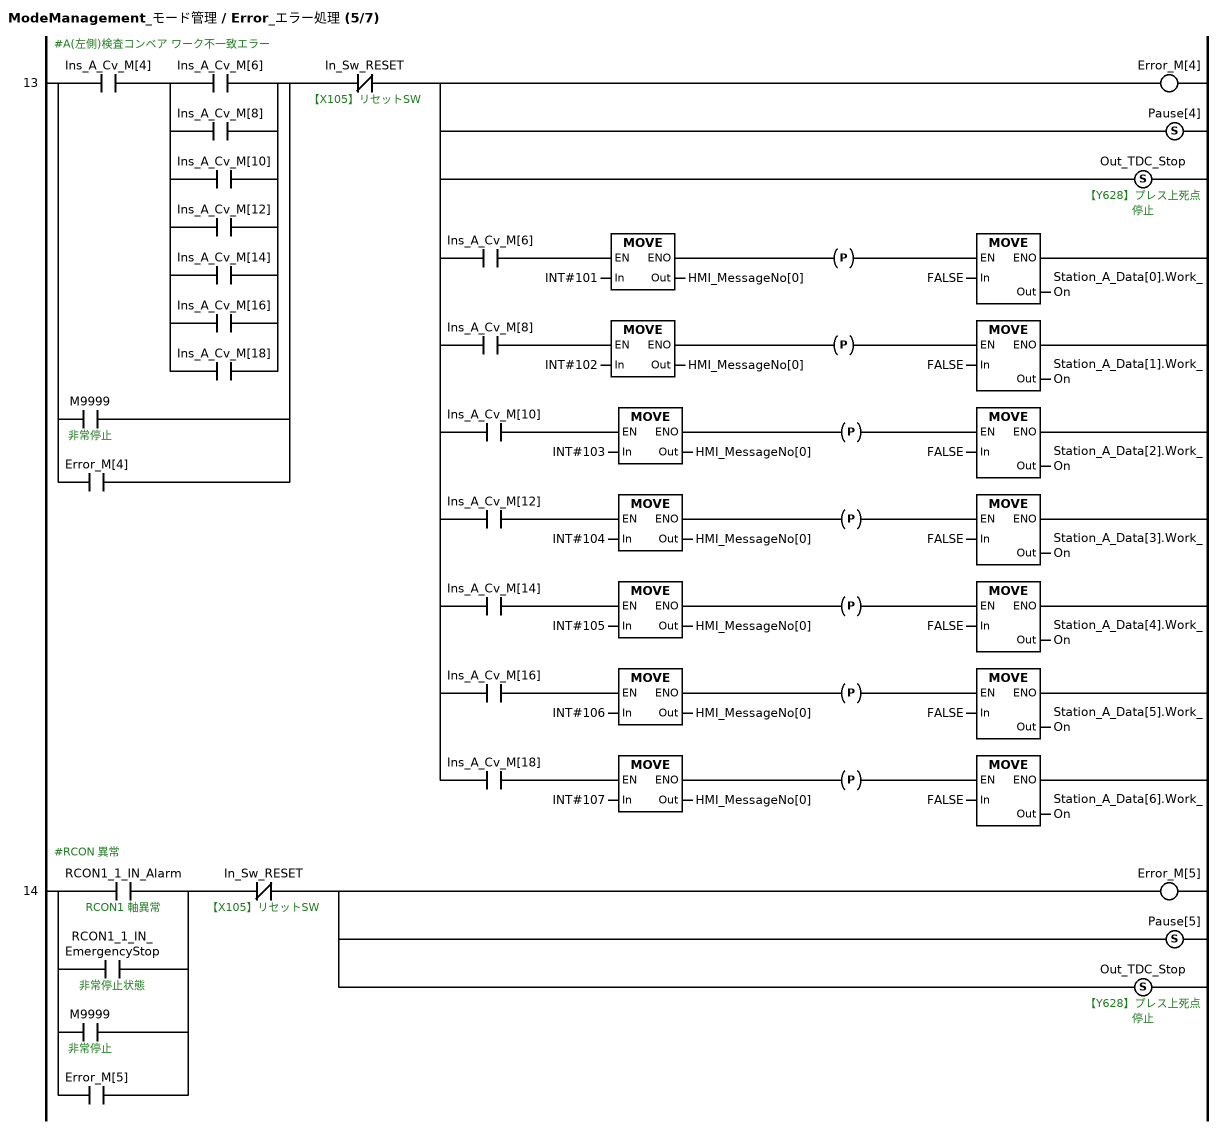
(* [picture p15: ModeManagement_モード管理 / Error_エラー処理, rungs 13-14] *)
(* Rung 13: #A(左側)検査コンベア ワーク不一致エラー *)
_p39 := ((Ins_A_Cv_M[4] AND (Ins_A_Cv_M[6] OR Ins_A_Cv_M[8] OR Ins_A_Cv_M[10] OR Ins_A_Cv_M[12] OR Ins_A_Cv_M[14] OR Ins_A_Cv_M[16] OR Ins_A_Cv_M[18])) OR M9999 OR Error_M[4]) AND NOT In_Sw_RESET;
Error_M[4] := _p39;
IF _p39 THEN
    Pause[4] := TRUE;
    Out_TDC_Stop := TRUE;
END_IF;
IF _p39 AND Ins_A_Cv_M[6] THEN HMI_MessageNo[0] := INT#101; END_IF;
_e40(CLK := _p39 AND Ins_A_Cv_M[6]);
IF _e40.Q THEN Station_A_Data[0].Work_On := FALSE; END_IF;
IF _p39 AND Ins_A_Cv_M[8] THEN HMI_MessageNo[0] := INT#102; END_IF;
_e41(CLK := _p39 AND Ins_A_Cv_M[8]);
IF _e41.Q THEN Station_A_Data[1].Work_On := FALSE; END_IF;
IF _p39 AND Ins_A_Cv_M[10] THEN HMI_MessageNo[0] := INT#103; END_IF;
_e42(CLK := _p39 AND Ins_A_Cv_M[10]);
IF _e42.Q THEN Station_A_Data[2].Work_On := FALSE; END_IF;
IF _p39 AND Ins_A_Cv_M[12] THEN HMI_MessageNo[0] := INT#104; END_IF;
_e43(CLK := _p39 AND Ins_A_Cv_M[12]);
IF _e43.Q THEN Station_A_Data[3].Work_On := FALSE; END_IF;
IF _p39 AND Ins_A_Cv_M[14] THEN HMI_MessageNo[0] := INT#105; END_IF;
_e44(CLK := _p39 AND Ins_A_Cv_M[14]);
IF _e44.Q THEN Station_A_Data[4].Work_On := FALSE; END_IF;
IF _p39 AND Ins_A_Cv_M[16] THEN HMI_MessageNo[0] := INT#106; END_IF;
_e45(CLK := _p39 AND Ins_A_Cv_M[16]);
IF _e45.Q THEN Station_A_Data[5].Work_On := FALSE; END_IF;
IF _p39 AND Ins_A_Cv_M[18] THEN HMI_MessageNo[0] := INT#107; END_IF;
_e46(CLK := _p39 AND Ins_A_Cv_M[18]);
IF _e46.Q THEN Station_A_Data[6].Work_On := FALSE; END_IF;
(* Rung 14: #RCON 異常 *)
_p47 := (RCON1_1_IN_Alarm OR RCON1_1_IN_EmergencyStop OR M9999 OR Error_M[5]) AND NOT In_Sw_RESET;
Error_M[5] := _p47;
IF _p47 THEN
    Pause[5] := TRUE;
    Out_TDC_Stop := TRUE;
END_IF;

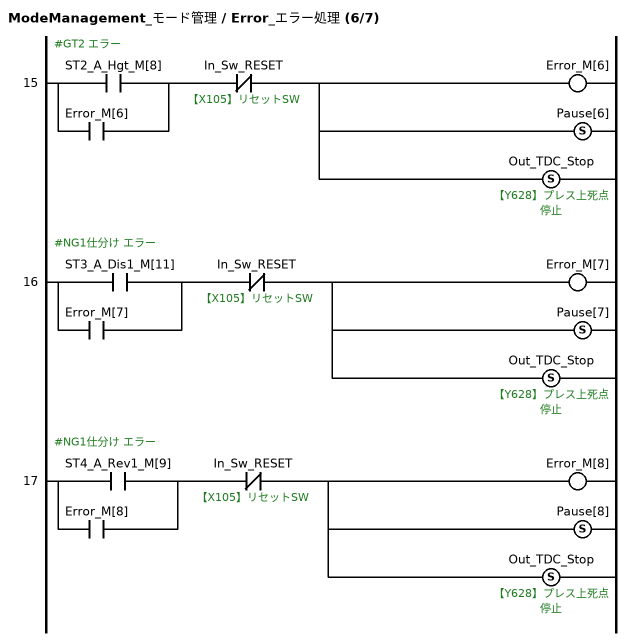
(* Rung 15: #GT2 エラー *)
_p48 := (ST2_A_Hgt_M[8] OR Error_M[6]) AND NOT In_Sw_RESET;
Error_M[6] := _p48;
IF _p48 THEN
    Pause[6] := TRUE;
    Out_TDC_Stop := TRUE;
END_IF;
(* Rung 16: #NG1仕分け エラー *)
_p49 := (ST3_A_Dis1_M[11] OR Error_M[7]) AND NOT In_Sw_RESET;
Error_M[7] := _p49;
IF _p49 THEN
    Pause[7] := TRUE;
    Out_TDC_Stop := TRUE;
END_IF;
(* Rung 17: #NG1仕分け エラー *)
_p50 := (ST4_A_Rev1_M[9] OR Error_M[8]) AND NOT In_Sw_RESET;
Error_M[8] := _p50;
IF _p50 THEN
    Pause[8] := TRUE;
    Out_TDC_Stop := TRUE;
END_IF;

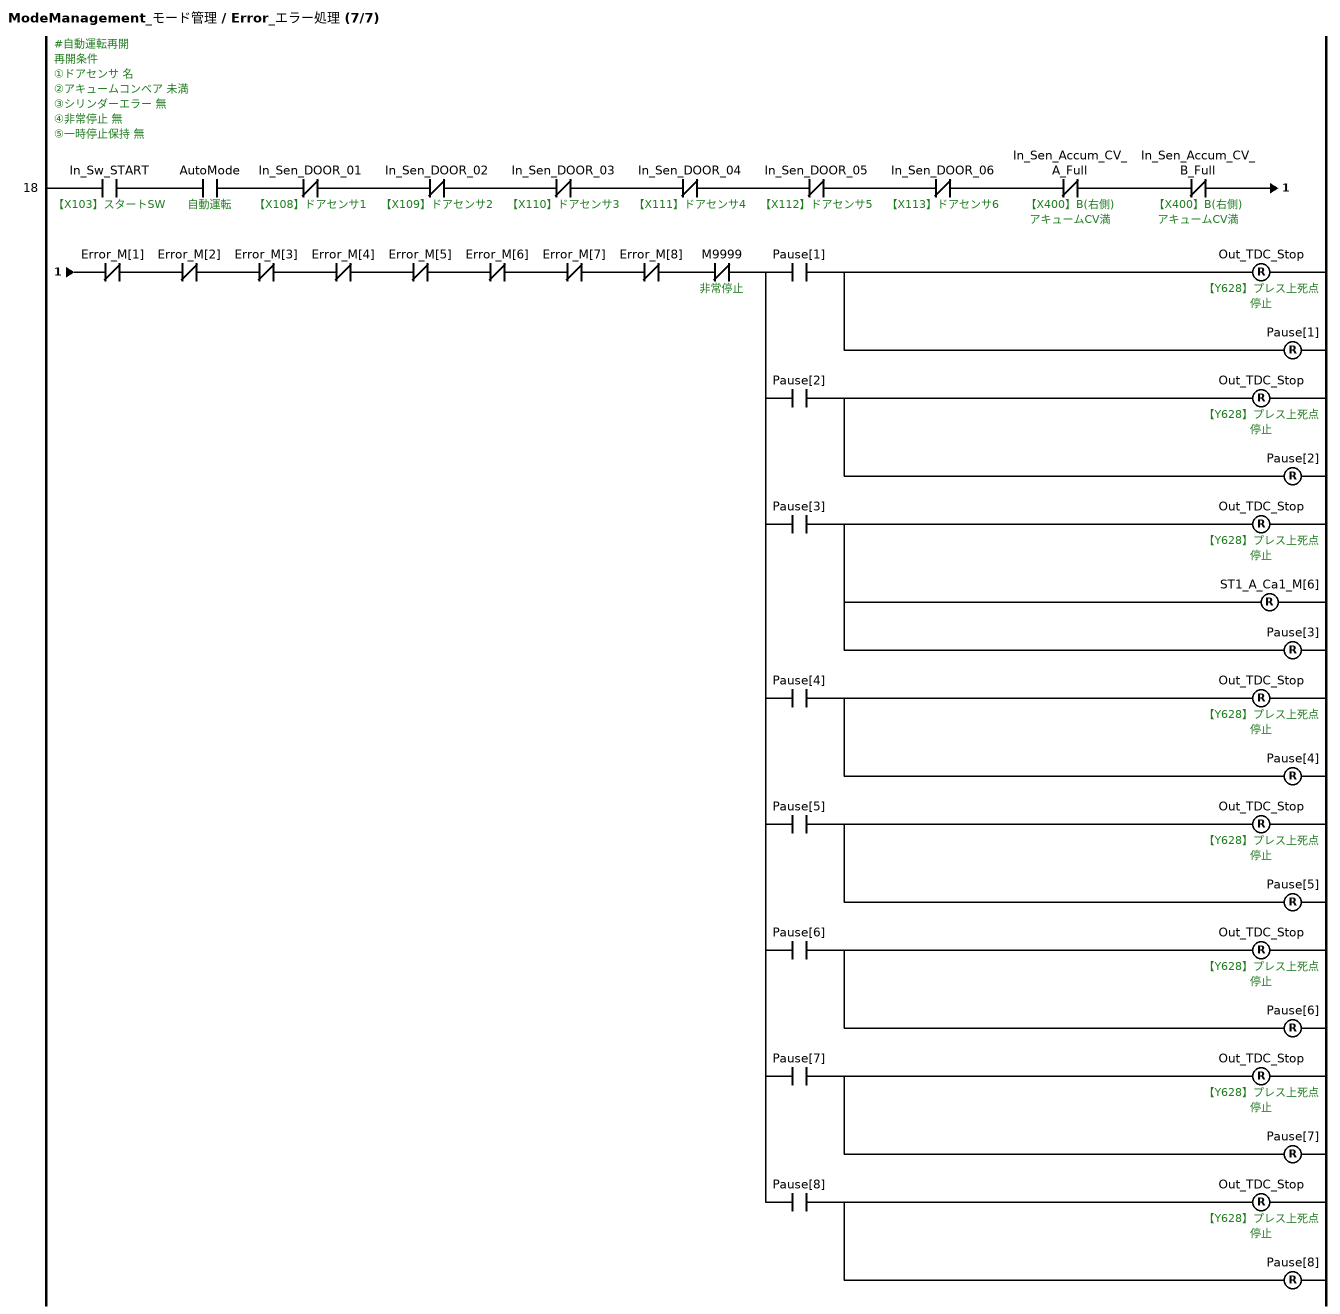
(* Rung 18: #自動運転再開 / 再開条件 / ①ドアセンサ 名 / ②アキュームコンベア 未満 / ③シリンダーエラー 無 / ④非常停止 無 / ⑤一時停止保持 無 *)
_p51 := In_Sw_START AND AutoMode AND NOT In_Sen_DOOR_01 AND NOT In_Sen_DOOR_02 AND NOT In_Sen_DOOR_03 AND NOT In_Sen_DOOR_04 AND NOT In_Sen_DOOR_05 AND NOT In_Sen_DOOR_06 AND NOT In_Sen_Accum_CV_A_Full AND NOT In_Sen_Accum_CV_B_Full AND NOT Error_M[1] AND NOT Error_M[2] AND NOT Error_M[3] AND NOT Error_M[4] AND NOT Error_M[5] AND NOT Error_M[6] AND NOT Error_M[7] AND NOT Error_M[8] AND NOT M9999;
IF _p51 AND Pause[1] THEN
    Out_TDC_Stop := FALSE;
    Pause[1] := FALSE;
END_IF;
IF _p51 AND Pause[2] THEN
    Out_TDC_Stop := FALSE;
    Pause[2] := FALSE;
END_IF;
IF _p51 AND Pause[3] THEN
    Out_TDC_Stop := FALSE;
    ST1_A_Ca1_M[6] := FALSE;
    Pause[3] := FALSE;
END_IF;
IF _p51 AND Pause[4] THEN
    Out_TDC_Stop := FALSE;
    Pause[4] := FALSE;
END_IF;
IF _p51 AND Pause[5] THEN
    Out_TDC_Stop := FALSE;
    Pause[5] := FALSE;
END_IF;
IF _p51 AND Pause[6] THEN
    Out_TDC_Stop := FALSE;
    Pause[6] := FALSE;
END_IF;
IF _p51 AND Pause[7] THEN
    Out_TDC_Stop := FALSE;
    Pause[7] := FALSE;
END_IF;
IF _p51 AND Pause[8] THEN
    Out_TDC_Stop := FALSE;
    Pause[8] := FALSE;
END_IF;
END_PROGRAM

PROGRAM Movements_動作
VAR
    Mo_M : BOOL;
    ST0_A_Sup_M : ARRAY[0..99] OF Bool;  (* [4] 原点位置移動完了 *)
    ST1_Ins_Cv_Rdy : BOOL;
    ST2_Ins_Cv_Rdy : BOOL;
    ST3_Ins_Cv_Rdy : BOOL;
    ST4_Ins_Cv_Rdy : BOOL;
    ST5_Ins_Cv_Rdy : BOOL;
    ST6_Ins_Cv_Rdy : BOOL;
    ST7_Ins_Cv_Rdy : BOOL;
    Ins_A_Cv_T : ARRAY[0..99] OF TON;
    ST1_A_Ca1_Rdy : BOOL;
    GT2_A_Inspection_GetTime : DATE_AND_TIME;
    GT2_A_Inspection_GetTime_ST : STRING[256];
    GT2_A_Inspection_GetTime_ST_Del : STRING[20];
    ST4_A_Rev1_Busy : BOOL;  (* ST4 A 動作中 *)
END_VAR
VAR_EXTERNAL
    ST0_Sup_Start : BOOL;  (* ST0_動作開始 *)
    M9999 : BOOL;
    Out_CYw_Sply_Pick_A_H_Auto : ARRAY[0..10] OF Bool;
    Out_CYw_Sply_Pick_A_H_Done : BOOL;
    Out_CYw_Sply_Slide_A_H_Auto : ARRAY[0..10] OF Bool;
    Out_CYw_Sply_Slide_A_H_Done : BOOL;
    Out_CYw_Sup_Chuck_A_Cl_H_Auto : ARRAY[0..10] OF Bool;
    Out_CYw_Sup_Chuck_A_Cl_H_Done : BOOL;
    In_Sen_Accum_CV_A_Arrival : BOOL;
    In_Sen_Work_A_Pos_00 : BOOL;
    Out_CYw_Sply_Pick_A_F_Auto : ARRAY[0..10] OF Bool;
    Out_CYw_Sply_Pick_A_F_Done : BOOL;
    Out_CYw_Sup_Chuck_A_Cl_F_Auto : ARRAY[0..10] OF Bool;
    Out_CYw_Sup_Chuck_A_Cl_F_Done : BOOL;
    Out_CYw_Sply_Slide_A_F_Auto : ARRAY[0..10] OF Bool;
    Out_CYw_Sply_Slide_A_F_Done : BOOL;
    Station_A_Data : ARRAY[0..8] OF sData;
    Cv_A_Data : ARRAY[0..8] OF sData;
    ST0_A_Sup_End : BOOL;  (* ST0 検査コンベア運転可 *)
    Out_CYS_Pos_01_Stopper_B_H_Auto : ARRAY[0..10] OF Bool;
    Out_CYS_Pos_02_Stopper_B_H_Auto : ARRAY[0..10] OF Bool;
    Out_CYS_Pos_03_Stopper_B_H_Auto : ARRAY[0..10] OF Bool;
    Out_CYS_Pos_04_Stopper_B_H_Auto : ARRAY[0..10] OF Bool;
    Out_CYS_Pos_05_Stopper_B_H_Auto : ARRAY[0..10] OF Bool;
    Out_CYS_Pos_06_Stopper_B_H_Auto : ARRAY[0..10] OF Bool;
    TimerQ_In_SenCY_Pos_01_Stopper_A_H : BOOL;
    TimerQ_In_SenCY_Pos_02_Stopper_A_H : BOOL;
    TimerQ_In_SenCY_Pos_03_Stopper_A_H : BOOL;
    TimerQ_In_SenCY_Pos_04_Stopper_A_H : BOOL;
    TimerQ_In_SenCY_Pos_05_Stopper_A_H : BOOL;
    TimerQ_In_SenCY_Pos_06_Stopper_A_H : BOOL;
    Out_Insp_Cv_A_Run_Auto : ARRAY[0..10] OF Bool;
    TimerQ_In_Sen_Work_A_Pos_01 : BOOL;
    TimerQ_In_Sen_Work_A_Pos_02 : BOOL;
    Pause : ARRAY[0..99] OF Bool;
    TimerQ_In_Sen_Work_A_Pos_03 : BOOL;
    TimerQ_In_Sen_Work_A_Pos_04 : BOOL;
    TimerQ_In_Sen_Work_A_Pos_05 : BOOL;
    TimerQ_In_Sen_Work_A_Pos_06 : BOOL;
    TimerQ_In_Sen_Work_A_Pos_07 : BOOL;
    Out_CYS_Pos_01_Stopper_A_H_Auto : ARRAY[0..10] OF Bool;
    Out_CYS_Pos_02_Stopper_A_H_Auto : ARRAY[0..10] OF Bool;
    Out_CYS_Pos_03_Stopper_A_H_Auto : ARRAY[0..10] OF Bool;
    Out_CYS_Pos_04_Stopper_A_H_Auto : ARRAY[0..10] OF Bool;
    Out_CYS_Pos_05_Stopper_A_H_Auto : ARRAY[0..10] OF Bool;
    Out_CYS_Pos_06_Stopper_A_H_Auto : ARRAY[0..10] OF Bool;
    Ins_A_Cv_M : ARRAY[0..99] OF Bool;
    Ins_A_Cv_Error : BOOL;  (* 検査コンベア ワーク不一致エラー *)
    TimerQ_In_Sen_Work_A_Pos_00 : BOOL;
    Out_CYS_Pos_01_Stopper_A_F_Auto : ARRAY[0..10] OF Bool;
    Out_CYS_Pos_02_Stopper_A_F_Auto : ARRAY[0..10] OF Bool;
    Out_CYS_Pos_03_Stopper_A_F_Auto : ARRAY[0..10] OF Bool;
    Out_CYS_Pos_04_Stopper_A_F_Auto : ARRAY[0..10] OF Bool;
    Out_CYS_Pos_05_Stopper_A_F_Auto : ARRAY[0..10] OF Bool;
    Out_CYS_Pos_06_Stopper_A_F_Auto : ARRAY[0..10] OF Bool;
    Ins_A_Next_Cycle : BOOL;  (* A(左側)検査コンベア 動作完了 *)
    ST0_A_Sup_Busy : BOOL;  (* ST0 稼働中 *)
    Ins_A_End : BOOL;  (* 検査完了 コンベア運転可能 *)
    Auto_A_Start : BOOL;
    Out_CYS_Pos_01_Stopper_A_H_Done : BOOL;
    FH_5552_10_A_Auto : BOOL;
    FH_A_ST1_Done : BOOL;
    ST1_A_Ca1_Busy : BOOL;  (* ST1 A検査中 *)
    ST1_A_Ca1_End : BOOL;  (* ST1 A 動作完了 *)
    ST2_A_Hgt_Busy : BOOL;  (* ST2 A 動作中 *)
    Out_CYw_HgtInsp_Clp_A_H_Auto : ARRAY[0..10] OF Bool;
    Out_CYw_HgtInsp_Clp_A_H_Done : BOOL;
    Out_CYw_HgtInsp_Lf_A_H_Auto : ARRAY[0..10] OF Bool;
    Out_CYw_HgtInsp_Lf_A_H_Done : BOOL;
    Out_CYS_Pos_02_Stopper_A_H_Done : BOOL;
    Out_CYw_HgtInsp_Clp_A_F_Auto : ARRAY[0..10] OF Bool;
    Out_CYw_HgtInsp_Clp_A_F_Done : BOOL;
    Out_CYw_HgtInsp_Lf_A_F_Auto : ARRAY[0..10] OF Bool;
    Out_CYw_HgtInsp_Lf_A_F_Done : BOOL;
    DLEP1_GT2_A_Auto : BOOL;
    Hgt_A_ComputedValueData : LREAL;
    Hight_LowerLimit : LREAL;  (* 高さ検査 下限値 *)
    Hight_UpperLimit : LREAL;  (* 高さ検査 上限値 *)
    ST2_A_Hgt_End : BOOL;  (* 高さ検査完了 *)
    ST3_A_Dis1_Busy : BOOL;  (* ST3 A 動作中 *)
    Out_CYw_NG1_Srt_A_H_Auto : ARRAY[0..10] OF Bool;
    Out_CYw_NG1_Srt_A_H_Done : BOOL;
    Out_CYw_Rev_01_Pick_A_H_Auto : ARRAY[0..10] OF Bool;  (* 自動【Y710】A(左側)ST4 反転1ピックアップ戻： *)
    Out_CYw_Rev_01_Pick_A_H_Done : BOOL;  (* 【Y710】A(左側)ST4 反転1ピックアップ戻 動作完了 *)
    Out_CYw_NG1_Pick_A_H_Auto : ARRAY[0..10] OF Bool;
    Out_CYw_NG1_Pick_A_H_Done : BOOL;
    Out_CYw_NG1_Chk_A_H_Auto : ARRAY[0..10] OF Bool;
    Out_CYw_NG1_Chk_A_H_Done : BOOL;
    RCON1_IAI_Auto : ARRAY[0..99] OF Bool;  (* A(左側) RCON1/Node1/ NG排出： *)
    RCON1_OUT_TargetPos_mm : LREAL;
    HMI_RCON1_OUT_TargetPos : ARRAY[0..99] OF LREAL;  (* HMI RC01 NG仕分け位置： *)
    RCON1_1_M : ARRAY[0..99] OF BOOL;
    Error_M : ARRAY[0..99] OF Bool;
    ST1_A_Ca1_M : ARRAY[0..99] OF Bool;  (* [6] ST2 検査前ワーク不一致エラー; [3] ワーク有無 判定; [1] ST1 A カメラ1 検査開始; [4] ST1 A ワーク有; [5] ST1 A ワーク無; [2] 【Y720】A(左側) 位置1ストッパー 戻; [7] ST1 FH測定開始 *)
    ST2_A_Hgt_M : ARRAY[0..99] OF Bool;  (* [4] 【Y721】A(左側) 位置2ストッパー戻; [6] ST1 A ワーク有; [7] ST1 A ワーク無; [5] ワーク有無 判定; [9] 【Y703】A(左側) 高さ検査持上行; [10] 【Y701】A(左側) 高さ検査押え行; [11] A(左側) 高さ検査OK判定; [12] A(左側) 高さ検査NG判定; [2] 【Y701】A(左側) 高さ検査押え行; [8] ST3 検査前ワーク不一致エラー *)
    Out_CYS_Pos_03_Stopper_A_H_Done : BOOL;
    Out_CYw_NG1_Pick_A_F_Auto : ARRAY[0..10] OF Bool;
    Out_CYw_NG1_Pick_A_F_Done : BOOL;
    Out_CYw_NG1_Chk_A_F_Auto : ARRAY[0..10] OF Bool;
    Out_CYw_NG1_Chk_A_F_Done : BOOL;
    Out_CYw_NG1_Srt_A_F_Auto : ARRAY[0..10] OF Bool;
    Out_CYw_NG1_Srt_A_F_Done : BOOL;
    ST3_A_Dis1_End : BOOL;  (* 左NG1排出 完了 *)
    ST3_A_Dis1_M : ARRAY[0..99] OF Bool;  (* [7] 原点位置 移動開始; [6] 原点位置移動 データ転送; [5] 【Y722】A(左側) 位置3ストッパー戻; [4] 【Y706】A(左側) NG1チャック戻; [8] ワーク有無 / 検査前ワーク不一致 判定; [9] S3 A ワーク有 工程NG; [10] S3 A ワーク無  前工程OK; [14] 【Y704】A(左側) NG1ピックアップ戻 ; [24] 仕分け完了 *)
    ST4_A_Rev1_M : ARRAY[0..99] OF Bool;  (* [2] ワーク有無 / 検査前ワーク不一致 判定; [3] 【Y723】A(左側) 位置4ストッパー戻; [4] ST4 A ワーク有; [5] ST4 A ワーク無 / 前工程NG; [6] ST4 検査前ワーク不一致エラー *)
    Stm_A_Rev_Axis000_MovePos_Degree : LREAL;
    HMI_Stm_A_Rev_Axis000_MovePos_Degree : LREAL;  (* A(左側)ステッピングモータ000 回転角度 *)
    Stm_A_Rev_Axis000_Auto : ARRAY[0..99] OF Bool;  (* [1] 原点位置移動 開始 *)
    Stm_A_Rev_Axis000_MoveAbsoluteDone : BOOL;
END_VAR
VAR
    _e1 : R_TRIG;
    _p2 : BOOL;
    _e3 : R_TRIG;
    _e4 : R_TRIG;
    _p5 : BOOL;
    _e6 : R_TRIG;
    _e7 : R_TRIG;
    _p8 : BOOL;
    _p9 : BOOL;
    _p10 : BOOL;
    _p11 : BOOL;
    _p12 : BOOL;
    _p13 : BOOL;
    _p14 : BOOL;
    _p15 : BOOL;
    _e16 : R_TRIG;
    _p17 : BOOL;
    _p18 : BOOL;
    _p19 : BOOL;
    _p20 : BOOL;
    _p21 : BOOL;
    _p22 : BOOL;
    _p23 : BOOL;
    _p24 : BOOL;
    _p25 : BOOL;
    _p26 : BOOL;
    _p27 : BOOL;
    _p28 : BOOL;
    _e29 : R_TRIG;
    _p30 : BOOL;
    _p31 : BOOL;
    _p32 : BOOL;
    _p33 : BOOL;
    _p34 : BOOL;
    _p35 : BOOL;
    _p36 : BOOL;
    _p37 : BOOL;
    _p38 : BOOL;
    _p39 : BOOL;
    _p40 : BOOL;
    _p41 : BOOL;
    _p42 : BOOL;
    _p43 : BOOL;
    _p44 : BOOL;
    _p45 : BOOL;
    _p46 : BOOL;
    _p47 : BOOL;
    _p48 : BOOL;
    _p49 : BOOL;
    _p50 : BOOL;
    _p51 : BOOL;
    _p52 : BOOL;
    _p53 : BOOL;
    _p54 : BOOL;
    _p55 : BOOL;
    _p56 : BOOL;
    _p57 : BOOL;
    _p58 : BOOL;
    _p59 : BOOL;
    _p60 : BOOL;
    _p61 : BOOL;
END_VAR

(* Section Ins_A_Cv_左検査Cv: ladder, written here as Structured Text *)

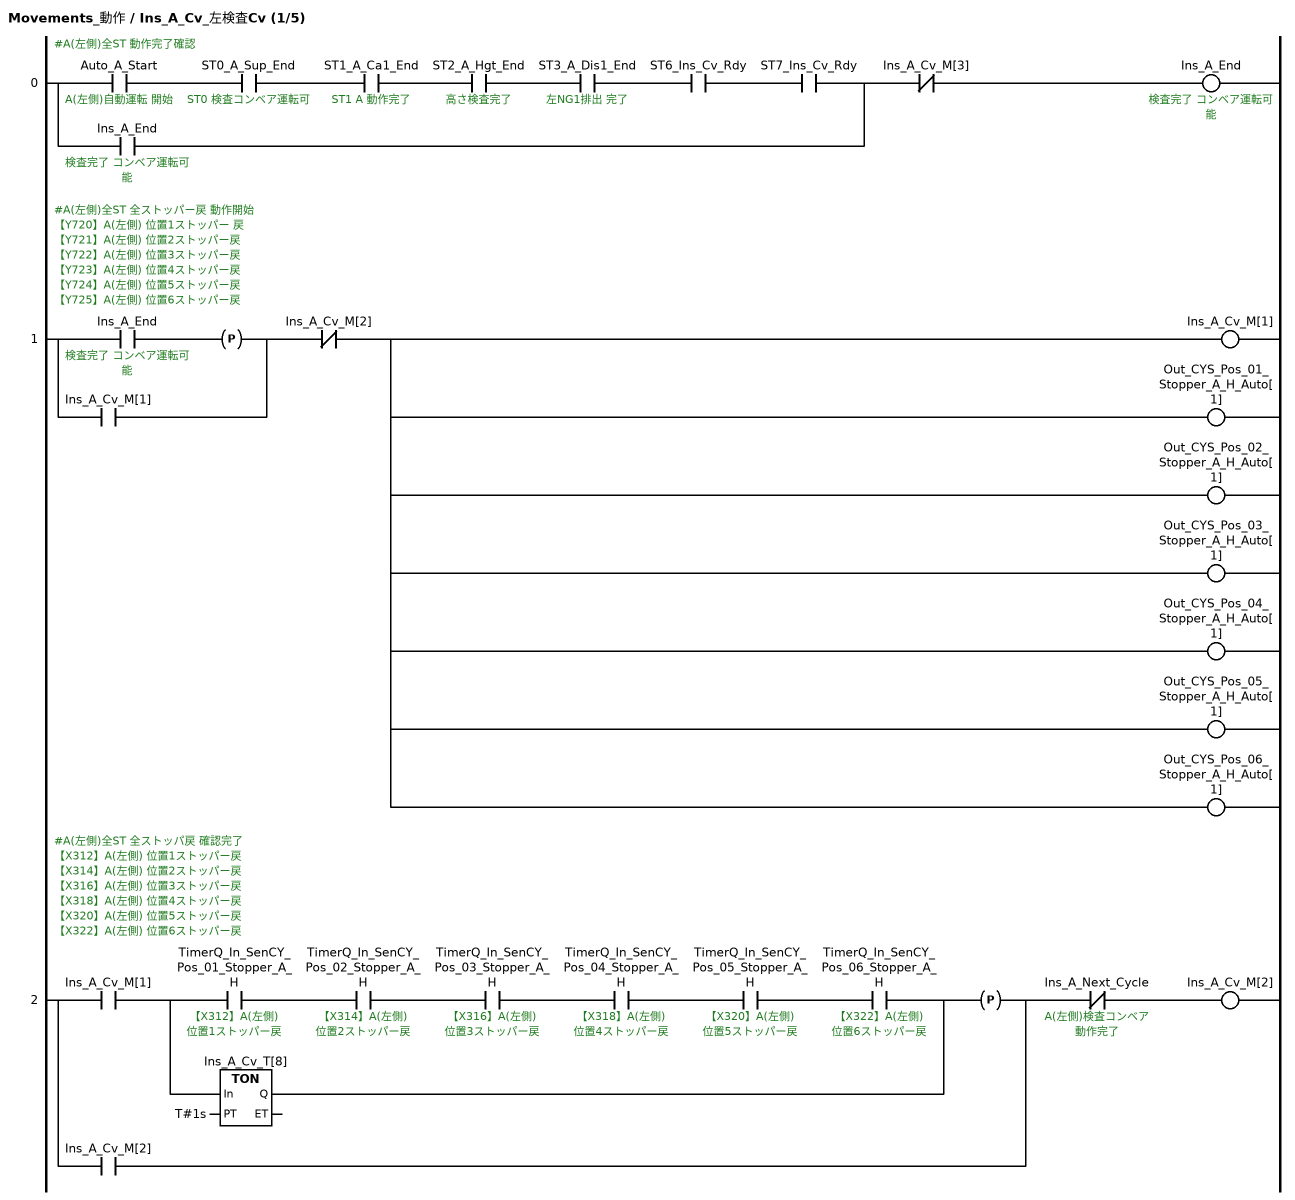
(* Rung 0: #A(左側)全ST 動作完了確認 *)
Ins_A_End := ((Auto_A_Start AND ST0_A_Sup_End AND ST1_A_Ca1_End AND ST2_A_Hgt_End AND ST3_A_Dis1_End AND ST6_Ins_Cv_Rdy AND ST7_Ins_Cv_Rdy) OR Ins_A_End) AND NOT Ins_A_Cv_M[3];
(* Rung 1: #A(左側)全ST 全ストッパー戻 動作開始 / 【Y720】A(左側) 位置1ストッパー 戻 / 【Y721】A(左側) 位置2ストッパー戻 / 【Y722】A(左側) 位置3ストッパー戻 / 【Y723】A(左側) 位置4ストッパー戻 / 【Y724】A(左側) 位置5ストッパー戻 / 【Y725】A(左側) 位置6ストッパー戻 *)
_e1(CLK := Ins_A_End);
_p2 := (_e1.Q OR Ins_A_Cv_M[1]) AND NOT Ins_A_Cv_M[2];
Ins_A_Cv_M[1] := _p2;
Out_CYS_Pos_01_Stopper_A_H_Auto[1] := _p2;
Out_CYS_Pos_02_Stopper_A_H_Auto[1] := _p2;
Out_CYS_Pos_03_Stopper_A_H_Auto[1] := _p2;
Out_CYS_Pos_04_Stopper_A_H_Auto[1] := _p2;
Out_CYS_Pos_05_Stopper_A_H_Auto[1] := _p2;
Out_CYS_Pos_06_Stopper_A_H_Auto[1] := _p2;
(* Rung 2: #A(左側)全ST 全ストッパ戻 確認完了 / 【X312】A(左側) 位置1ストッパー戻 / 【X314】A(左側) 位置2ストッパー戻 / 【X316】A(左側) 位置3ストッパー戻 / 【X318】A(左側) 位置4ストッパー戻 / 【X320】A(左側) 位置5ストッパー戻 / 【X322】A(左側) 位置6ストッパー戻 *)
Ins_A_Cv_T[8](In := Ins_A_Cv_M[1], PT := T#1s);
_e3(CLK := (Ins_A_Cv_M[1] AND TimerQ_In_SenCY_Pos_01_Stopper_A_H AND TimerQ_In_SenCY_Pos_02_Stopper_A_H AND TimerQ_In_SenCY_Pos_03_Stopper_A_H AND TimerQ_In_SenCY_Pos_04_Stopper_A_H AND TimerQ_In_SenCY_Pos_05_Stopper_A_H AND TimerQ_In_SenCY_Pos_06_Stopper_A_H) OR Ins_A_Cv_T[8].Q);
Ins_A_Cv_M[2] := (_e3.Q OR Ins_A_Cv_M[2]) AND NOT Ins_A_Next_Cycle;

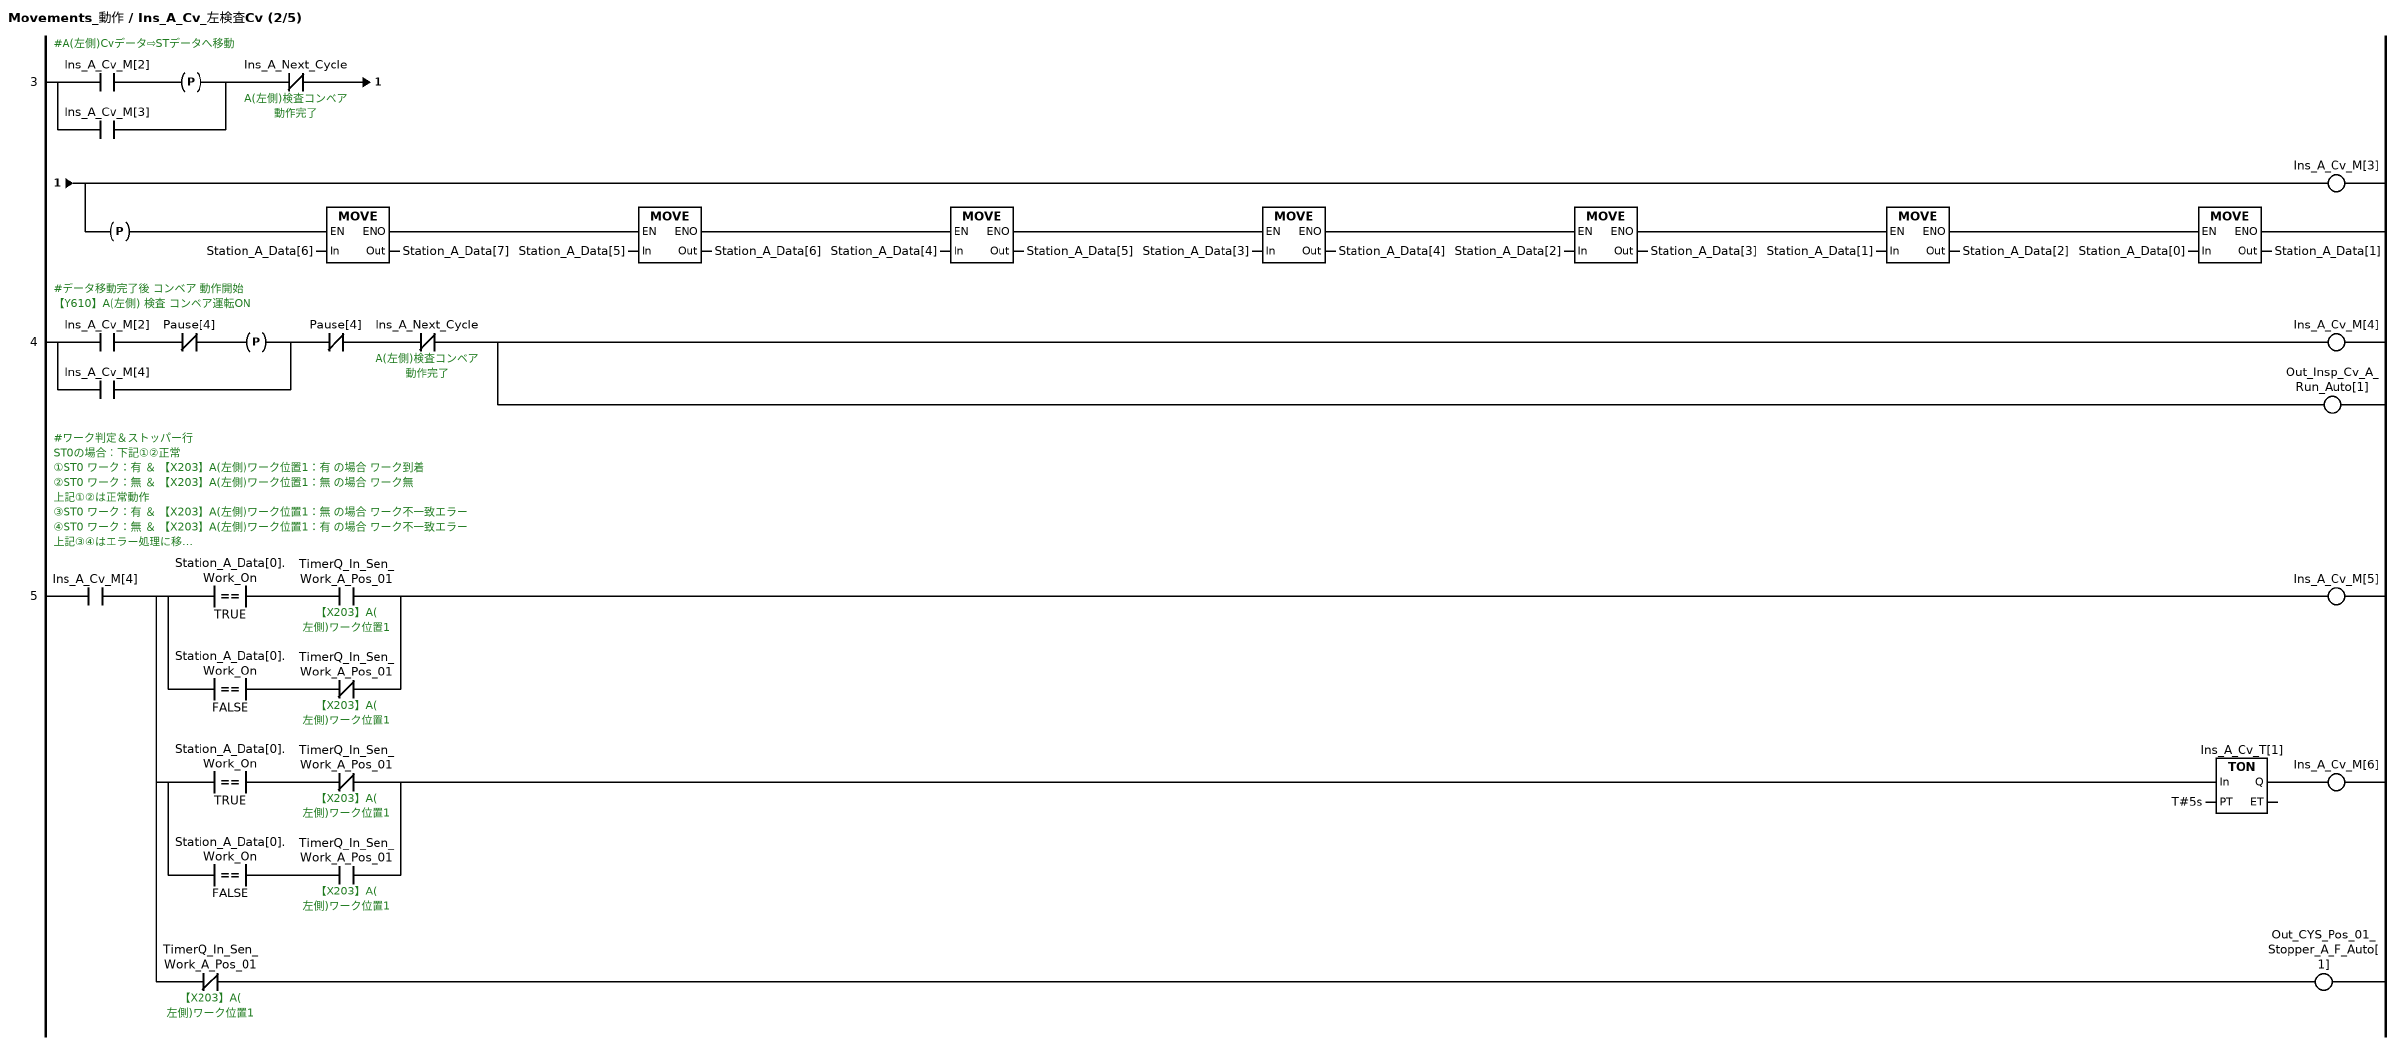
(* Rung 3: #A(左側)Cvデータ⇨STデータへ移動 *)
_e4(CLK := Ins_A_Cv_M[2]);
_p5 := (_e4.Q OR Ins_A_Cv_M[3]) AND NOT Ins_A_Next_Cycle;
Ins_A_Cv_M[3] := _p5;
_e6(CLK := _p5);
IF _e6.Q THEN
    Station_A_Data[7] := Station_A_Data[6];
    Station_A_Data[6] := Station_A_Data[5];
    Station_A_Data[5] := Station_A_Data[4];
    Station_A_Data[4] := Station_A_Data[3];
    Station_A_Data[3] := Station_A_Data[2];
    Station_A_Data[2] := Station_A_Data[1];
    Station_A_Data[1] := Station_A_Data[0];
END_IF;
(* Rung 4: #データ移動完了後 コンベア 動作開始 / 【Y610】A(左側) 検査 コンベア運転ON *)
_e7(CLK := Ins_A_Cv_M[2] AND NOT Pause[4]);
_p8 := (_e7.Q OR Ins_A_Cv_M[4]) AND NOT Pause[4] AND NOT Ins_A_Next_Cycle;
Ins_A_Cv_M[4] := _p8;
Out_Insp_Cv_A_Run_Auto[1] := _p8;
(* Rung 5: #ワーク判定＆ストッパー行 / ST0の場合：下記①②正常 / ①ST0 ワーク：有 ＆ 【X203】A(左側)ワーク位置1：有 の場合 ワーク到着 / ②ST0 ワーク：無 ＆ 【X203】A(左側)ワーク位置1：無 の場合 ワーク無 / 上記①②は正常動作 / ③ST0 ワーク：有 ＆ 【X203】A(左側)ワーク位置1：無 の場合 ワーク不一致エラー / ④ST0 ワーク：無 ＆ 【X203】A(左側)ワーク位置1：有 の場合 ワーク不一致エラー / 上記③④はエラー処理に移動 / ⑤【X203】A(左側)ワーク位置1：無 の場合 / 【Y720】A(左側) 位置1ストッパー 行 *)
_p9 := Ins_A_Cv_M[4];
Ins_A_Cv_M[5] := Ins_A_Cv_M[4] AND (((Station_A_Data[0].Work_On = TRUE) AND TimerQ_In_Sen_Work_A_Pos_01) OR ((Station_A_Data[0].Work_On = FALSE) AND NOT TimerQ_In_Sen_Work_A_Pos_01));
Ins_A_Cv_T[1](In := _p9 AND (((Station_A_Data[0].Work_On = TRUE) AND NOT TimerQ_In_Sen_Work_A_Pos_01) OR ((Station_A_Data[0].Work_On = FALSE) AND TimerQ_In_Sen_Work_A_Pos_01)), PT := T#5s);
Ins_A_Cv_M[6] := Ins_A_Cv_T[1].Q;
Out_CYS_Pos_01_Stopper_A_F_Auto[1] := _p9 AND NOT TimerQ_In_Sen_Work_A_Pos_01;

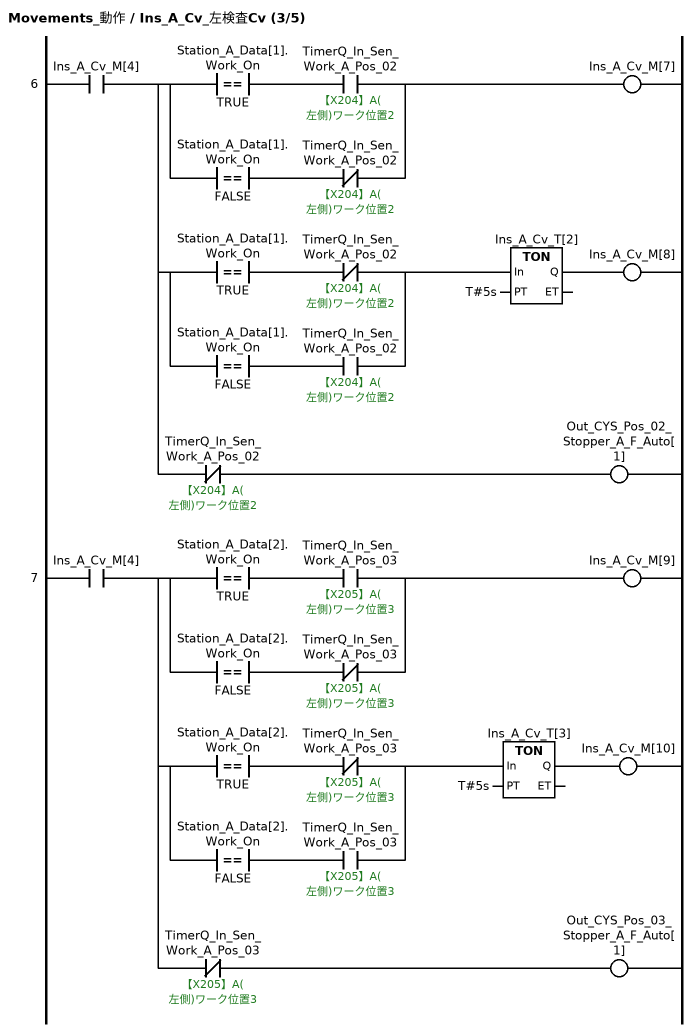
(* Rung 6 *)
_p10 := Ins_A_Cv_M[4];
Ins_A_Cv_M[7] := Ins_A_Cv_M[4] AND (((Station_A_Data[1].Work_On = TRUE) AND TimerQ_In_Sen_Work_A_Pos_02) OR ((Station_A_Data[1].Work_On = FALSE) AND NOT TimerQ_In_Sen_Work_A_Pos_02));
Ins_A_Cv_T[2](In := _p10 AND (((Station_A_Data[1].Work_On = TRUE) AND NOT TimerQ_In_Sen_Work_A_Pos_02) OR ((Station_A_Data[1].Work_On = FALSE) AND TimerQ_In_Sen_Work_A_Pos_02)), PT := T#5s);
Ins_A_Cv_M[8] := Ins_A_Cv_T[2].Q;
Out_CYS_Pos_02_Stopper_A_F_Auto[1] := _p10 AND NOT TimerQ_In_Sen_Work_A_Pos_02;
(* Rung 7 *)
_p11 := Ins_A_Cv_M[4];
Ins_A_Cv_M[9] := Ins_A_Cv_M[4] AND (((Station_A_Data[2].Work_On = TRUE) AND TimerQ_In_Sen_Work_A_Pos_03) OR ((Station_A_Data[2].Work_On = FALSE) AND NOT TimerQ_In_Sen_Work_A_Pos_03));
Ins_A_Cv_T[3](In := _p11 AND (((Station_A_Data[2].Work_On = TRUE) AND NOT TimerQ_In_Sen_Work_A_Pos_03) OR ((Station_A_Data[2].Work_On = FALSE) AND TimerQ_In_Sen_Work_A_Pos_03)), PT := T#5s);
Ins_A_Cv_M[10] := Ins_A_Cv_T[3].Q;
Out_CYS_Pos_03_Stopper_A_F_Auto[1] := _p11 AND NOT TimerQ_In_Sen_Work_A_Pos_03;

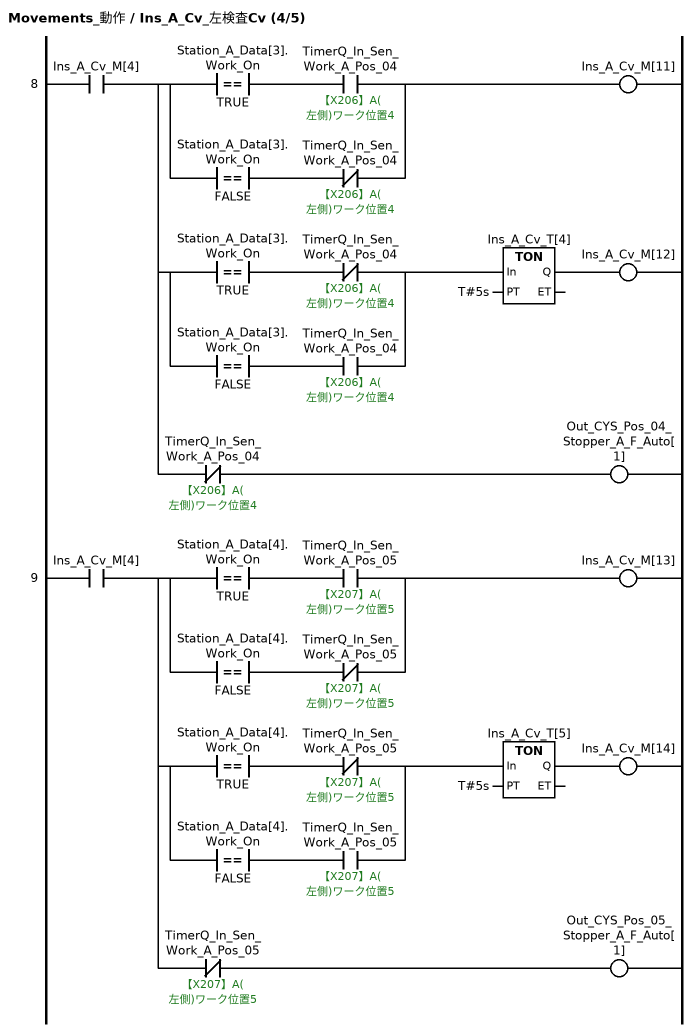
(* Rung 8 *)
_p12 := Ins_A_Cv_M[4];
Ins_A_Cv_M[11] := Ins_A_Cv_M[4] AND (((Station_A_Data[3].Work_On = TRUE) AND TimerQ_In_Sen_Work_A_Pos_04) OR ((Station_A_Data[3].Work_On = FALSE) AND NOT TimerQ_In_Sen_Work_A_Pos_04));
Ins_A_Cv_T[4](In := _p12 AND (((Station_A_Data[3].Work_On = TRUE) AND NOT TimerQ_In_Sen_Work_A_Pos_04) OR ((Station_A_Data[3].Work_On = FALSE) AND TimerQ_In_Sen_Work_A_Pos_04)), PT := T#5s);
Ins_A_Cv_M[12] := Ins_A_Cv_T[4].Q;
Out_CYS_Pos_04_Stopper_A_F_Auto[1] := _p12 AND NOT TimerQ_In_Sen_Work_A_Pos_04;
(* Rung 9 *)
_p13 := Ins_A_Cv_M[4];
Ins_A_Cv_M[13] := Ins_A_Cv_M[4] AND (((Station_A_Data[4].Work_On = TRUE) AND TimerQ_In_Sen_Work_A_Pos_05) OR ((Station_A_Data[4].Work_On = FALSE) AND NOT TimerQ_In_Sen_Work_A_Pos_05));
Ins_A_Cv_T[5](In := _p13 AND (((Station_A_Data[4].Work_On = TRUE) AND NOT TimerQ_In_Sen_Work_A_Pos_05) OR ((Station_A_Data[4].Work_On = FALSE) AND TimerQ_In_Sen_Work_A_Pos_05)), PT := T#5s);
Ins_A_Cv_M[14] := Ins_A_Cv_T[5].Q;
Out_CYS_Pos_05_Stopper_A_F_Auto[1] := _p13 AND NOT TimerQ_In_Sen_Work_A_Pos_05;

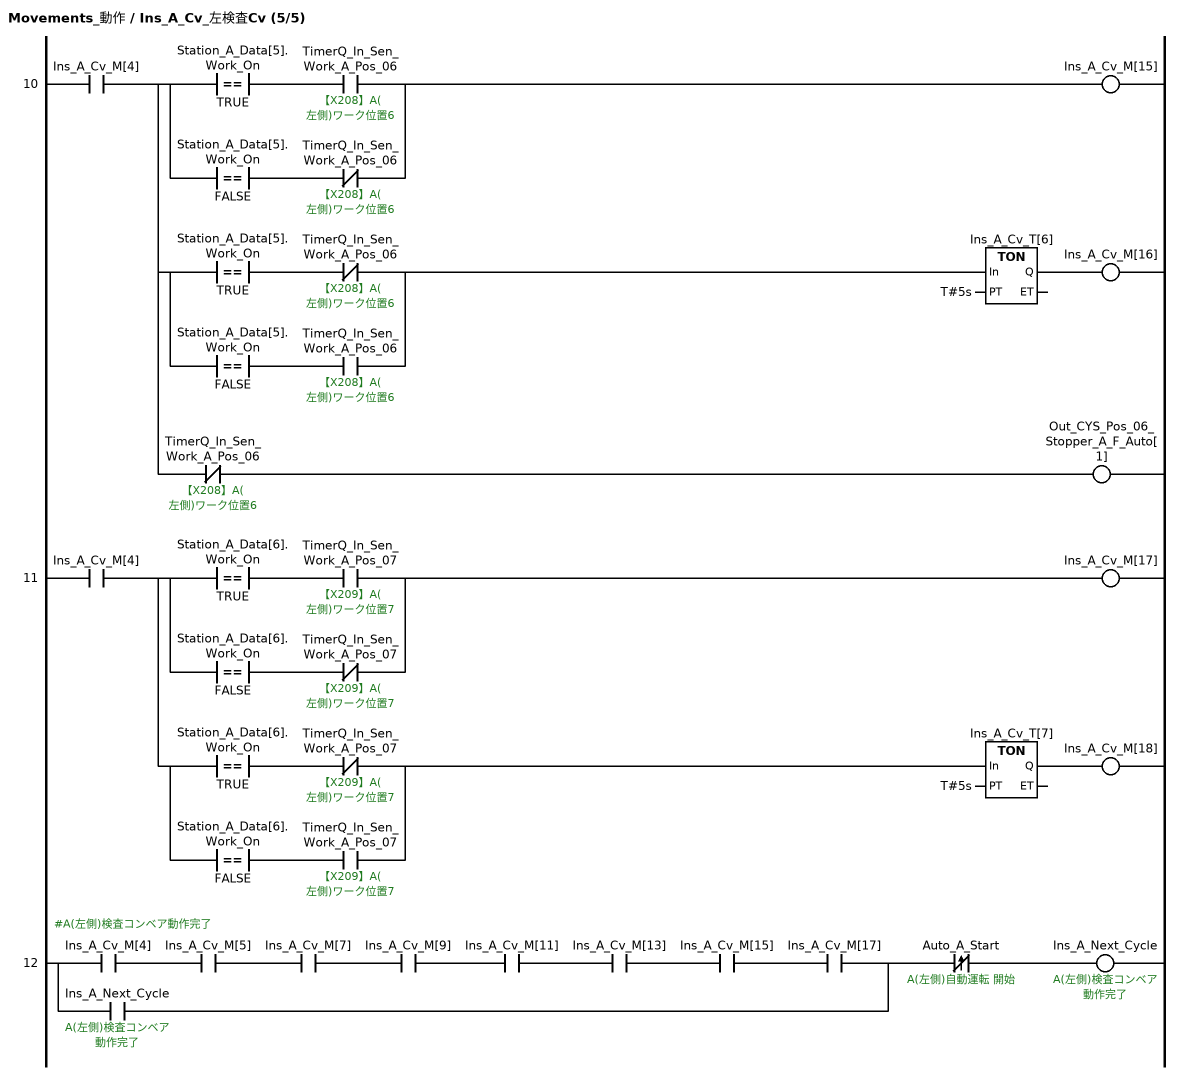
(* Rung 10 *)
_p14 := Ins_A_Cv_M[4];
Ins_A_Cv_M[15] := Ins_A_Cv_M[4] AND (((Station_A_Data[5].Work_On = TRUE) AND TimerQ_In_Sen_Work_A_Pos_06) OR ((Station_A_Data[5].Work_On = FALSE) AND NOT TimerQ_In_Sen_Work_A_Pos_06));
Ins_A_Cv_T[6](In := _p14 AND (((Station_A_Data[5].Work_On = TRUE) AND NOT TimerQ_In_Sen_Work_A_Pos_06) OR ((Station_A_Data[5].Work_On = FALSE) AND TimerQ_In_Sen_Work_A_Pos_06)), PT := T#5s);
Ins_A_Cv_M[16] := Ins_A_Cv_T[6].Q;
Out_CYS_Pos_06_Stopper_A_F_Auto[1] := _p14 AND NOT TimerQ_In_Sen_Work_A_Pos_06;
(* Rung 11 *)
_p15 := Ins_A_Cv_M[4];
Ins_A_Cv_M[17] := Ins_A_Cv_M[4] AND (((Station_A_Data[6].Work_On = TRUE) AND TimerQ_In_Sen_Work_A_Pos_07) OR ((Station_A_Data[6].Work_On = FALSE) AND NOT TimerQ_In_Sen_Work_A_Pos_07));
Ins_A_Cv_T[7](In := _p15 AND (((Station_A_Data[6].Work_On = TRUE) AND NOT TimerQ_In_Sen_Work_A_Pos_07) OR ((Station_A_Data[6].Work_On = FALSE) AND TimerQ_In_Sen_Work_A_Pos_07)), PT := T#5s);
Ins_A_Cv_M[18] := Ins_A_Cv_T[7].Q;
(* Rung 12: #A(左側)検査コンベア動作完了 *)
_e16(CLK := Auto_A_Start);
Ins_A_Next_Cycle := ((Ins_A_Cv_M[4] AND Ins_A_Cv_M[5] AND Ins_A_Cv_M[7] AND Ins_A_Cv_M[9] AND Ins_A_Cv_M[11] AND Ins_A_Cv_M[13] AND Ins_A_Cv_M[15] AND Ins_A_Cv_M[17]) OR Ins_A_Next_Cycle) AND NOT _e16.Q;

(* Section ST0_A_Sup_左供給: ladder, written here as Structured Text *)

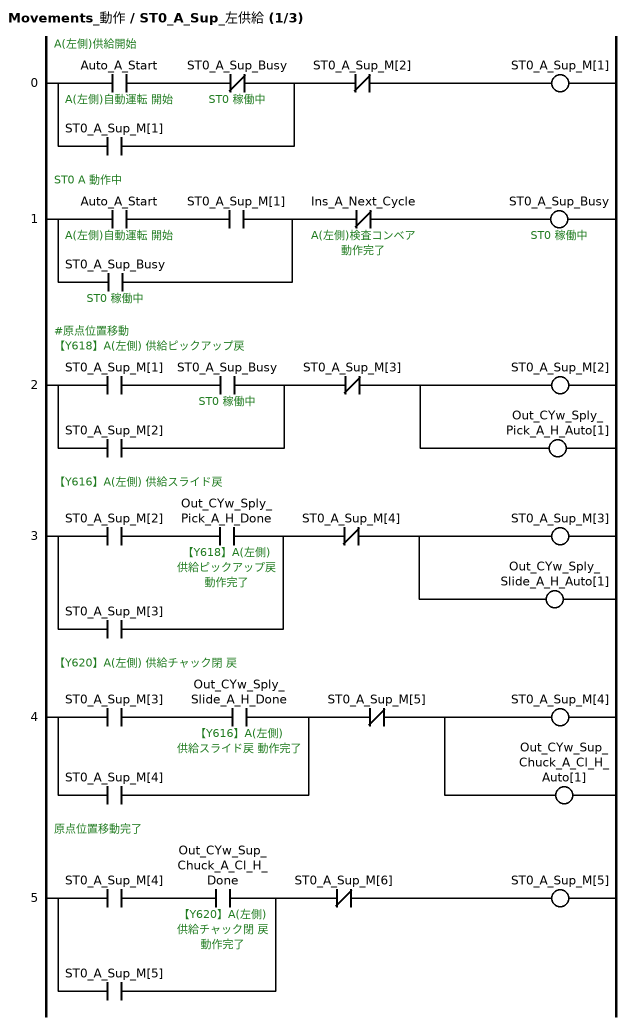
(* Rung 0: A(左側)供給開始 *)
ST0_A_Sup_M[1] := ((Auto_A_Start AND NOT ST0_A_Sup_Busy) OR ST0_A_Sup_M[1]) AND NOT ST0_A_Sup_M[2];
(* Rung 1: ST0 A 動作中 *)
ST0_A_Sup_Busy := ((Auto_A_Start AND ST0_A_Sup_M[1]) OR ST0_A_Sup_Busy) AND NOT Ins_A_Next_Cycle;
(* Rung 2: #原点位置移動 / 【Y618】A(左側) 供給ピックアップ戻 *)
_p17 := ((ST0_A_Sup_M[1] AND ST0_A_Sup_Busy) OR ST0_A_Sup_M[2]) AND NOT ST0_A_Sup_M[3];
ST0_A_Sup_M[2] := _p17;
Out_CYw_Sply_Pick_A_H_Auto[1] := _p17;
(* Rung 3: 【Y616】A(左側) 供給スライド戻 *)
_p18 := ((ST0_A_Sup_M[2] AND Out_CYw_Sply_Pick_A_H_Done) OR ST0_A_Sup_M[3]) AND NOT ST0_A_Sup_M[4];
ST0_A_Sup_M[3] := _p18;
Out_CYw_Sply_Slide_A_H_Auto[1] := _p18;
(* Rung 4: 【Y620】A(左側) 供給チャック閉 戻 *)
_p19 := ((ST0_A_Sup_M[3] AND Out_CYw_Sply_Slide_A_H_Done) OR ST0_A_Sup_M[4]) AND NOT ST0_A_Sup_M[5];
ST0_A_Sup_M[4] := _p19;
Out_CYw_Sup_Chuck_A_Cl_H_Auto[1] := _p19;
(* Rung 5: 原点位置移動完了 *)
ST0_A_Sup_M[5] := ((ST0_A_Sup_M[4] AND Out_CYw_Sup_Chuck_A_Cl_H_Done) OR ST0_A_Sup_M[5]) AND NOT ST0_A_Sup_M[6];

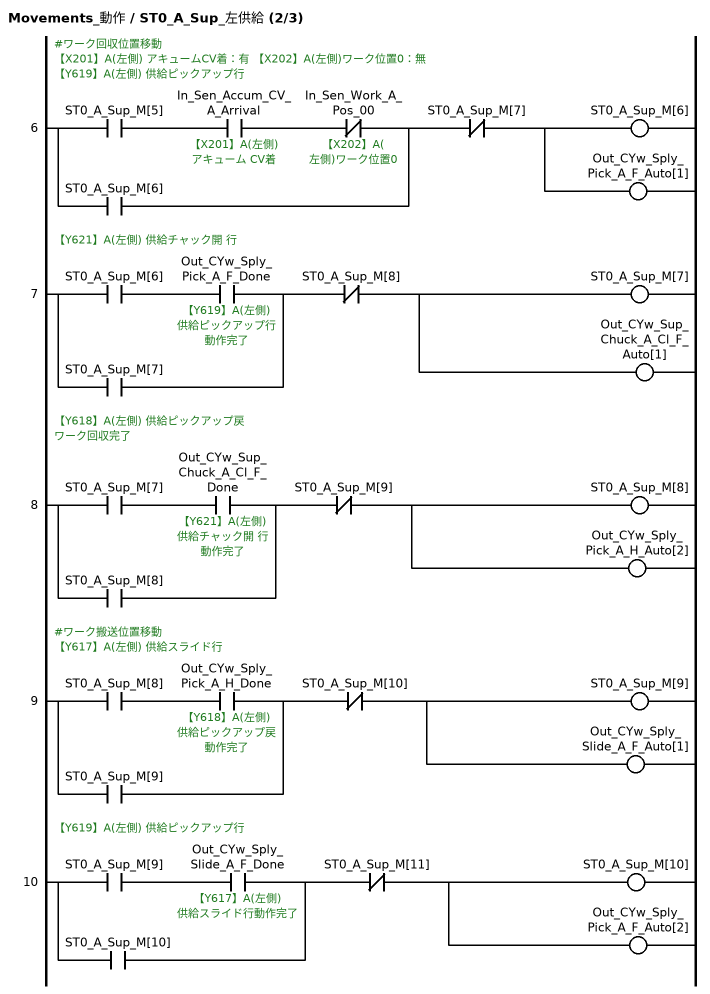
(* Rung 6: #ワーク回収位置移動 / 【X201】A(左側) アキュームCV着：有 【X202】A(左側)ワーク位置0：無 / 【Y619】A(左側) 供給ピックアップ行 *)
_p20 := ((ST0_A_Sup_M[5] AND In_Sen_Accum_CV_A_Arrival AND NOT In_Sen_Work_A_Pos_00) OR ST0_A_Sup_M[6]) AND NOT ST0_A_Sup_M[7];
ST0_A_Sup_M[6] := _p20;
Out_CYw_Sply_Pick_A_F_Auto[1] := _p20;
(* Rung 7: 【Y621】A(左側) 供給チャック開 行 *)
_p21 := ((ST0_A_Sup_M[6] AND Out_CYw_Sply_Pick_A_F_Done) OR ST0_A_Sup_M[7]) AND NOT ST0_A_Sup_M[8];
ST0_A_Sup_M[7] := _p21;
Out_CYw_Sup_Chuck_A_Cl_F_Auto[1] := _p21;
(* Rung 8: 【Y618】A(左側) 供給ピックアップ戻 / ワーク回収完了 *)
_p22 := ((ST0_A_Sup_M[7] AND Out_CYw_Sup_Chuck_A_Cl_F_Done) OR ST0_A_Sup_M[8]) AND NOT ST0_A_Sup_M[9];
ST0_A_Sup_M[8] := _p22;
Out_CYw_Sply_Pick_A_H_Auto[2] := _p22;
(* Rung 9: #ワーク搬送位置移動 / 【Y617】A(左側) 供給スライド行 *)
_p23 := ((ST0_A_Sup_M[8] AND Out_CYw_Sply_Pick_A_H_Done) OR ST0_A_Sup_M[9]) AND NOT ST0_A_Sup_M[10];
ST0_A_Sup_M[9] := _p23;
Out_CYw_Sply_Slide_A_F_Auto[1] := _p23;
(* Rung 10: 【Y619】A(左側) 供給ピックアップ行 *)
_p24 := ((ST0_A_Sup_M[9] AND Out_CYw_Sply_Slide_A_F_Done) OR ST0_A_Sup_M[10]) AND NOT ST0_A_Sup_M[11];
ST0_A_Sup_M[10] := _p24;
Out_CYw_Sply_Pick_A_F_Auto[2] := _p24;

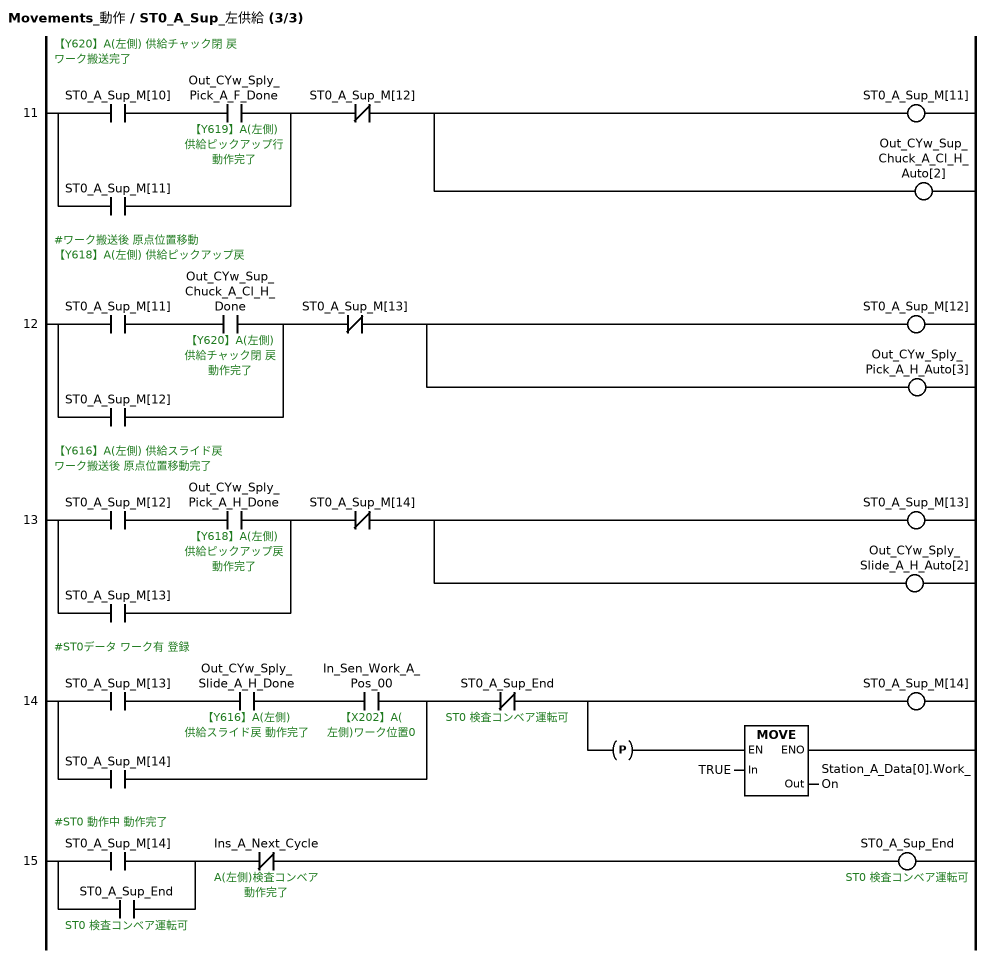
(* Rung 11: 【Y620】A(左側) 供給チャック閉 戻 / ワーク搬送完了 *)
_p25 := ((ST0_A_Sup_M[10] AND Out_CYw_Sply_Pick_A_F_Done) OR ST0_A_Sup_M[11]) AND NOT ST0_A_Sup_M[12];
ST0_A_Sup_M[11] := _p25;
Out_CYw_Sup_Chuck_A_Cl_H_Auto[2] := _p25;
(* Rung 12: #ワーク搬送後 原点位置移動 / 【Y618】A(左側) 供給ピックアップ戻 *)
_p26 := ((ST0_A_Sup_M[11] AND Out_CYw_Sup_Chuck_A_Cl_H_Done) OR ST0_A_Sup_M[12]) AND NOT ST0_A_Sup_M[13];
ST0_A_Sup_M[12] := _p26;
Out_CYw_Sply_Pick_A_H_Auto[3] := _p26;
(* Rung 13: 【Y616】A(左側) 供給スライド戻 / ワーク搬送後 原点位置移動完了 *)
_p27 := ((ST0_A_Sup_M[12] AND Out_CYw_Sply_Pick_A_H_Done) OR ST0_A_Sup_M[13]) AND NOT ST0_A_Sup_M[14];
ST0_A_Sup_M[13] := _p27;
Out_CYw_Sply_Slide_A_H_Auto[2] := _p27;
(* Rung 14: #ST0データ ワーク有 登録 *)
_p28 := ((ST0_A_Sup_M[13] AND Out_CYw_Sply_Slide_A_H_Done AND In_Sen_Work_A_Pos_00) OR ST0_A_Sup_M[14]) AND NOT ST0_A_Sup_End;
ST0_A_Sup_M[14] := _p28;
_e29(CLK := _p28);
IF _e29.Q THEN Station_A_Data[0].Work_On := TRUE; END_IF;
(* Rung 15: #ST0 動作中 動作完了 *)
ST0_A_Sup_End := (ST0_A_Sup_M[14] OR ST0_A_Sup_End) AND NOT Ins_A_Next_Cycle;

(* Section ST1_A_Ca1_左Ca1検査: ladder, written here as Structured Text *)

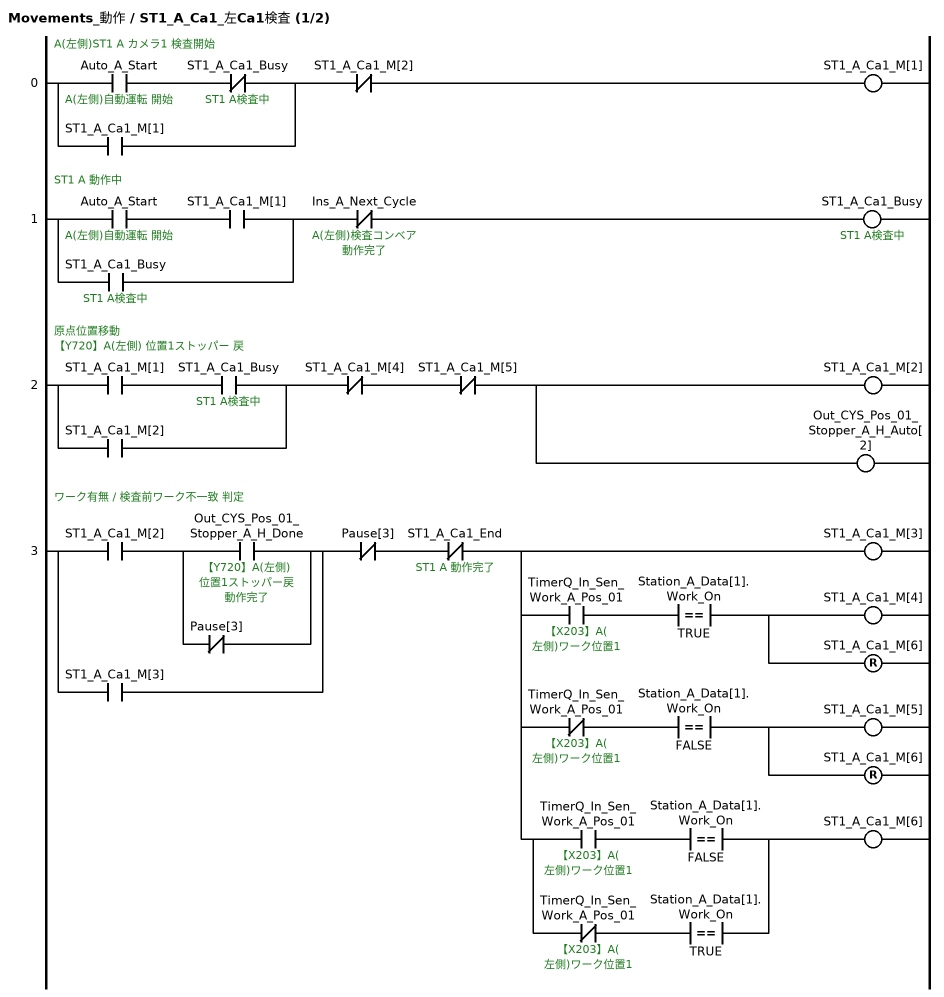
(* Rung 0: A(左側)ST1 A カメラ1 検査開始 *)
ST1_A_Ca1_M[1] := ((Auto_A_Start AND NOT ST1_A_Ca1_Busy) OR ST1_A_Ca1_M[1]) AND NOT ST1_A_Ca1_M[2];
(* Rung 1: ST1 A 動作中 *)
ST1_A_Ca1_Busy := ((Auto_A_Start AND ST1_A_Ca1_M[1]) OR ST1_A_Ca1_Busy) AND NOT Ins_A_Next_Cycle;
(* Rung 2: 原点位置移動 / 【Y720】A(左側) 位置1ストッパー 戻 *)
_p30 := ((ST1_A_Ca1_M[1] AND ST1_A_Ca1_Busy) OR ST1_A_Ca1_M[2]) AND NOT ST1_A_Ca1_M[4] AND NOT ST1_A_Ca1_M[5];
ST1_A_Ca1_M[2] := _p30;
Out_CYS_Pos_01_Stopper_A_H_Auto[2] := _p30;
(* Rung 3: ワーク有無 / 検査前ワーク不一致 判定 *)
_p31 := ((ST1_A_Ca1_M[2] AND (Out_CYS_Pos_01_Stopper_A_H_Done OR NOT Pause[3])) OR ST1_A_Ca1_M[3]) AND NOT Pause[3] AND NOT ST1_A_Ca1_End;
ST1_A_Ca1_M[3] := _p31;
_p32 := _p31 AND TimerQ_In_Sen_Work_A_Pos_01 AND (Station_A_Data[1].Work_On = TRUE);
ST1_A_Ca1_M[4] := _p32;
IF _p32 THEN ST1_A_Ca1_M[6] := FALSE; END_IF;
_p33 := _p31 AND NOT TimerQ_In_Sen_Work_A_Pos_01 AND (Station_A_Data[1].Work_On = FALSE);
ST1_A_Ca1_M[5] := _p33;
IF _p33 THEN ST1_A_Ca1_M[6] := FALSE; END_IF;
ST1_A_Ca1_M[6] := _p31 AND ((TimerQ_In_Sen_Work_A_Pos_01 AND (Station_A_Data[1].Work_On = FALSE)) OR (NOT TimerQ_In_Sen_Work_A_Pos_01 AND (Station_A_Data[1].Work_On = TRUE)));

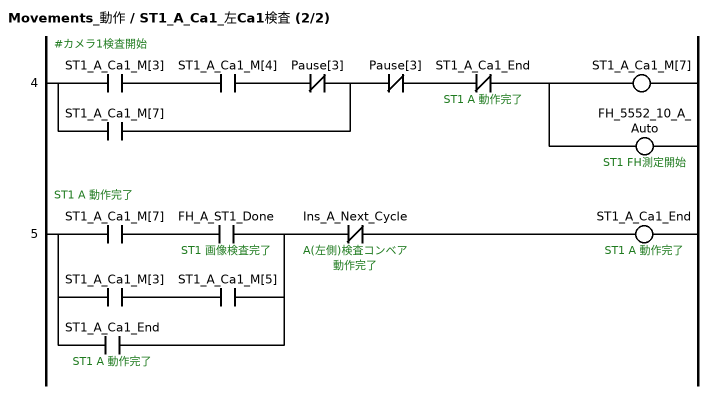
(* Rung 4: #カメラ1検査開始 *)
_p34 := ((ST1_A_Ca1_M[3] AND ST1_A_Ca1_M[4] AND NOT Pause[3]) OR ST1_A_Ca1_M[7]) AND NOT Pause[3] AND NOT ST1_A_Ca1_End;
ST1_A_Ca1_M[7] := _p34;
FH_5552_10_A_Auto := _p34;
(* Rung 5: ST1 A 動作完了 *)
ST1_A_Ca1_End := ((ST1_A_Ca1_M[7] AND FH_A_ST1_Done) OR (ST1_A_Ca1_M[3] AND ST1_A_Ca1_M[5]) OR ST1_A_Ca1_End) AND NOT Ins_A_Next_Cycle;

(* Section ST2_A_Hgt_左高さ検査: ladder, written here as Structured Text *)

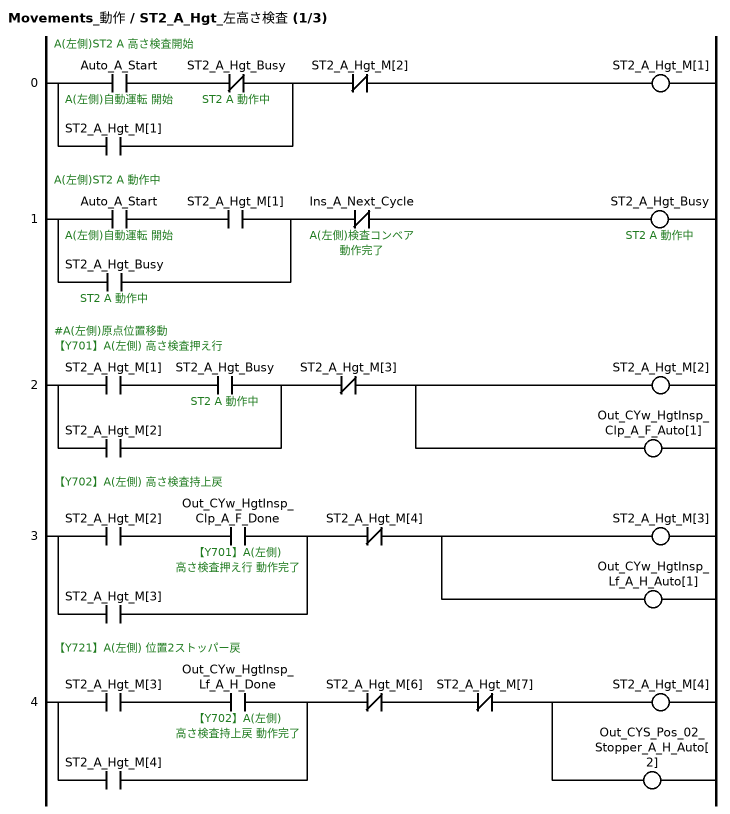
(* Rung 0: A(左側)ST2 A 高さ検査開始 *)
ST2_A_Hgt_M[1] := ((Auto_A_Start AND NOT ST2_A_Hgt_Busy) OR ST2_A_Hgt_M[1]) AND NOT ST2_A_Hgt_M[2];
(* Rung 1: A(左側)ST2 A 動作中 *)
ST2_A_Hgt_Busy := ((Auto_A_Start AND ST2_A_Hgt_M[1]) OR ST2_A_Hgt_Busy) AND NOT Ins_A_Next_Cycle;
(* Rung 2: #A(左側)原点位置移動 / 【Y701】A(左側) 高さ検査押え行 *)
_p35 := ((ST2_A_Hgt_M[1] AND ST2_A_Hgt_Busy) OR ST2_A_Hgt_M[2]) AND NOT ST2_A_Hgt_M[3];
ST2_A_Hgt_M[2] := _p35;
Out_CYw_HgtInsp_Clp_A_F_Auto[1] := _p35;
(* Rung 3: 【Y702】A(左側) 高さ検査持上戻 *)
_p36 := ((ST2_A_Hgt_M[2] AND Out_CYw_HgtInsp_Clp_A_F_Done) OR ST2_A_Hgt_M[3]) AND NOT ST2_A_Hgt_M[4];
ST2_A_Hgt_M[3] := _p36;
Out_CYw_HgtInsp_Lf_A_H_Auto[1] := _p36;
(* Rung 4: 【Y721】A(左側) 位置2ストッパー戻 *)
_p37 := ((ST2_A_Hgt_M[3] AND Out_CYw_HgtInsp_Lf_A_H_Done) OR ST2_A_Hgt_M[4]) AND NOT ST2_A_Hgt_M[6] AND NOT ST2_A_Hgt_M[7];
ST2_A_Hgt_M[4] := _p37;
Out_CYS_Pos_02_Stopper_A_H_Auto[2] := _p37;

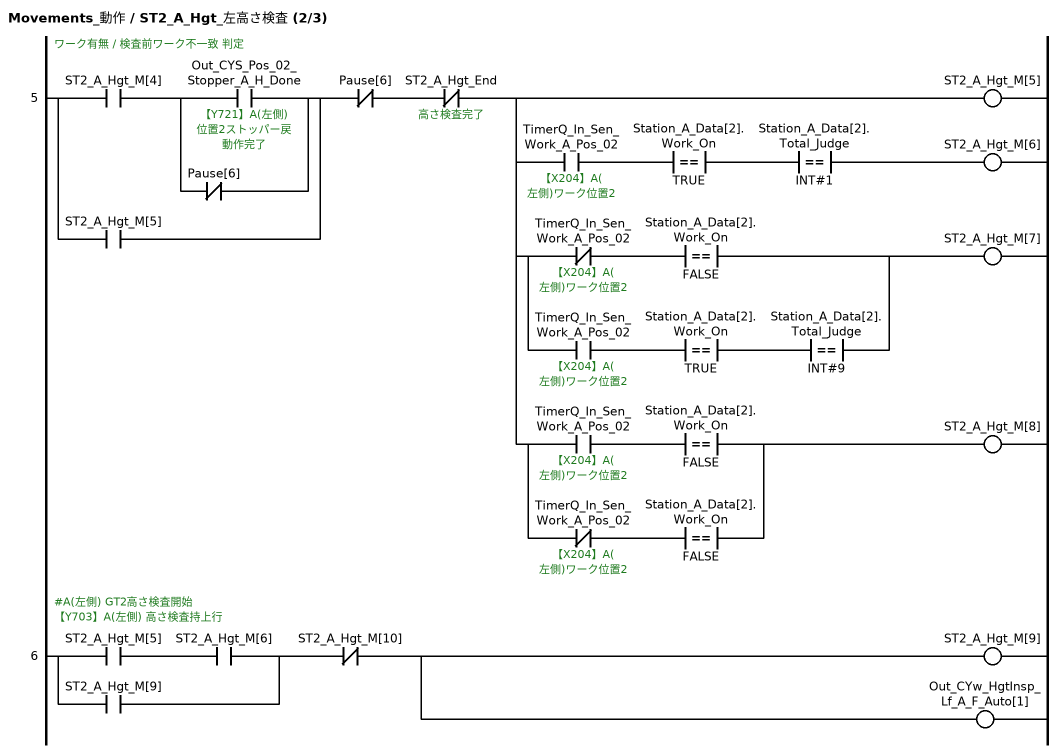
(* Rung 5: ワーク有無 / 検査前ワーク不一致 判定 *)
_p38 := ((ST2_A_Hgt_M[4] AND (Out_CYS_Pos_02_Stopper_A_H_Done OR NOT Pause[6])) OR ST2_A_Hgt_M[5]) AND NOT Pause[6] AND NOT ST2_A_Hgt_End;
ST2_A_Hgt_M[5] := _p38;
ST2_A_Hgt_M[6] := _p38 AND TimerQ_In_Sen_Work_A_Pos_02 AND (Station_A_Data[2].Work_On = TRUE) AND (Station_A_Data[2].Total_Judge = INT#1);
ST2_A_Hgt_M[7] := _p38 AND ((NOT TimerQ_In_Sen_Work_A_Pos_02 AND (Station_A_Data[2].Work_On = FALSE)) OR (TimerQ_In_Sen_Work_A_Pos_02 AND (Station_A_Data[2].Work_On = TRUE) AND (Station_A_Data[2].Total_Judge = INT#9)));
ST2_A_Hgt_M[8] := _p38 AND ((TimerQ_In_Sen_Work_A_Pos_02 AND (Station_A_Data[2].Work_On = FALSE)) OR (NOT TimerQ_In_Sen_Work_A_Pos_02 AND (Station_A_Data[2].Work_On = FALSE)));
(* Rung 6: #A(左側) GT2高さ検査開始 / 【Y703】A(左側) 高さ検査持上行 *)
_p39 := ((ST2_A_Hgt_M[5] AND ST2_A_Hgt_M[6]) OR ST2_A_Hgt_M[9]) AND NOT ST2_A_Hgt_M[10];
ST2_A_Hgt_M[9] := _p39;
Out_CYw_HgtInsp_Lf_A_F_Auto[1] := _p39;

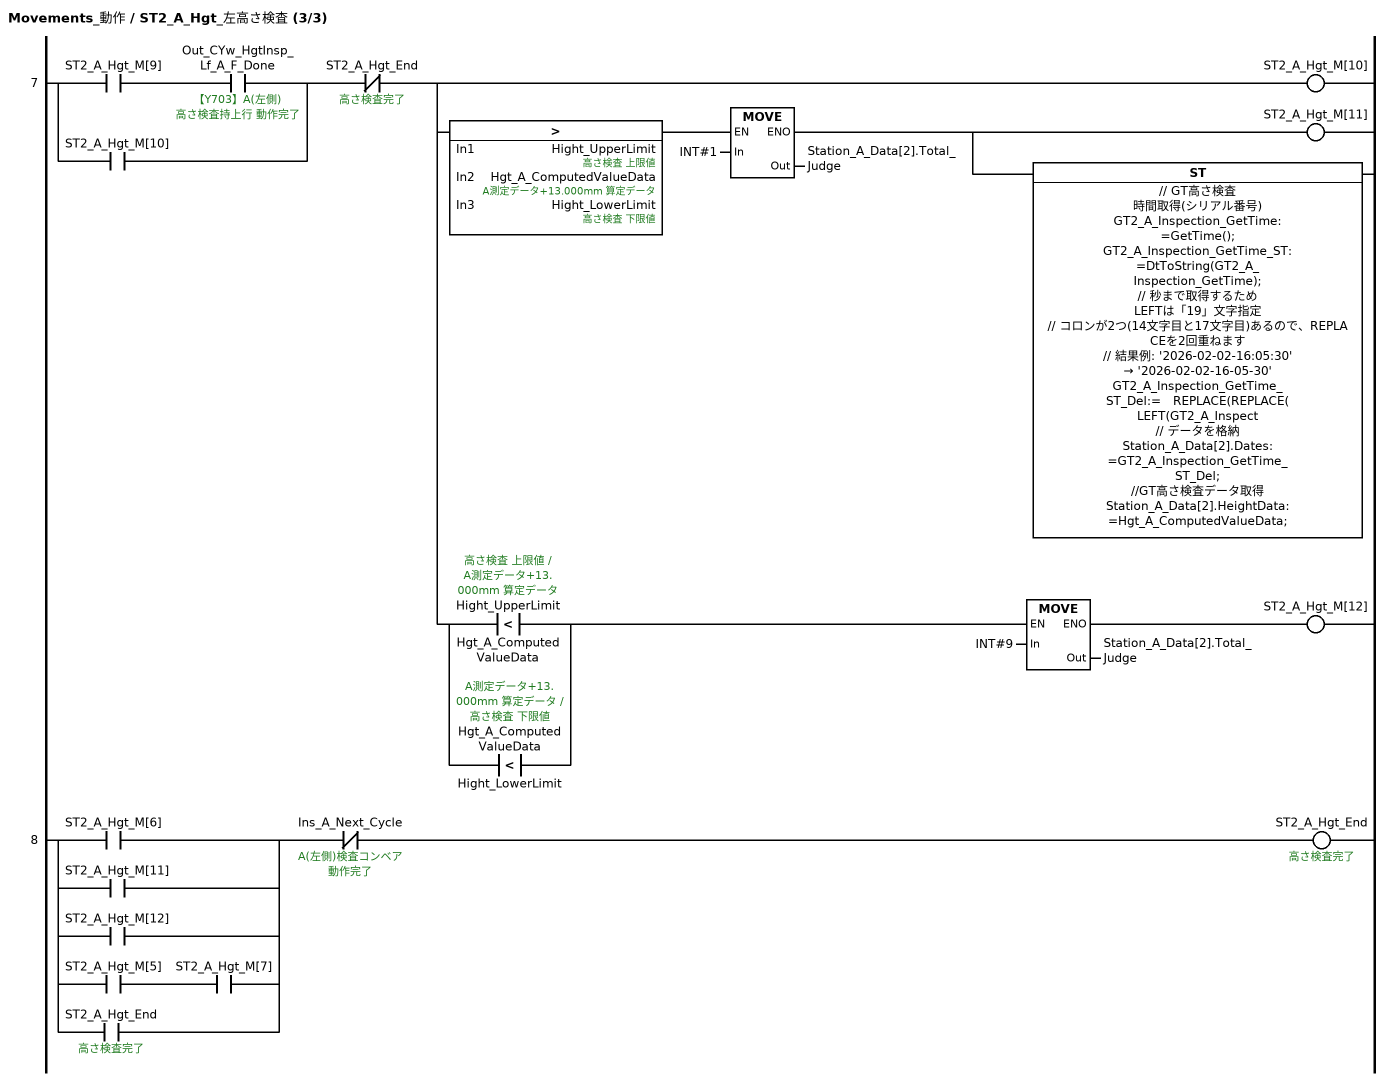
(* Rung 7 *)
_p40 := ((ST2_A_Hgt_M[9] AND Out_CYw_HgtInsp_Lf_A_F_Done) OR ST2_A_Hgt_M[10]) AND NOT ST2_A_Hgt_End;
ST2_A_Hgt_M[10] := _p40;
IF _p40 AND GT(Hight_UpperLimit, Hgt_A_ComputedValueData, Hight_LowerLimit) THEN
    Station_A_Data[2].Total_Judge := INT#1;
END_IF;
_p41 := _p40 AND GT(Hight_UpperLimit, Hgt_A_ComputedValueData, Hight_LowerLimit);
ST2_A_Hgt_M[11] := _p41;
IF _p41 THEN
    // GT高さ検査 時間取得(シリアル番号)
    GT2_A_Inspection_GetTime:=GetTime();
    GT2_A_Inspection_GetTime_ST:=DtToString(GT2_A_Inspection_GetTime);
    // 秒まで取得するため LEFTは「19」文字指定
    // コロンが2つ(14文字目と17文字目)あるので、REPLACEを2回重ねます
    // 結果例: '2026-02-02-16:05:30' → '2026-02-02-16-05-30'
    GT2_A_Inspection_GetTime_ST_Del:=   REPLACE(REPLACE(LEFT(GT2_A_Inspection_GetTime_ST, UINT#19), STRING#'-', UINT#1, UINT#17), STRING#'-', UINT#1, UINT#14);
    // データを格納
    Station_A_Data[2].Dates:=GT2_A_Inspection_GetTime_ST_Del;
    //GT高さ検査データ取得
    Station_A_Data[2].HeightData:=Hgt_A_ComputedValueData;
END_IF;
IF _p40 AND ((Hight_UpperLimit < Hgt_A_ComputedValueData) OR (Hgt_A_ComputedValueData < Hight_LowerLimit)) THEN
    Station_A_Data[2].Total_Judge := INT#9;
END_IF;
ST2_A_Hgt_M[12] := _p40 AND ((Hight_UpperLimit < Hgt_A_ComputedValueData) OR (Hgt_A_ComputedValueData < Hight_LowerLimit));
(* Rung 8 *)
ST2_A_Hgt_End := (ST2_A_Hgt_M[6] OR ST2_A_Hgt_M[11] OR ST2_A_Hgt_M[12] OR (ST2_A_Hgt_M[5] AND ST2_A_Hgt_M[7]) OR ST2_A_Hgt_End) AND NOT Ins_A_Next_Cycle;

(* Section ST3_A_Dis1_左NG1排出: ladder, written here as Structured Text *)

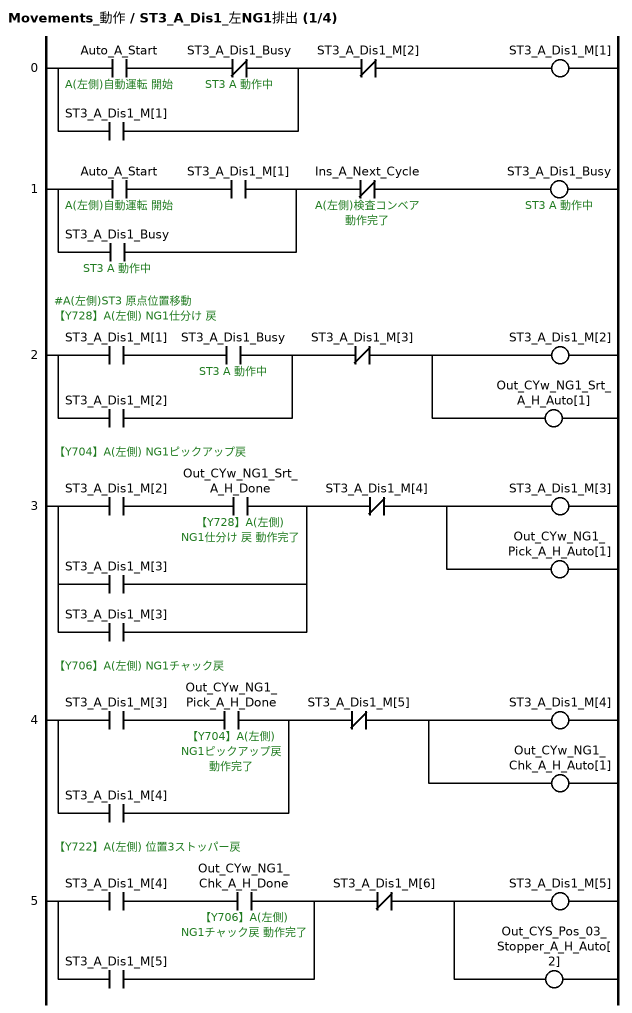
(* Rung 0 *)
ST3_A_Dis1_M[1] := ((Auto_A_Start AND NOT ST3_A_Dis1_Busy) OR ST3_A_Dis1_M[1]) AND NOT ST3_A_Dis1_M[2];
(* Rung 1 *)
ST3_A_Dis1_Busy := ((Auto_A_Start AND ST3_A_Dis1_M[1]) OR ST3_A_Dis1_Busy) AND NOT Ins_A_Next_Cycle;
(* Rung 2: #A(左側)ST3 原点位置移動 / 【Y728】A(左側) NG1仕分け 戻 *)
_p42 := ((ST3_A_Dis1_M[1] AND ST3_A_Dis1_Busy) OR ST3_A_Dis1_M[2]) AND NOT ST3_A_Dis1_M[3];
ST3_A_Dis1_M[2] := _p42;
Out_CYw_NG1_Srt_A_H_Auto[1] := _p42;
(* Rung 3: 【Y704】A(左側) NG1ピックアップ戻 *)
_p43 := ((ST3_A_Dis1_M[2] AND Out_CYw_NG1_Srt_A_H_Done) OR ST3_A_Dis1_M[3] OR ST3_A_Dis1_M[3]) AND NOT ST3_A_Dis1_M[4];
ST3_A_Dis1_M[3] := _p43;
Out_CYw_NG1_Pick_A_H_Auto[1] := _p43;
(* Rung 4: 【Y706】A(左側) NG1チャック戻 *)
_p44 := ((ST3_A_Dis1_M[3] AND Out_CYw_NG1_Pick_A_H_Done) OR ST3_A_Dis1_M[4]) AND NOT ST3_A_Dis1_M[5];
ST3_A_Dis1_M[4] := _p44;
Out_CYw_NG1_Chk_A_H_Auto[1] := _p44;
(* Rung 5: 【Y722】A(左側) 位置3ストッパー戻 *)
_p45 := ((ST3_A_Dis1_M[4] AND Out_CYw_NG1_Chk_A_H_Done) OR ST3_A_Dis1_M[5]) AND NOT ST3_A_Dis1_M[6];
ST3_A_Dis1_M[5] := _p45;
Out_CYS_Pos_03_Stopper_A_H_Auto[2] := _p45;

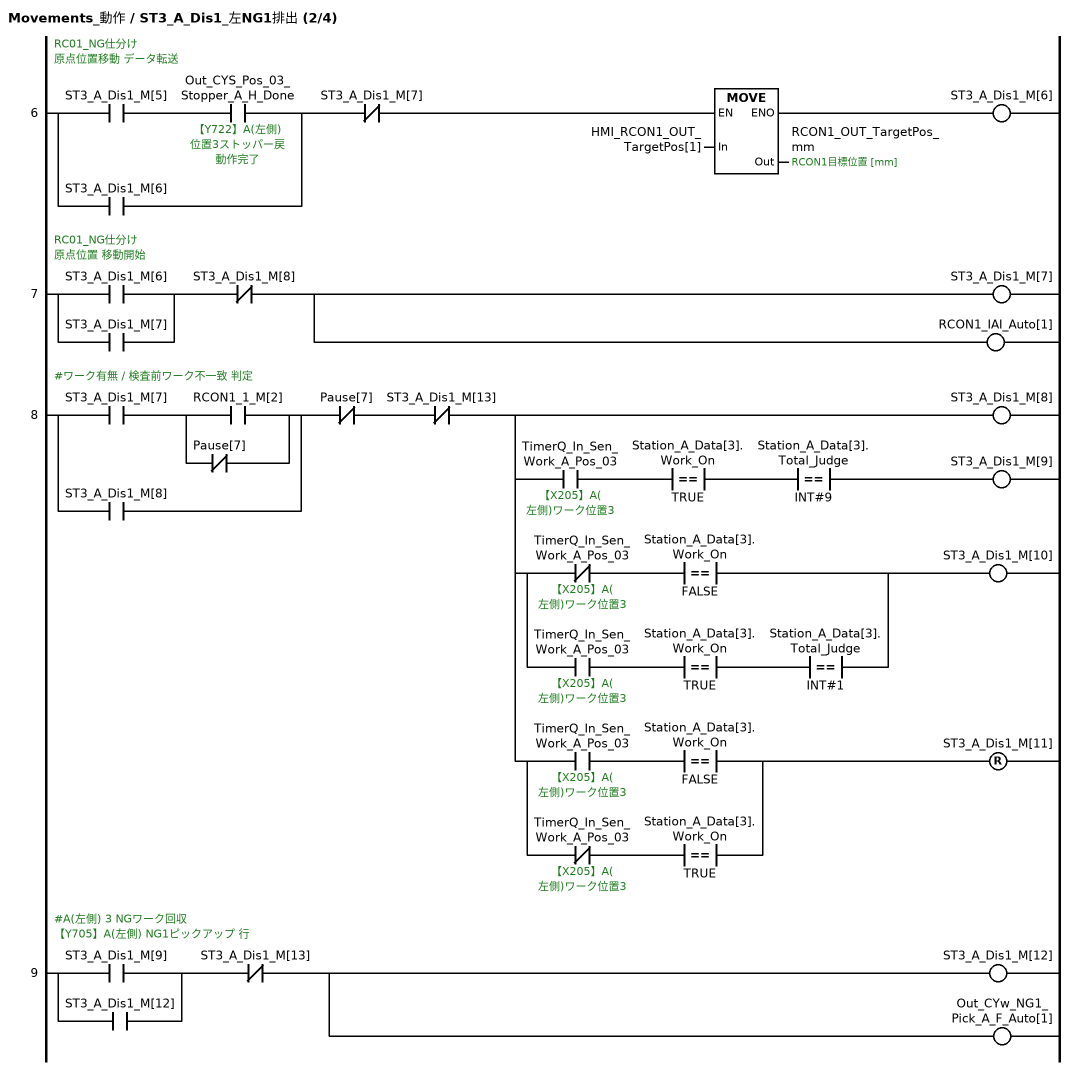
(* Rung 6: RC01_NG仕分け / 原点位置移動 データ転送 *)
IF ((ST3_A_Dis1_M[5] AND Out_CYS_Pos_03_Stopper_A_H_Done) OR ST3_A_Dis1_M[6]) AND NOT ST3_A_Dis1_M[7] THEN
    RCON1_OUT_TargetPos_mm := HMI_RCON1_OUT_TargetPos[1];
END_IF;
ST3_A_Dis1_M[6] := ((ST3_A_Dis1_M[5] AND Out_CYS_Pos_03_Stopper_A_H_Done) OR ST3_A_Dis1_M[6]) AND NOT ST3_A_Dis1_M[7];
(* Rung 7: RC01_NG仕分け / 原点位置 移動開始 *)
_p46 := (ST3_A_Dis1_M[6] OR ST3_A_Dis1_M[7]) AND NOT ST3_A_Dis1_M[8];
ST3_A_Dis1_M[7] := _p46;
RCON1_IAI_Auto[1] := _p46;
(* Rung 8: #ワーク有無 / 検査前ワーク不一致 判定 *)
_p47 := ((ST3_A_Dis1_M[7] AND (RCON1_1_M[2] OR NOT Pause[7])) OR ST3_A_Dis1_M[8]) AND NOT Pause[7] AND NOT ST3_A_Dis1_M[13];
ST3_A_Dis1_M[8] := _p47;
ST3_A_Dis1_M[9] := _p47 AND TimerQ_In_Sen_Work_A_Pos_03 AND (Station_A_Data[3].Work_On = TRUE) AND (Station_A_Data[3].Total_Judge = INT#9);
ST3_A_Dis1_M[10] := _p47 AND ((NOT TimerQ_In_Sen_Work_A_Pos_03 AND (Station_A_Data[3].Work_On = FALSE)) OR (TimerQ_In_Sen_Work_A_Pos_03 AND (Station_A_Data[3].Work_On = TRUE) AND (Station_A_Data[3].Total_Judge = INT#1)));
IF _p47 AND ((TimerQ_In_Sen_Work_A_Pos_03 AND (Station_A_Data[3].Work_On = FALSE)) OR (NOT TimerQ_In_Sen_Work_A_Pos_03 AND (Station_A_Data[3].Work_On = TRUE))) THEN
    ST3_A_Dis1_M[11] := FALSE;
END_IF;
(* Rung 9: #A(左側) 3 NGワーク回収 / 【Y705】A(左側) NG1ピックアップ 行 *)
_p48 := (ST3_A_Dis1_M[9] OR ST3_A_Dis1_M[12]) AND NOT ST3_A_Dis1_M[13];
ST3_A_Dis1_M[12] := _p48;
Out_CYw_NG1_Pick_A_F_Auto[1] := _p48;

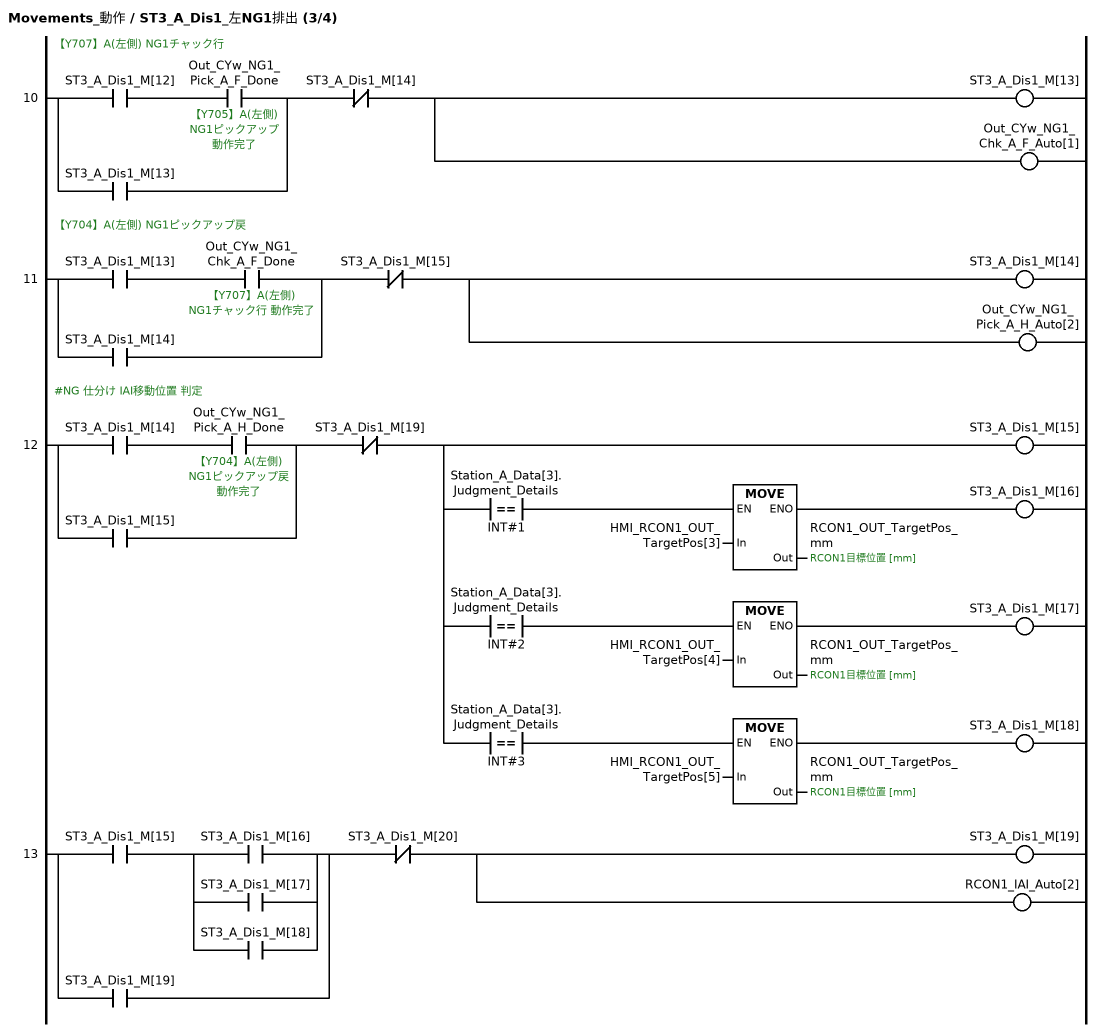
(* Rung 10: 【Y707】A(左側) NG1チャック行 *)
_p49 := ((ST3_A_Dis1_M[12] AND Out_CYw_NG1_Pick_A_F_Done) OR ST3_A_Dis1_M[13]) AND NOT ST3_A_Dis1_M[14];
ST3_A_Dis1_M[13] := _p49;
Out_CYw_NG1_Chk_A_F_Auto[1] := _p49;
(* Rung 11: 【Y704】A(左側) NG1ピックアップ戻 *)
_p50 := ((ST3_A_Dis1_M[13] AND Out_CYw_NG1_Chk_A_F_Done) OR ST3_A_Dis1_M[14]) AND NOT ST3_A_Dis1_M[15];
ST3_A_Dis1_M[14] := _p50;
Out_CYw_NG1_Pick_A_H_Auto[2] := _p50;
(* Rung 12: #NG 仕分け IAI移動位置 判定 *)
_p51 := ((ST3_A_Dis1_M[14] AND Out_CYw_NG1_Pick_A_H_Done) OR ST3_A_Dis1_M[15]) AND NOT ST3_A_Dis1_M[19];
ST3_A_Dis1_M[15] := _p51;
IF _p51 AND (Station_A_Data[3].Judgment_Details = INT#1) THEN
    RCON1_OUT_TargetPos_mm := HMI_RCON1_OUT_TargetPos[3];
END_IF;
ST3_A_Dis1_M[16] := _p51 AND (Station_A_Data[3].Judgment_Details = INT#1);
IF _p51 AND (Station_A_Data[3].Judgment_Details = INT#2) THEN
    RCON1_OUT_TargetPos_mm := HMI_RCON1_OUT_TargetPos[4];
END_IF;
ST3_A_Dis1_M[17] := _p51 AND (Station_A_Data[3].Judgment_Details = INT#2);
IF _p51 AND (Station_A_Data[3].Judgment_Details = INT#3) THEN
    RCON1_OUT_TargetPos_mm := HMI_RCON1_OUT_TargetPos[5];
END_IF;
ST3_A_Dis1_M[18] := _p51 AND (Station_A_Data[3].Judgment_Details = INT#3);
(* Rung 13 *)
_p52 := ((ST3_A_Dis1_M[15] AND (ST3_A_Dis1_M[16] OR ST3_A_Dis1_M[17] OR ST3_A_Dis1_M[18])) OR ST3_A_Dis1_M[19]) AND NOT ST3_A_Dis1_M[20];
ST3_A_Dis1_M[19] := _p52;
RCON1_IAI_Auto[2] := _p52;

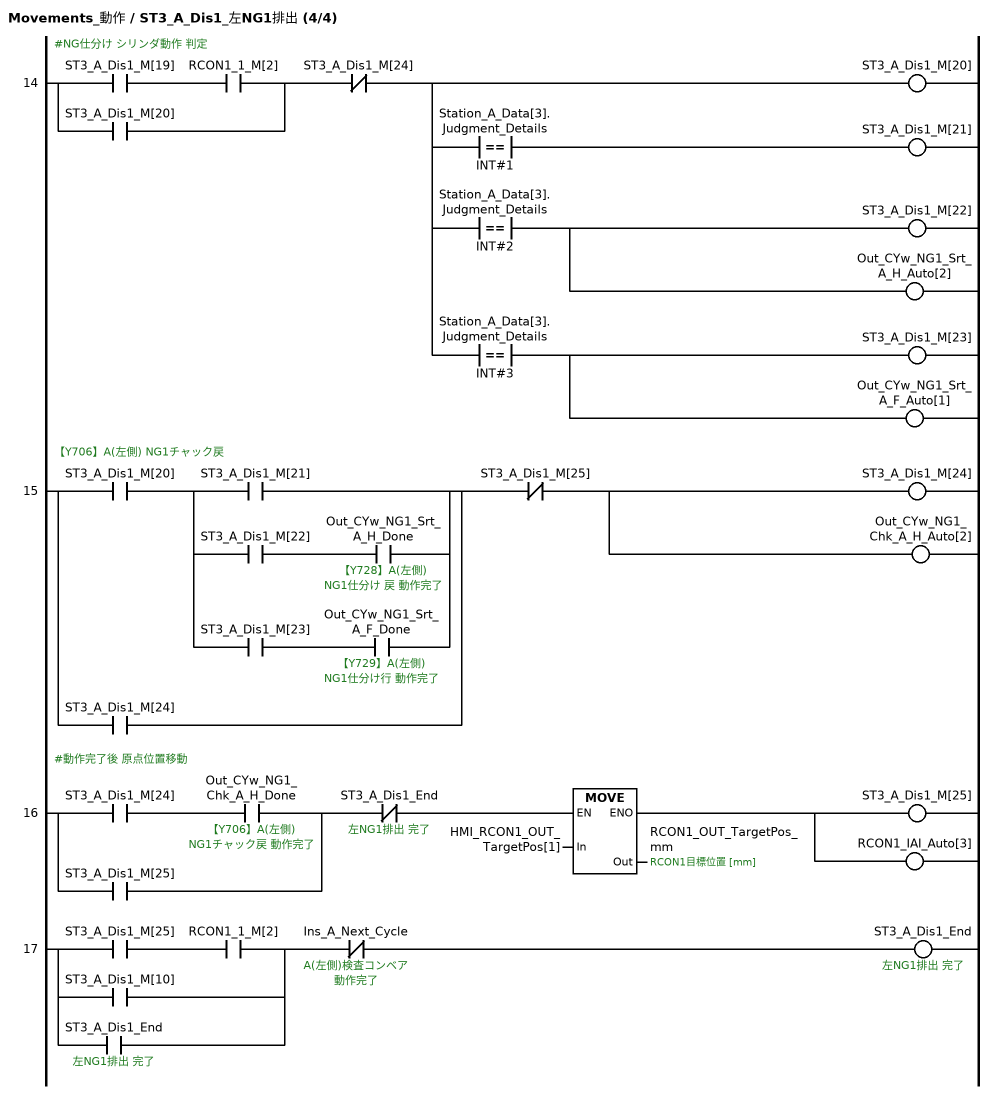
(* Rung 14: #NG仕分け シリンダ動作 判定 *)
_p53 := ((ST3_A_Dis1_M[19] AND RCON1_1_M[2]) OR ST3_A_Dis1_M[20]) AND NOT ST3_A_Dis1_M[24];
ST3_A_Dis1_M[20] := _p53;
ST3_A_Dis1_M[21] := _p53 AND (Station_A_Data[3].Judgment_Details = INT#1);
_p54 := _p53 AND (Station_A_Data[3].Judgment_Details = INT#2);
ST3_A_Dis1_M[22] := _p54;
Out_CYw_NG1_Srt_A_H_Auto[2] := _p54;
_p55 := _p53 AND (Station_A_Data[3].Judgment_Details = INT#3);
ST3_A_Dis1_M[23] := _p55;
Out_CYw_NG1_Srt_A_F_Auto[1] := _p55;
(* Rung 15: 【Y706】A(左側) NG1チャック戻 *)
_p56 := ((ST3_A_Dis1_M[20] AND (ST3_A_Dis1_M[21] OR (ST3_A_Dis1_M[22] AND Out_CYw_NG1_Srt_A_H_Done) OR (ST3_A_Dis1_M[23] AND Out_CYw_NG1_Srt_A_F_Done))) OR ST3_A_Dis1_M[24]) AND NOT ST3_A_Dis1_M[25];
ST3_A_Dis1_M[24] := _p56;
Out_CYw_NG1_Chk_A_H_Auto[2] := _p56;
(* Rung 16: #動作完了後 原点位置移動 *)
IF ((ST3_A_Dis1_M[24] AND Out_CYw_NG1_Chk_A_H_Done) OR ST3_A_Dis1_M[25]) AND NOT ST3_A_Dis1_End THEN
    RCON1_OUT_TargetPos_mm := HMI_RCON1_OUT_TargetPos[1];
END_IF;
_p57 := ((ST3_A_Dis1_M[24] AND Out_CYw_NG1_Chk_A_H_Done) OR ST3_A_Dis1_M[25]) AND NOT ST3_A_Dis1_End;
ST3_A_Dis1_M[25] := _p57;
RCON1_IAI_Auto[3] := _p57;
(* Rung 17 *)
ST3_A_Dis1_End := ((ST3_A_Dis1_M[25] AND RCON1_1_M[2]) OR ST3_A_Dis1_M[10] OR ST3_A_Dis1_End) AND NOT Ins_A_Next_Cycle;

(* Section ST4_A_Rev1_左反転1: ladder, written here as Structured Text *)

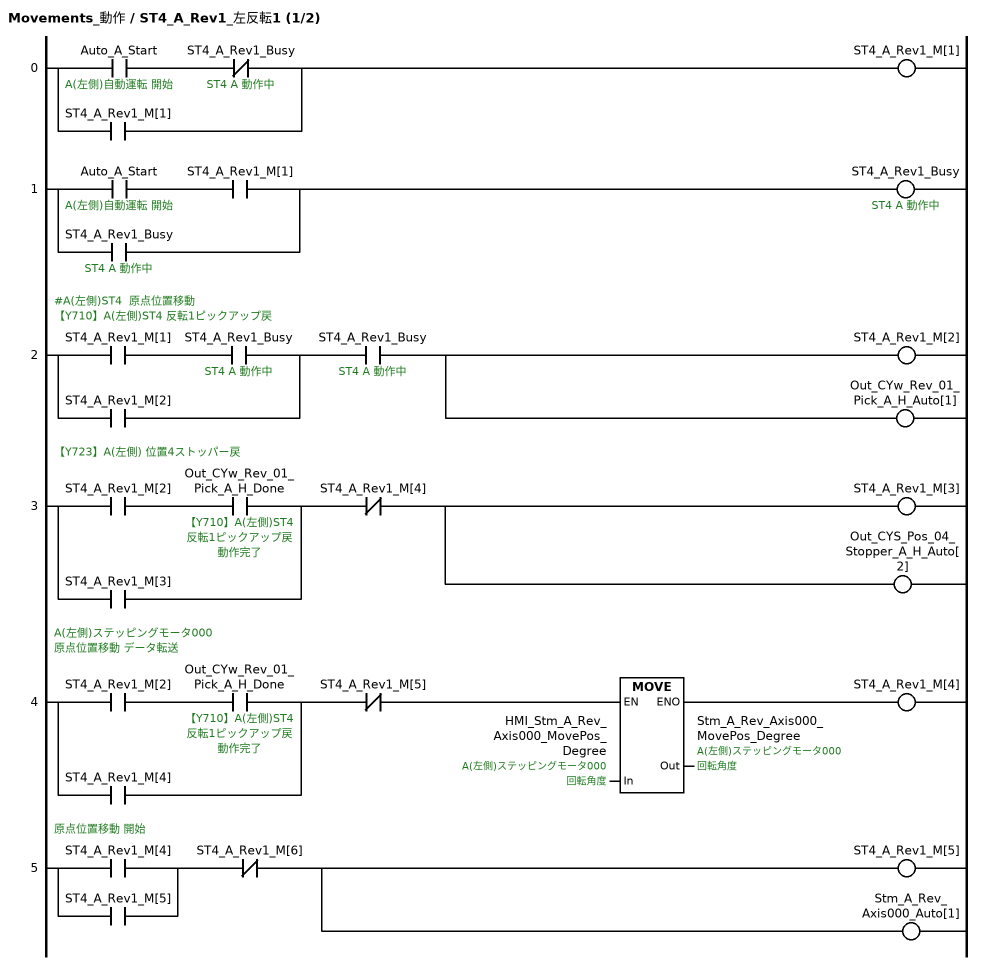
(* Rung 0 *)
ST4_A_Rev1_M[1] := (Auto_A_Start AND NOT ST4_A_Rev1_Busy) OR ST4_A_Rev1_M[1];
(* Rung 1 *)
ST4_A_Rev1_Busy := (Auto_A_Start AND ST4_A_Rev1_M[1]) OR ST4_A_Rev1_Busy;
(* Rung 2: #A(左側)ST4  原点位置移動 / 【Y710】A(左側)ST4 反転1ピックアップ戻 *)
_p58 := ((ST4_A_Rev1_M[1] AND ST4_A_Rev1_Busy) OR ST4_A_Rev1_M[2]) AND ST4_A_Rev1_Busy;
ST4_A_Rev1_M[2] := _p58;
Out_CYw_Rev_01_Pick_A_H_Auto[1] := _p58;
(* Rung 3: 【Y723】A(左側) 位置4ストッパー戻 *)
_p59 := ((ST4_A_Rev1_M[2] AND Out_CYw_Rev_01_Pick_A_H_Done) OR ST4_A_Rev1_M[3]) AND NOT ST4_A_Rev1_M[4];
ST4_A_Rev1_M[3] := _p59;
Out_CYS_Pos_04_Stopper_A_H_Auto[2] := _p59;
(* Rung 4: A(左側)ステッピングモータ000 / 原点位置移動 データ転送 *)
IF ((ST4_A_Rev1_M[2] AND Out_CYw_Rev_01_Pick_A_H_Done) OR ST4_A_Rev1_M[4]) AND NOT ST4_A_Rev1_M[5] THEN
    Stm_A_Rev_Axis000_MovePos_Degree := HMI_Stm_A_Rev_Axis000_MovePos_Degree;
END_IF;
ST4_A_Rev1_M[4] := ((ST4_A_Rev1_M[2] AND Out_CYw_Rev_01_Pick_A_H_Done) OR ST4_A_Rev1_M[4]) AND NOT ST4_A_Rev1_M[5];
(* Rung 5: 原点位置移動 開始 *)
_p60 := (ST4_A_Rev1_M[4] OR ST4_A_Rev1_M[5]) AND NOT ST4_A_Rev1_M[6];
ST4_A_Rev1_M[5] := _p60;
Stm_A_Rev_Axis000_Auto[1] := _p60;

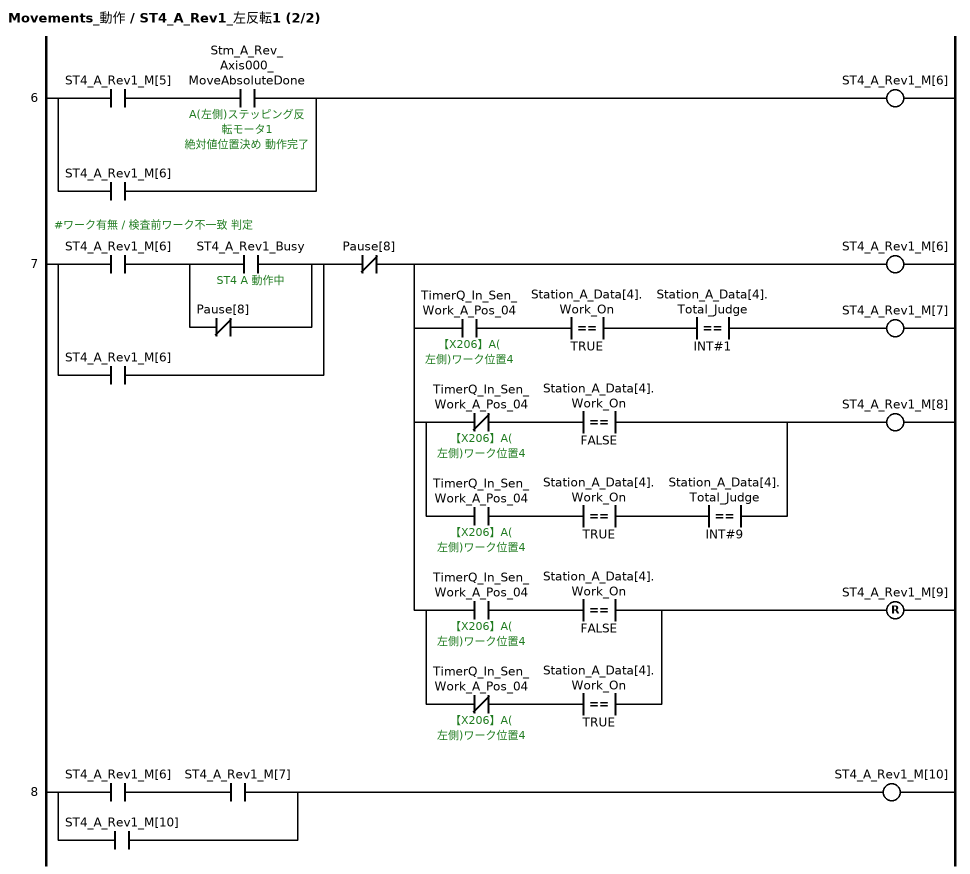
(* Rung 6 *)
ST4_A_Rev1_M[6] := (ST4_A_Rev1_M[5] AND Stm_A_Rev_Axis000_MoveAbsoluteDone) OR ST4_A_Rev1_M[6];
(* Rung 7: #ワーク有無 / 検査前ワーク不一致 判定 *)
_p61 := ((ST4_A_Rev1_M[6] AND (ST4_A_Rev1_Busy OR NOT Pause[8])) OR ST4_A_Rev1_M[6]) AND NOT Pause[8];
ST4_A_Rev1_M[6] := _p61;
ST4_A_Rev1_M[7] := _p61 AND TimerQ_In_Sen_Work_A_Pos_04 AND (Station_A_Data[4].Work_On = TRUE) AND (Station_A_Data[4].Total_Judge = INT#1);
ST4_A_Rev1_M[8] := _p61 AND ((NOT TimerQ_In_Sen_Work_A_Pos_04 AND (Station_A_Data[4].Work_On = FALSE)) OR (TimerQ_In_Sen_Work_A_Pos_04 AND (Station_A_Data[4].Work_On = TRUE) AND (Station_A_Data[4].Total_Judge = INT#9)));
IF _p61 AND ((TimerQ_In_Sen_Work_A_Pos_04 AND (Station_A_Data[4].Work_On = FALSE)) OR (NOT TimerQ_In_Sen_Work_A_Pos_04 AND (Station_A_Data[4].Work_On = TRUE))) THEN
    ST4_A_Rev1_M[9] := FALSE;
END_IF;
(* Rung 8 *)
ST4_A_Rev1_M[10] := (ST4_A_Rev1_M[6] AND ST4_A_Rev1_M[7]) OR ST4_A_Rev1_M[10];
END_PROGRAM

PROGRAM OtherDevice_外部機器
VAR
    FH_M : BOOL;
    GT2_M : BOOL;
    IAI_M : BOOL;  (* 旧ダミーマーカー（ST許可ではない） *)
    HMI_M : BOOL;
    FH_A_ST1_M : ARRAY[0..99] OF Bool;  (* [1] ST1 FH測定中; [5] ST1 測定完了 *)
    FH_A_ST1_OK : BOOL;  (* ST1 OK判定 *)
    FH_A_ST1_NG : BOOL;  (* ST1 NG 判定 *)
    FH_A_ST1_TON : ARRAY[0..99] OF TON;
    FH_A_ST1_TOF : ARRAY[0..99] OF TOF;
    ４ : UINT;
    ConvWordIndex : INT;  (* 作業用 ワード番号 *)
    ConvAxisIndex : INT;  (* 作業用 軸番号（RCON1:1～6／RCON2:1～5） *)
    ConvBase : INT;  (* 作業用 軸先頭ワード番号 *)
    ConvDWord : DWORD;  (* 作業用 32bit分割・結合 *)
    ConvPos : DINT;  (* 作業用 目標位置 [0.01mm・符号付き] *)
    ConvBand : UDINT;  (* 作業用 位置決め幅 [0.01mm] *)
    ConvSpeed : UINT;  (* 作業用 速度送信値 *)
    ConvAccDec : UINT;  (* 作業用 共通加減速 [0.01G] *)
    ConvPush : UINT;  (* 作業用 押付け制限 [255=100%] *)
    ConvScaled : LREAL;  (* 作業用 換算後の小数値 *)
    ConvWord : WORD;  (* 作業用 16bitワード *)
    ConvUnitOK : BOOL;  (* 作業用 速度単位正常 *)
    RCON1_1_TOF : ARRAY[0..99] OF TOF;
    RCON1_1_TON : ARRAY[0..99] OF TON;
    Stm_A_Rev_Axis000_ZeroSet : MC_SetPosition;
    Stm_A_Rev_Axis000_HomeWithParameter : MC_HomeWithParameter;
    Stm_A_Rev_Axis000_Power : MC_Power;  (* A(左側)ステッピングモータ000 電源ON状態 *)
    Stm_A_Rev_Axis000_MoveAbsolute : MC_MoveAbsolute;
    Stm_A_Rev_Axis000_MoveVel : LREAL;  (* 動作速度 *)
    Stm_A_Rev_Axis000_MoveAcc : LREAL;  (* 動作加速度 *)
    Stm_A_Rev_Axis000_MoveDec : LREAL;  (* 動作減速度 *)
    Stm_A_Rev_Axis000_MoveBusy : BOOL;  (* 動作中 *)
    Stm_A_Rev_Axis000_MoveError : BOOL;  (* 動作エラー *)
    Stm_A_Rev_Axis000_TON : ARRAY[0..99] OF TON;
END_VAR
VAR_EXTERNAL
    HMI_MessageNo : ARRAY[0..9] OF UINT;
    HMI_Message : ARRAY[0..9] OF String[256];
    HMI_Language : BOOL;
    FH_Line0_Trigger_Ready_1 : BOOL;
    FH_Line0_Trigger_1 : BOOL;
    M9999 : BOOL;
    FH_Line0_Busy_1 : BOOL;
    FH_Line0_Result_Notification_1 : BOOL;
    FH_Line0_DINT_Result_Data_0_1 : DINT;
    FH_Line0_DINT_Result_Data_1_1 : DINT;
    FH_Line0_DINT_Result_Data_2_1 : DINT;
    FH_Line0_Command_Code_1 : DWORD;
    FH_Line0_Command_Request_1 : BOOL;
    FH_Line0_Command_Completion_1 : BOOL;
    MdlChg : BOOL;  (* 機種切替：ON【GA120】 OFF【GA90】 *)
    FH_Line0_Error_Status_1 : BOOL;
    FH_5552_10_A_Auto : BOOL;  (* ST1 FH測定開始 *)
    FH_A_ST1_Manual : BOOL;  (* ST1 *)
    Pause : ARRAY[0..99] OF Bool;
    FH_A_ST1_Done : BOOL;  (* ST1 画像検査完了 *)
    Station_A_Data : ARRAY[0..8] OF sData;
    DLEP1_OUT : ARRAY[0..79] OF BOOL;
    DLEP2_OUT : ARRAY[0..79] OF BOOL;
    DLEP1_IN : ARRAY[0..167] OF byte;
    DLEP2_IN : ARRAY[0..167] OF byte;
    DLEP2_IN_Error : BOOL;  (* B(右側)センサエラー *)
    DLEP1_IN_Error : BOOL;  (* A(右側)センサエラー *)
    GT2_A_CurrentVal : INT;  (* A(左側) 測定値 *)
    GT2_B_CurrentVal : INT;  (* B(右側) 測定値 *)
    Hgt_A_Ins_Data : LREAL;  (* A測定データに変換 *)
    Hgt_B_Ins_Data : LREAL;
    Hgt_A_ComputedValueData : LREAL;  (* A測定データ+13.000mm 算定データ *)
    Hgt_B_ComputedValueData : LREAL;  (* B測定データ+13.000mm 算定データ *)
    E001_In_IN00_2004_01 : UINT;  (* RCON1 IN00 GW状態 *)
    E001_In_IN01_2004_02 : UINT;  (* RCON1 IN01 軸リンク状態 *)
    E001_In_IN02_2004_03 : UINT;  (* RCON1 IN02 電源状態0 *)
    E001_In_IN03_2004_04 : UINT;  (* RCON1 IN03 電源状態1 *)
    E001_In_IN04_2004_05 : UINT;  (* RCON1 IN04 電源状態2 *)
    E001_In_IN05_2004_06 : UINT;  (* RCON1 IN05 電源状態3 *)
    E001_In_IN06_2004_07 : UINT;  (* RCON1 IN06 電源状態4（構成依存） *)
    E001_In_IN07_2004_08 : UINT;  (* RCON1 IN07 予約（使用禁止） *)
    E001_In_IN08_2004_09 : UINT;  (* RCON1 IN08 1軸目 現在位置 下位 [0.01mm] *)
    E001_In_IN09_2004_0A : UINT;  (* RCON1 IN09 1軸目 現在位置 上位 [0.01mm] *)
    E001_In_IN10_2004_0B : UINT;  (* RCON1 IN10 1軸目 指令電流 下位 [mA] *)
    E001_In_IN11_2004_0C : UINT;  (* RCON1 IN11 1軸目 指令電流 上位 [mA] *)
    E001_In_IN12_2004_0D : UINT;  (* RCON1 IN12 1軸目 現在速度 [実機単位・符号付き] *)
    E001_In_IN13_2004_0E : UINT;  (* RCON1 IN13 1軸目 予約（使用禁止） *)
    E001_In_IN14_2004_0F : UINT;  (* RCON1 IN14 1軸目 軸異常コード *)
    E001_In_IN15_2004_10 : UINT;  (* RCON1 IN15 1軸目 状態信号（PEND/SV等） *)
    E001_In_IN16_2004_11 : UINT;  (* RCON1 IN16 2軸目 現在位置 下位 [0.01mm] *)
    E001_In_IN17_2004_12 : UINT;  (* RCON1 IN17 2軸目 現在位置 上位 [0.01mm] *)
    E001_In_IN18_2004_13 : UINT;  (* RCON1 IN18 2軸目 指令電流 下位 [mA] *)
    E001_In_IN19_2004_14 : UINT;  (* RCON1 IN19 2軸目 指令電流 上位 [mA] *)
    E001_In_IN20_2004_15 : UINT;  (* RCON1 IN20 2軸目 現在速度 [実機単位・符号付き] *)
    E001_In_IN21_2004_16 : UINT;  (* RCON1 IN21 2軸目 予約（使用禁止） *)
    E001_In_IN22_2004_17 : UINT;  (* RCON1 IN22 2軸目 軸異常コード *)
    E001_In_IN23_2004_18 : UINT;  (* RCON1 IN23 2軸目 状態信号（PEND/SV等） *)
    E001_In_IN24_2004_19 : UINT;  (* RCON1 IN24 3軸目 現在位置 下位 [0.01mm] *)
    E001_In_IN25_2004_1A : UINT;  (* RCON1 IN25 3軸目 現在位置 上位 [0.01mm] *)
    E001_In_IN26_2004_1B : UINT;  (* RCON1 IN26 3軸目 指令電流 下位 [mA] *)
    E001_In_IN27_2004_1C : UINT;  (* RCON1 IN27 3軸目 指令電流 上位 [mA] *)
    E001_In_IN28_2004_1D : UINT;  (* RCON1 IN28 3軸目 現在速度 [実機単位・符号付き] *)
    E001_In_IN29_2004_1E : UINT;  (* RCON1 IN29 3軸目 予約（使用禁止） *)
    E001_In_IN30_2004_1F : UINT;  (* RCON1 IN30 3軸目 軸異常コード *)
    E001_In_IN31_2004_20 : UINT;  (* RCON1 IN31 3軸目 状態信号（PEND/SV等） *)
    E001_In_IN32_2004_21 : UINT;  (* RCON1 IN32 4軸目 現在位置 下位 [0.01mm] *)
    E001_In_IN33_2004_22 : UINT;  (* RCON1 IN33 4軸目 現在位置 上位 [0.01mm] *)
    E001_In_IN34_2004_23 : UINT;  (* RCON1 IN34 4軸目 指令電流 下位 [mA] *)
    E001_In_IN35_2004_24 : UINT;  (* RCON1 IN35 4軸目 指令電流 上位 [mA] *)
    E001_In_IN36_2004_25 : UINT;  (* RCON1 IN36 4軸目 現在速度 [実機単位・符号付き] *)
    E001_In_IN37_2004_26 : UINT;  (* RCON1 IN37 4軸目 予約（使用禁止） *)
    E001_In_IN38_2004_27 : UINT;  (* RCON1 IN38 4軸目 軸異常コード *)
    E001_In_IN39_2004_28 : UINT;  (* RCON1 IN39 4軸目 状態信号（PEND/SV等） *)
    E001_In_IN40_2004_29 : UINT;  (* RCON1 IN40 5軸目 現在位置 下位 [0.01mm] *)
    E001_In_IN41_2004_2A : UINT;  (* RCON1 IN41 5軸目 現在位置 上位 [0.01mm] *)
    E001_In_IN42_2004_2B : UINT;  (* RCON1 IN42 5軸目 指令電流 下位 [mA] *)
    E001_In_IN43_2004_2C : UINT;  (* RCON1 IN43 5軸目 指令電流 上位 [mA] *)
    E001_In_IN44_2004_2D : UINT;  (* RCON1 IN44 5軸目 現在速度 [実機単位・符号付き] *)
    E001_In_IN45_2004_2E : UINT;  (* RCON1 IN45 5軸目 予約（使用禁止） *)
    E001_In_IN46_2004_2F : UINT;  (* RCON1 IN46 5軸目 軸異常コード *)
    E001_In_IN47_2004_30 : UINT;  (* RCON1 IN47 5軸目 状態信号（PEND/SV等） *)
    E001_In_IN48_2004_31 : UINT;  (* RCON1 IN48 6軸目 現在位置 下位 [0.01mm] *)
    E001_In_IN49_2004_32 : UINT;  (* RCON1 IN49 6軸目 現在位置 上位 [0.01mm] *)
    E001_In_IN50_2004_33 : UINT;  (* RCON1 IN50 6軸目 指令電流 下位 [mA] *)
    E001_In_IN51_2004_34 : UINT;  (* RCON1 IN51 6軸目 指令電流 上位 [mA] *)
    E001_In_IN52_2004_35 : UINT;  (* RCON1 IN52 6軸目 現在速度 [実機単位・符号付き] *)
    E001_In_IN53_2004_36 : UINT;  (* RCON1 IN53 6軸目 予約（使用禁止） *)
    E001_In_IN54_2004_37 : UINT;  (* RCON1 IN54 6軸目 軸異常コード *)
    E001_In_IN55_2004_38 : UINT;  (* RCON1 IN55 6軸目 状態信号（PEND/SV等） *)
    E001_In_IN56_2004_39 : UINT;  (* RCON1 IN56 112Byte範囲外（未割付・不使用） *)
    E001_In_IN57_2004_3A : UINT;  (* RCON1 IN57 112Byte範囲外（未割付・不使用） *)
    E001_In_IN58_2004_3B : UINT;  (* RCON1 IN58 112Byte範囲外（未割付・不使用） *)
    E001_In_IN59_2004_3C : UINT;  (* RCON1 IN59 112Byte範囲外（未割付・不使用） *)
    E001_In_IN60_2004_3D : UINT;  (* RCON1 IN60 112Byte範囲外（未割付・不使用） *)
    E001_In_IN61_2004_3E : UINT;  (* RCON1 IN61 112Byte範囲外（未割付・不使用） *)
    E001_In_IN62_2004_3F : UINT;  (* RCON1 IN62 112Byte範囲外（未割付・不使用） *)
    E001_In_IN63_2004_40 : UINT;  (* RCON1 IN63 112Byte範囲外（未割付・不使用） *)
    E001_In_IN64_2004_41 : UINT;  (* RCON1 IN64 112Byte範囲外（未割付・不使用） *)
    E001_In_IN65_2004_42 : UINT;  (* RCON1 IN65 112Byte範囲外（未割付・不使用） *)
    E001_In_IN66_2004_43 : UINT;  (* RCON1 IN66 112Byte範囲外（未割付・不使用） *)
    E001_In_IN67_2004_44 : UINT;  (* RCON1 IN67 112Byte範囲外（未割付・不使用） *)
    E001_In_IN68_2004_45 : UINT;  (* RCON1 IN68 112Byte範囲外（未割付・不使用） *)
    E001_In_IN69_2004_46 : UINT;  (* RCON1 IN69 112Byte範囲外（未割付・不使用） *)
    E001_In_IN70_2004_47 : UINT;  (* RCON1 IN70 112Byte範囲外（未割付・不使用） *)
    E001_In_IN71_2004_48 : UINT;  (* RCON1 IN71 112Byte範囲外（未割付・不使用） *)
    E001_Out_OUT00_2003_01 : UINT;  (* RCON1 OUT00 共通制御（MON/RTE） *)
    E001_Out_OUT08_2003_09 : UINT;  (* RCON1 OUT08 1軸目 目標位置 下位 [0.01mm] *)
    E001_Out_OUT09_2003_0A : UINT;  (* RCON1 OUT09 1軸目 目標位置 上位 [0.01mm] *)
    E001_Out_OUT10_2003_0B : UINT;  (* RCON1 OUT10 1軸目 位置決め幅 下位 [0.01mm] *)
    E001_Out_OUT11_2003_0C : UINT;  (* RCON1 OUT11 1軸目 位置決め幅 上位 [0.01mm] *)
    E001_Out_OUT12_2003_0D : UINT;  (* RCON1 OUT12 1軸目 速度指令 [実機単位] *)
    E001_Out_OUT13_2003_0E : UINT;  (* RCON1 OUT13 1軸目 共通加減速 [0.01G] *)
    E001_Out_OUT14_2003_0F : UINT;  (* RCON1 OUT14 1軸目 押付け制限 [255=100%] *)
    E001_Out_OUT15_2003_10 : UINT;  (* RCON1 OUT15 1軸目 制御信号（DSTR/SON等） *)
    E001_Out_OUT16_2003_11 : UINT;  (* RCON1 OUT16 2軸目 目標位置 下位 [0.01mm] *)
    E001_Out_OUT17_2003_12 : UINT;  (* RCON1 OUT17 2軸目 目標位置 上位 [0.01mm] *)
    E001_Out_OUT18_2003_13 : UINT;  (* RCON1 OUT18 2軸目 位置決め幅 下位 [0.01mm] *)
    E001_Out_OUT19_2003_14 : UINT;  (* RCON1 OUT19 2軸目 位置決め幅 上位 [0.01mm] *)
    E001_Out_OUT20_2003_15 : UINT;  (* RCON1 OUT20 2軸目 速度指令 [実機単位] *)
    E001_Out_OUT21_2003_16 : UINT;  (* RCON1 OUT21 2軸目 共通加減速 [0.01G] *)
    E001_Out_OUT22_2003_17 : UINT;  (* RCON1 OUT22 2軸目 押付け制限 [255=100%] *)
    E001_Out_OUT23_2003_18 : UINT;  (* RCON1 OUT23 2軸目 制御信号（DSTR/SON等） *)
    E001_Out_OUT24_2003_19 : UINT;  (* RCON1 OUT24 3軸目 目標位置 下位 [0.01mm] *)
    E001_Out_OUT25_2003_1A : UINT;  (* RCON1 OUT25 3軸目 目標位置 上位 [0.01mm] *)
    E001_Out_OUT26_2003_1B : UINT;  (* RCON1 OUT26 3軸目 位置決め幅 下位 [0.01mm] *)
    E001_Out_OUT27_2003_1C : UINT;  (* RCON1 OUT27 3軸目 位置決め幅 上位 [0.01mm] *)
    E001_Out_OUT28_2003_1D : UINT;  (* RCON1 OUT28 3軸目 速度指令 [実機単位] *)
    E001_Out_OUT29_2003_1E : UINT;  (* RCON1 OUT29 3軸目 共通加減速 [0.01G] *)
    E001_Out_OUT30_2003_1F : UINT;  (* RCON1 OUT30 3軸目 押付け制限 [255=100%] *)
    E001_Out_OUT31_2003_20 : UINT;  (* RCON1 OUT31 3軸目 制御信号（DSTR/SON等） *)
    E001_Out_OUT32_2003_21 : UINT;  (* RCON1 OUT32 4軸目 目標位置 下位 [0.01mm] *)
    E001_Out_OUT33_2003_22 : UINT;  (* RCON1 OUT33 4軸目 目標位置 上位 [0.01mm] *)
    E001_Out_OUT34_2003_23 : UINT;  (* RCON1 OUT34 4軸目 位置決め幅 下位 [0.01mm] *)
    E001_Out_OUT35_2003_24 : UINT;  (* RCON1 OUT35 4軸目 位置決め幅 上位 [0.01mm] *)
    E001_Out_OUT36_2003_25 : UINT;  (* RCON1 OUT36 4軸目 速度指令 [実機単位] *)
    E001_Out_OUT37_2003_26 : UINT;  (* RCON1 OUT37 4軸目 共通加減速 [0.01G] *)
    E001_Out_OUT38_2003_27 : UINT;  (* RCON1 OUT38 4軸目 押付け制限 [255=100%] *)
    E001_Out_OUT39_2003_28 : UINT;  (* RCON1 OUT39 4軸目 制御信号（DSTR/SON等） *)
    E001_Out_OUT40_2003_29 : UINT;  (* RCON1 OUT40 5軸目 目標位置 下位 [0.01mm] *)
    E001_Out_OUT41_2003_2A : UINT;  (* RCON1 OUT41 5軸目 目標位置 上位 [0.01mm] *)
    E001_Out_OUT42_2003_2B : UINT;  (* RCON1 OUT42 5軸目 位置決め幅 下位 [0.01mm] *)
    E001_Out_OUT43_2003_2C : UINT;  (* RCON1 OUT43 5軸目 位置決め幅 上位 [0.01mm] *)
    E001_Out_OUT44_2003_2D : UINT;  (* RCON1 OUT44 5軸目 速度指令 [実機単位] *)
    E001_Out_OUT45_2003_2E : UINT;  (* RCON1 OUT45 5軸目 共通加減速 [0.01G] *)
    E001_Out_OUT46_2003_2F : UINT;  (* RCON1 OUT46 5軸目 押付け制限 [255=100%] *)
    E001_Out_OUT47_2003_30 : UINT;  (* RCON1 OUT47 5軸目 制御信号（DSTR/SON等） *)
    E001_Out_OUT48_2003_31 : UINT;  (* RCON1 OUT48 6軸目 目標位置 下位 [0.01mm] *)
    E001_Out_OUT49_2003_32 : UINT;  (* RCON1 OUT49 6軸目 目標位置 上位 [0.01mm] *)
    E001_Out_OUT50_2003_33 : UINT;  (* RCON1 OUT50 6軸目 位置決め幅 下位 [0.01mm] *)
    E001_Out_OUT51_2003_34 : UINT;  (* RCON1 OUT51 6軸目 位置決め幅 上位 [0.01mm] *)
    E001_Out_OUT52_2003_35 : UINT;  (* RCON1 OUT52 6軸目 速度指令 [実機単位] *)
    E001_Out_OUT53_2003_36 : UINT;  (* RCON1 OUT53 6軸目 共通加減速 [0.01G] *)
    E001_Out_OUT54_2003_37 : UINT;  (* RCON1 OUT54 6軸目 押付け制限 [255=100%] *)
    E001_Out_OUT55_2003_38 : UINT;  (* RCON1 OUT55 6軸目 制御信号（DSTR/SON等） *)
    E005_In_IN00_2004_01_1 : UINT;  (* RCON2 IN00 GW状態 *)
    E005_In_IN01_2004_02_1 : UINT;  (* RCON2 IN01 軸リンク状態 *)
    E005_In_IN02_2004_03_1 : UINT;  (* RCON2 IN02 電源状態0 *)
    E005_In_IN03_2004_04_1 : UINT;  (* RCON2 IN03 電源状態1 *)
    E005_In_IN04_2004_05_1 : UINT;  (* RCON2 IN04 電源状態2 *)
    E005_In_IN05_2004_06_1 : UINT;  (* RCON2 IN05 電源状態3 *)
    E005_In_IN06_2004_07_1 : UINT;  (* RCON2 IN06 電源状態4（構成依存） *)
    E005_In_IN07_2004_08_1 : UINT;  (* RCON2 IN07 予約（使用禁止） *)
    E005_In_IN08_2004_09_1 : UINT;  (* RCON2 IN08 1軸目 現在位置 下位 [0.01mm] *)
    E005_In_IN09_2004_0A_1 : UINT;  (* RCON2 IN09 1軸目 現在位置 上位 [0.01mm] *)
    E005_In_IN10_2004_0B_1 : UINT;  (* RCON2 IN10 1軸目 指令電流 下位 [mA] *)
    E005_In_IN11_2004_0C_1 : UINT;  (* RCON2 IN11 1軸目 指令電流 上位 [mA] *)
    E005_In_IN12_2004_0D_1 : UINT;  (* RCON2 IN12 1軸目 現在速度 [実機単位・符号付き] *)
    E005_In_IN13_2004_0E_1 : UINT;  (* RCON2 IN13 1軸目 予約（使用禁止） *)
    E005_In_IN14_2004_0F_1 : UINT;  (* RCON2 IN14 1軸目 軸異常コード *)
    E005_In_IN15_2004_10_1 : UINT;  (* RCON2 IN15 1軸目 状態信号（PEND/SV等） *)
    E005_In_IN16_2004_11_1 : UINT;  (* RCON2 IN16 2軸目 現在位置 下位 [0.01mm] *)
    E005_In_IN17_2004_12_1 : UINT;  (* RCON2 IN17 2軸目 現在位置 上位 [0.01mm] *)
    E005_In_IN18_2004_13_1 : UINT;  (* RCON2 IN18 2軸目 指令電流 下位 [mA] *)
    E005_In_IN19_2004_14_1 : UINT;  (* RCON2 IN19 2軸目 指令電流 上位 [mA] *)
    E005_In_IN20_2004_15_1 : UINT;  (* RCON2 IN20 2軸目 現在速度 [実機単位・符号付き] *)
    E005_In_IN21_2004_16_1 : UINT;  (* RCON2 IN21 2軸目 予約（使用禁止） *)
    E005_In_IN22_2004_17_1 : UINT;  (* RCON2 IN22 2軸目 軸異常コード *)
    E005_In_IN23_2004_18_1 : UINT;  (* RCON2 IN23 2軸目 状態信号（PEND/SV等） *)
    E005_In_IN24_2004_19_1 : UINT;  (* RCON2 IN24 3軸目 現在位置 下位 [0.01mm] *)
    E005_In_IN25_2004_1A_1 : UINT;  (* RCON2 IN25 3軸目 現在位置 上位 [0.01mm] *)
    E005_In_IN26_2004_1B_1 : UINT;  (* RCON2 IN26 3軸目 指令電流 下位 [mA] *)
    E005_In_IN27_2004_1C_1 : UINT;  (* RCON2 IN27 3軸目 指令電流 上位 [mA] *)
    E005_In_IN28_2004_1D_1 : UINT;  (* RCON2 IN28 3軸目 現在速度 [実機単位・符号付き] *)
    E005_In_IN29_2004_1E_1 : UINT;  (* RCON2 IN29 3軸目 予約（使用禁止） *)
    E005_In_IN30_2004_1F_1 : UINT;  (* RCON2 IN30 3軸目 軸異常コード *)
    E005_In_IN31_2004_20_1 : UINT;  (* RCON2 IN31 3軸目 状態信号（PEND/SV等） *)
    E005_In_IN32_2004_21_1 : UINT;  (* RCON2 IN32 4軸目 現在位置 下位 [0.01mm] *)
    E005_In_IN33_2004_22_1 : UINT;  (* RCON2 IN33 4軸目 現在位置 上位 [0.01mm] *)
    E005_In_IN34_2004_23_1 : UINT;  (* RCON2 IN34 4軸目 指令電流 下位 [mA] *)
    E005_In_IN35_2004_24_1 : UINT;  (* RCON2 IN35 4軸目 指令電流 上位 [mA] *)
    E005_In_IN36_2004_25_1 : UINT;  (* RCON2 IN36 4軸目 現在速度 [実機単位・符号付き] *)
    E005_In_IN37_2004_26_1 : UINT;  (* RCON2 IN37 4軸目 予約（使用禁止） *)
    E005_In_IN38_2004_27_1 : UINT;  (* RCON2 IN38 4軸目 軸異常コード *)
    E005_In_IN39_2004_28_1 : UINT;  (* RCON2 IN39 4軸目 状態信号（PEND/SV等） *)
    E005_In_IN40_2004_29_1 : UINT;  (* RCON2 IN40 5軸目 現在位置 下位 [0.01mm] *)
    E005_In_IN41_2004_2A_1 : UINT;  (* RCON2 IN41 5軸目 現在位置 上位 [0.01mm] *)
    E005_In_IN42_2004_2B_1 : UINT;  (* RCON2 IN42 5軸目 指令電流 下位 [mA] *)
    E005_In_IN43_2004_2C_1 : UINT;  (* RCON2 IN43 5軸目 指令電流 上位 [mA] *)
    E005_In_IN44_2004_2D_1 : UINT;  (* RCON2 IN44 5軸目 現在速度 [実機単位・符号付き] *)
    E005_In_IN45_2004_2E_1 : UINT;  (* RCON2 IN45 5軸目 予約（使用禁止） *)
    E005_In_IN46_2004_2F_1 : UINT;  (* RCON2 IN46 5軸目 軸異常コード *)
    E005_In_IN47_2004_30_1 : UINT;  (* RCON2 IN47 5軸目 状態信号（PEND/SV等） *)
    E005_In_IN48_2004_31_1 : UINT;  (* RCON2 IN48 用途未確認（今回未使用） *)
    E005_In_IN49_2004_32_1 : UINT;  (* RCON2 IN49 用途未確認（今回未使用） *)
    E005_In_IN50_2004_33_1 : UINT;  (* RCON2 IN50 用途未確認（今回未使用） *)
    E005_In_IN51_2004_34_1 : UINT;  (* RCON2 IN51 用途未確認（今回未使用） *)
    E005_In_IN52_2004_35_1 : UINT;  (* RCON2 IN52 用途未確認（今回未使用） *)
    E005_In_IN53_2004_36_1 : UINT;  (* RCON2 IN53 用途未確認（今回未使用） *)
    E005_In_IN54_2004_37_1 : UINT;  (* RCON2 IN54 用途未確認（今回未使用） *)
    E005_In_IN55_2004_38_1 : UINT;  (* RCON2 IN55 用途未確認（今回未使用） *)
    E005_Out_OUT00_2003_01_1 : UINT;  (* RCON2 OUT00 共通制御（MON/RTE） *)
    E005_Out_OUT08_2003_09_1 : UINT;  (* RCON2 OUT08 1軸目 目標位置 下位 [0.01mm] *)
    E005_Out_OUT09_2003_0A_1 : UINT;  (* RCON2 OUT09 1軸目 目標位置 上位 [0.01mm] *)
    E005_Out_OUT10_2003_0B_1 : UINT;  (* RCON2 OUT10 1軸目 位置決め幅 下位 [0.01mm] *)
    E005_Out_OUT11_2003_0C_1 : UINT;  (* RCON2 OUT11 1軸目 位置決め幅 上位 [0.01mm] *)
    E005_Out_OUT12_2003_0D_1 : UINT;  (* RCON2 OUT12 1軸目 速度指令 [実機単位] *)
    E005_Out_OUT13_2003_0E_1 : UINT;  (* RCON2 OUT13 1軸目 共通加減速 [0.01G] *)
    E005_Out_OUT14_2003_0F_1 : UINT;  (* RCON2 OUT14 1軸目 押付け制限 [255=100%] *)
    E005_Out_OUT15_2003_10_1 : UINT;  (* RCON2 OUT15 1軸目 制御信号（DSTR/SON等） *)
    E005_Out_OUT16_2003_11_1 : UINT;  (* RCON2 OUT16 2軸目 目標位置 下位 [0.01mm] *)
    E005_Out_OUT17_2003_12_1 : UINT;  (* RCON2 OUT17 2軸目 目標位置 上位 [0.01mm] *)
    E005_Out_OUT18_2003_13_1 : UINT;  (* RCON2 OUT18 2軸目 位置決め幅 下位 [0.01mm] *)
    E005_Out_OUT19_2003_14_1 : UINT;  (* RCON2 OUT19 2軸目 位置決め幅 上位 [0.01mm] *)
    E005_Out_OUT20_2003_15_1 : UINT;  (* RCON2 OUT20 2軸目 速度指令 [実機単位] *)
    E005_Out_OUT21_2003_16_1 : UINT;  (* RCON2 OUT21 2軸目 共通加減速 [0.01G] *)
    E005_Out_OUT22_2003_17_1 : UINT;  (* RCON2 OUT22 2軸目 押付け制限 [255=100%] *)
    E005_Out_OUT23_2003_18_1 : UINT;  (* RCON2 OUT23 2軸目 制御信号（DSTR/SON等） *)
    E005_Out_OUT24_2003_19_1 : UINT;  (* RCON2 OUT24 3軸目 目標位置 下位 [0.01mm] *)
    E005_Out_OUT25_2003_1A_1 : UINT;  (* RCON2 OUT25 3軸目 目標位置 上位 [0.01mm] *)
    E005_Out_OUT26_2003_1B_1 : UINT;  (* RCON2 OUT26 3軸目 位置決め幅 下位 [0.01mm] *)
    E005_Out_OUT27_2003_1C_1 : UINT;  (* RCON2 OUT27 3軸目 位置決め幅 上位 [0.01mm] *)
    E005_Out_OUT28_2003_1D_1 : UINT;  (* RCON2 OUT28 3軸目 速度指令 [実機単位] *)
    E005_Out_OUT29_2003_1E_1 : UINT;  (* RCON2 OUT29 3軸目 共通加減速 [0.01G] *)
    E005_Out_OUT30_2003_1F_1 : UINT;  (* RCON2 OUT30 3軸目 押付け制限 [255=100%] *)
    E005_Out_OUT31_2003_20_1 : UINT;  (* RCON2 OUT31 3軸目 制御信号（DSTR/SON等） *)
    E005_Out_OUT32_2003_21_1 : UINT;  (* RCON2 OUT32 4軸目 目標位置 下位 [0.01mm] *)
    E005_Out_OUT33_2003_22_1 : UINT;  (* RCON2 OUT33 4軸目 目標位置 上位 [0.01mm] *)
    E005_Out_OUT34_2003_23_1 : UINT;  (* RCON2 OUT34 4軸目 位置決め幅 下位 [0.01mm] *)
    E005_Out_OUT35_2003_24_1 : UINT;  (* RCON2 OUT35 4軸目 位置決め幅 上位 [0.01mm] *)
    E005_Out_OUT36_2003_25_1 : UINT;  (* RCON2 OUT36 4軸目 速度指令 [実機単位] *)
    E005_Out_OUT37_2003_26_1 : UINT;  (* RCON2 OUT37 4軸目 共通加減速 [0.01G] *)
    E005_Out_OUT38_2003_27_1 : UINT;  (* RCON2 OUT38 4軸目 押付け制限 [255=100%] *)
    E005_Out_OUT39_2003_28_1 : UINT;  (* RCON2 OUT39 4軸目 制御信号（DSTR/SON等） *)
    E005_Out_OUT40_2003_29_1 : UINT;  (* RCON2 OUT40 5軸目 目標位置 下位 [0.01mm] *)
    E005_Out_OUT41_2003_2A_1 : UINT;  (* RCON2 OUT41 5軸目 目標位置 上位 [0.01mm] *)
    E005_Out_OUT42_2003_2B_1 : UINT;  (* RCON2 OUT42 5軸目 位置決め幅 下位 [0.01mm] *)
    E005_Out_OUT43_2003_2C_1 : UINT;  (* RCON2 OUT43 5軸目 位置決め幅 上位 [0.01mm] *)
    E005_Out_OUT44_2003_2D_1 : UINT;  (* RCON2 OUT44 5軸目 速度指令 [実機単位] *)
    E005_Out_OUT45_2003_2E_1 : UINT;  (* RCON2 OUT45 5軸目 共通加減速 [0.01G] *)
    E005_Out_OUT46_2003_2F_1 : UINT;  (* RCON2 OUT46 5軸目 押付け制限 [255=100%] *)
    E005_Out_OUT47_2003_30_1 : UINT;  (* RCON2 OUT47 5軸目 制御信号（DSTR/SON等） *)
    RCON1_AxisApply : ARRAY[1..6] OF BOOL;  (* RCON1 軸別出力更新許可（OFF=前値保持）; [1] 1軸目（No.0）出力更新許可（OFF=前値保持）; [2] 2軸目（No.1）出力更新許可（OFF=前値保持）; [3] 3軸目（No.2）出力更新許可（OFF=前値保持）; [4] 4軸目（No.3）出力更新許可（OFF=前値保持）; [5] 5軸目（No.4）出力更新許可（OFF=前値保持）; [6] 6軸目（No.5）出力更新許可（OFF=前値保持） *)
    RCON1_AxisLinked : ARRAY[1..6] OF BOOL;  (* RCON1 軸別リンク状態; [1] 1軸目（No.0）リンク状態; [2] 2軸目（No.1）リンク状態; [3] 3軸目（No.2）リンク状態; [4] 4軸目（No.3）リンク状態; [5] 5軸目（No.4）リンク状態; [6] 6軸目（No.5）リンク状態 *)
    RCON1_AxisWritten : ARRAY[1..6] OF BOOL;  (* RCON1 軸別出力代入済み（RCON受付とは別）; [1] 1軸目（No.0）出力代入済み（RCON受付とは別）; [2] 2軸目（No.1）出力代入済み（RCON受付とは別）; [3] 3軸目（No.2）出力代入済み（RCON受付とは別）; [4] 4軸目（No.3）出力代入済み（RCON受付とは別）; [5] 5軸目（No.4）出力代入済み（RCON受付とは別）; [6] 6軸目（No.5）出力代入済み（RCON受付とは別） *)
    RCON1_ByteOrderConfirmed : BOOL;  (* RCON1 ワード・バイト順確認済み（初期OFF） *)
    RCON1_CommOK : BOOL;  (* RCON1 通信正常（外部判定・固定ON不可） *)
    RCON1_EncodeError : ARRAY[1..6] OF UINT;  (* RCON1 軸別変換エラー番号（0=正常）; [1] 1軸目（No.0）変換エラー番号; [2] 2軸目（No.1）変換エラー番号; [3] 3軸目（No.2）変換エラー番号; [4] 4軸目（No.3）変換エラー番号; [5] 5軸目（No.4）変換エラー番号; [6] 6軸目（No.5）変換エラー番号 *)
    RCON1_EncodeOK : ARRAY[1..6] OF BOOL;  (* RCON1 軸別変換正常（運転許可とは別）; [1] 1軸目（No.0）変換正常; [2] 2軸目（No.1）変換正常; [3] 3軸目（No.2）変換正常; [4] 4軸目（No.3）変換正常; [5] 5軸目（No.4）変換正常; [6] 6軸目（No.5）変換正常 *)
    RCON1_GwAlarmCode : UINT;  (* RCON1 GW異常コード（ALMC/b0～7） *)
    RCON1_GwApply : BOOL;  (* RCON1 共通出力更新許可（OFF=前値保持） *)
    RCON1_GwAxisCommError : BOOL;  (* RCON1 GW－軸 通信異常（ERRT/b13） *)
    RCON1_GwControllerCommLatch : BOOL;  (* RCON1 GW通信異常保持（LERC/b14） *)
    RCON1_GwHeavyAlarm : BOOL;  (* RCON1 GW重故障（ALMH/b11） *)
    RCON1_GwLightAlarm : BOOL;  (* RCON1 GW軽故障（ALML/b10） *)
    RCON1_GwMON_Request : BOOL;  (* RCON1 MON要求（b15） *)
    RCON1_GwManual : BOOL;  (* RCON1 手動モード（MOD/b12） *)
    RCON1_GwRTE_Request : BOOL;  (* RCON1 通信異常ラッチ解除要求（b13） *)
    RCON1_GwRun : BOOL;  (* RCON1 GW動作中（RUN/b15） *)
    RCON1_GwSystemStop : BOOL;  (* RCON1 システム停止状態（SEMG/b8・監視用） *)
    RCON1_GwWritten : BOOL;  (* RCON1 共通出力代入済み（RCON受付とは別） *)
    RCON1_IN : ARRAY[1..6] OF ST_RCON_Direct_IN_Axis;  (* RCON1 入力情報（RCON→PLC）; [1] 1軸目（No.0）入力情報; [2] 2軸目（No.1）入力情報; [3] 3軸目（No.2）入力情報; [4] 4軸目（No.3）入力情報; [5] 5軸目（No.4）入力情報; [6] 6軸目（No.5）入力情報 *)
    RCON1_LayoutConfirmed : BOOL;  (* RCON1 I/O配置確認済み（初期OFF） *)
    RCON1_MotionPermit : ARRAY[1..6] OF BOOL;  (* RCON1 軸別運転許可（外部判定・初期OFF）; [1] 1軸目（No.0）運転許可（外部判定）; [2] 2軸目（No.1）運転許可（外部判定）; [3] 3軸目（No.2）運転許可（外部判定）; [4] 4軸目（No.3）運転許可（外部判定）; [5] 5軸目（No.4）運転許可（外部判定）; [6] 6軸目（No.5）運転許可（外部判定） *)
    RCON1_OUT : ARRAY[1..6] OF ST_RCON_Direct_OUT_Axis;  (* RCON1 出力指令（PLC→RCON）; [1] 1軸目（No.0）出力指令; [2] 2軸目（No.1）出力指令; [3] 3軸目（No.2）出力指令; [4] 4軸目（No.3）出力指令; [5] 5軸目（No.4）出力指令; [6] 6軸目（No.5）出力指令 *)
    RCON1_PowerStateRaw : ARRAY[0..4] OF WORD;  (* RCON1 電源状態ワード（詳細未確認）; [0] IN02 電源状態0（詳細未確認）; [1] IN03 電源状態1（詳細未確認）; [2] IN04 電源状態2（詳細未確認）; [3] IN05 電源状態3（詳細未確認）; [4] IN06 電源状態4（詳細未確認） *)
    RCON1_RxRaw : ARRAY[0..55] OF UINT;  (* RCON1 受信値（バイト交換前）; [0] IN00 GW状態; [1] IN01 軸リンク状態; [2] IN02 電源状態0; [3] IN03 電源状態1; [4] IN04 電源状態2; [5] IN05 電源状態3; [6] IN06 電源状態4（構成依存）; [7] IN07 予約（使用禁止）; [8] IN08 1軸目 現在位置 下位 [0.01mm]; [9] IN09 1軸目 現在位置 上位 [0.01mm]; [10] IN10 1軸目 指令電流 下位 [mA]; [11] IN11 1軸目 指令電流 上位 [mA]; [12] IN12 1軸目 現在速度 [実機単位・符号付き]; [13] IN13 1軸目 予約（使用禁止）; [14] IN14 1軸目 軸異常コード; [15] IN15 1軸目 状態信号（PEND/SV等）; [16] IN16 2軸目 現在位置 下位 [0.01mm]; [17] IN17 2軸目 現在位置 上位 [0.01mm]; [18] IN18 2軸目 指令電流 下位 [mA]; [19] IN19 2軸目 指令電流 上位 [mA]; [20] IN20 2軸目 現在速度 [実機単位・符号付き]; [21] IN21 2軸目 予約（使用禁止）; [22] IN22 2軸目 軸異常コード; [23] IN23 2軸目 状態信号（PEND/SV等）; [24] IN24 3軸目 現在位置 下位 [0.01mm]; [25] IN25 3軸目 現在位置 上位 [0.01mm]; [26] IN26 3軸目 指令電流 下位 [mA]; [27] IN27 3軸目 指令電流 上位 [mA]; [28] IN28 3軸目 現在速度 [実機単位・符号付き]; [29] IN29 3軸目 予約（使用禁止）; [30] IN30 3軸目 軸異常コード; [31] IN31 3軸目 状態信号（PEND/SV等）; [32] IN32 4軸目 現在位置 下位 [0.01mm]; [33] IN33 4軸目 現在位置 上位 [0.01mm]; [34] IN34 4軸目 指令電流 下位 [mA]; [35] IN35 4軸目 指令電流 上位 [mA]; [36] IN36 4軸目 現在速度 [実機単位・符号付き]; [37] IN37 4軸目 予約（使用禁止）; [38] IN38 4軸目 軸異常コード; [39] IN39 4軸目 状態信号（PEND/SV等）; [40] IN40 5軸目 現在位置 下位 [0.01mm]; [41] IN41 5軸目 現在位置 上位 [0.01mm]; [42] IN42 5軸目 指令電流 下位 [mA]; [43] IN43 5軸目 指令電流 上位 [mA]; [44] IN44 5軸目 現在速度 [実機単位・符号付き]; [45] IN45 5軸目 予約（使用禁止）; [46] IN46 5軸目 軸異常コード; [47] IN47 5軸目 状態信号（PEND/SV等）; [48] IN48 6軸目 現在位置 下位 [0.01mm]; [49] IN49 6軸目 現在位置 上位 [0.01mm]; [50] IN50 6軸目 指令電流 下位 [mA]; [51] IN51 6軸目 指令電流 上位 [mA]; [52] IN52 6軸目 現在速度 [実機単位・符号付き]; [53] IN53 6軸目 予約（使用禁止）; [54] IN54 6軸目 軸異常コード; [55] IN55 6軸目 状態信号（PEND/SV等） *)
    RCON1_RxWord : ARRAY[0..55] OF WORD;  (* RCON1 受信ワード（正規化後）; [0] IN00 GW状態; [1] IN01 軸リンク状態; [2] IN02 電源状態0; [3] IN03 電源状態1; [4] IN04 電源状態2; [5] IN05 電源状態3; [6] IN06 電源状態4（構成依存）; [7] IN07 予約（使用禁止）; [8] IN08 1軸目 現在位置 下位 [0.01mm]; [9] IN09 1軸目 現在位置 上位 [0.01mm]; [10] IN10 1軸目 指令電流 下位 [mA]; [11] IN11 1軸目 指令電流 上位 [mA]; [12] IN12 1軸目 現在速度 [実機単位・符号付き]; [13] IN13 1軸目 予約（使用禁止）; [14] IN14 1軸目 軸異常コード; [15] IN15 1軸目 状態信号（PEND/SV等）; [16] IN16 2軸目 現在位置 下位 [0.01mm]; [17] IN17 2軸目 現在位置 上位 [0.01mm]; [18] IN18 2軸目 指令電流 下位 [mA]; [19] IN19 2軸目 指令電流 上位 [mA]; [20] IN20 2軸目 現在速度 [実機単位・符号付き]; [21] IN21 2軸目 予約（使用禁止）; [22] IN22 2軸目 軸異常コード; [23] IN23 2軸目 状態信号（PEND/SV等）; [24] IN24 3軸目 現在位置 下位 [0.01mm]; [25] IN25 3軸目 現在位置 上位 [0.01mm]; [26] IN26 3軸目 指令電流 下位 [mA]; [27] IN27 3軸目 指令電流 上位 [mA]; [28] IN28 3軸目 現在速度 [実機単位・符号付き]; [29] IN29 3軸目 予約（使用禁止）; [30] IN30 3軸目 軸異常コード; [31] IN31 3軸目 状態信号（PEND/SV等）; [32] IN32 4軸目 現在位置 下位 [0.01mm]; [33] IN33 4軸目 現在位置 上位 [0.01mm]; [34] IN34 4軸目 指令電流 下位 [mA]; [35] IN35 4軸目 指令電流 上位 [mA]; [36] IN36 4軸目 現在速度 [実機単位・符号付き]; [37] IN37 4軸目 予約（使用禁止）; [38] IN38 4軸目 軸異常コード; [39] IN39 4軸目 状態信号（PEND/SV等）; [40] IN40 5軸目 現在位置 下位 [0.01mm]; [41] IN41 5軸目 現在位置 上位 [0.01mm]; [42] IN42 5軸目 指令電流 下位 [mA]; [43] IN43 5軸目 指令電流 上位 [mA]; [44] IN44 5軸目 現在速度 [実機単位・符号付き]; [45] IN45 5軸目 予約（使用禁止）; [46] IN46 5軸目 軸異常コード; [47] IN47 5軸目 状態信号（PEND/SV等）; [48] IN48 6軸目 現在位置 下位 [0.01mm]; [49] IN49 6軸目 現在位置 上位 [0.01mm]; [50] IN50 6軸目 指令電流 下位 [mA]; [51] IN51 6軸目 指令電流 上位 [mA]; [52] IN52 6軸目 現在速度 [実機単位・符号付き]; [53] IN53 6軸目 予約（使用禁止）; [54] IN54 6軸目 軸異常コード; [55] IN55 6軸目 状態信号（PEND/SV等） *)
    RCON1_SpeedUnit_mm_s : LREAL;  (* RCON1 速度単位 [mm/s/カウント]（1.0/0.1） *)
    RCON1_SwapBytes : BOOL;  (* RCON1 上下バイト交換設定（ON=交換） *)
    RCON1_TxUInt : ARRAY[0..55] OF UINT;  (* RCON1 送信UINT候補（実I/Oではない）; [0] OUT00 共通制御（MON/RTE）; [1] OUT01 予約（書込禁止）; [2] OUT02 予約（書込禁止）; [3] OUT03 予約（書込禁止）; [4] OUT04 予約（書込禁止）; [5] OUT05 予約（書込禁止）; [6] OUT06 予約（書込禁止）; [7] OUT07 予約（書込禁止）; [8] OUT08 1軸目 目標位置 下位 [0.01mm]; [9] OUT09 1軸目 目標位置 上位 [0.01mm]; [10] OUT10 1軸目 位置決め幅 下位 [0.01mm]; [11] OUT11 1軸目 位置決め幅 上位 [0.01mm]; [12] OUT12 1軸目 速度指令 [実機単位]; [13] OUT13 1軸目 共通加減速 [0.01G]; [14] OUT14 1軸目 押付け制限 [255=100%]; [15] OUT15 1軸目 制御信号（DSTR/SON等）; [16] OUT16 2軸目 目標位置 下位 [0.01mm]; [17] OUT17 2軸目 目標位置 上位 [0.01mm]; [18] OUT18 2軸目 位置決め幅 下位 [0.01mm]; [19] OUT19 2軸目 位置決め幅 上位 [0.01mm]; [20] OUT20 2軸目 速度指令 [実機単位]; [21] OUT21 2軸目 共通加減速 [0.01G]; [22] OUT22 2軸目 押付け制限 [255=100%]; [23] OUT23 2軸目 制御信号（DSTR/SON等）; [24] OUT24 3軸目 目標位置 下位 [0.01mm]; [25] OUT25 3軸目 目標位置 上位 [0.01mm]; [26] OUT26 3軸目 位置決め幅 下位 [0.01mm]; [27] OUT27 3軸目 位置決め幅 上位 [0.01mm]; [28] OUT28 3軸目 速度指令 [実機単位]; [29] OUT29 3軸目 共通加減速 [0.01G]; [30] OUT30 3軸目 押付け制限 [255=100%]; [31] OUT31 3軸目 制御信号（DSTR/SON等）; [32] OUT32 4軸目 目標位置 下位 [0.01mm]; [33] OUT33 4軸目 目標位置 上位 [0.01mm]; [34] OUT34 4軸目 位置決め幅 下位 [0.01mm]; [35] OUT35 4軸目 位置決め幅 上位 [0.01mm]; [36] OUT36 4軸目 速度指令 [実機単位]; [37] OUT37 4軸目 共通加減速 [0.01G]; [38] OUT38 4軸目 押付け制限 [255=100%]; [39] OUT39 4軸目 制御信号（DSTR/SON等）; [40] OUT40 5軸目 目標位置 下位 [0.01mm]; [41] OUT41 5軸目 目標位置 上位 [0.01mm]; [42] OUT42 5軸目 位置決め幅 下位 [0.01mm]; [43] OUT43 5軸目 位置決め幅 上位 [0.01mm]; [44] OUT44 5軸目 速度指令 [実機単位]; [45] OUT45 5軸目 共通加減速 [0.01G]; [46] OUT46 5軸目 押付け制限 [255=100%]; [47] OUT47 5軸目 制御信号（DSTR/SON等）; [48] OUT48 6軸目 目標位置 下位 [0.01mm]; [49] OUT49 6軸目 目標位置 上位 [0.01mm]; [50] OUT50 6軸目 位置決め幅 下位 [0.01mm]; [51] OUT51 6軸目 位置決め幅 上位 [0.01mm]; [52] OUT52 6軸目 速度指令 [実機単位]; [53] OUT53 6軸目 共通加減速 [0.01G]; [54] OUT54 6軸目 押付け制限 [255=100%]; [55] OUT55 6軸目 制御信号（DSTR/SON等） *)
    RCON1_TxWord : ARRAY[0..55] OF WORD;  (* RCON1 送信ワード候補; [0] OUT00 共通制御（MON/RTE）; [1] OUT01 予約（書込禁止）; [2] OUT02 予約（書込禁止）; [3] OUT03 予約（書込禁止）; [4] OUT04 予約（書込禁止）; [5] OUT05 予約（書込禁止）; [6] OUT06 予約（書込禁止）; [7] OUT07 予約（書込禁止）; [8] OUT08 1軸目 目標位置 下位 [0.01mm]; [9] OUT09 1軸目 目標位置 上位 [0.01mm]; [10] OUT10 1軸目 位置決め幅 下位 [0.01mm]; [11] OUT11 1軸目 位置決め幅 上位 [0.01mm]; [12] OUT12 1軸目 速度指令 [実機単位]; [13] OUT13 1軸目 共通加減速 [0.01G]; [14] OUT14 1軸目 押付け制限 [255=100%]; [15] OUT15 1軸目 制御信号（DSTR/SON等）; [16] OUT16 2軸目 目標位置 下位 [0.01mm]; [17] OUT17 2軸目 目標位置 上位 [0.01mm]; [18] OUT18 2軸目 位置決め幅 下位 [0.01mm]; [19] OUT19 2軸目 位置決め幅 上位 [0.01mm]; [20] OUT20 2軸目 速度指令 [実機単位]; [21] OUT21 2軸目 共通加減速 [0.01G]; [22] OUT22 2軸目 押付け制限 [255=100%]; [23] OUT23 2軸目 制御信号（DSTR/SON等）; [24] OUT24 3軸目 目標位置 下位 [0.01mm]; [25] OUT25 3軸目 目標位置 上位 [0.01mm]; [26] OUT26 3軸目 位置決め幅 下位 [0.01mm]; [27] OUT27 3軸目 位置決め幅 上位 [0.01mm]; [28] OUT28 3軸目 速度指令 [実機単位]; [29] OUT29 3軸目 共通加減速 [0.01G]; [30] OUT30 3軸目 押付け制限 [255=100%]; [31] OUT31 3軸目 制御信号（DSTR/SON等）; [32] OUT32 4軸目 目標位置 下位 [0.01mm]; [33] OUT33 4軸目 目標位置 上位 [0.01mm]; [34] OUT34 4軸目 位置決め幅 下位 [0.01mm]; [35] OUT35 4軸目 位置決め幅 上位 [0.01mm]; [36] OUT36 4軸目 速度指令 [実機単位]; [37] OUT37 4軸目 共通加減速 [0.01G]; [38] OUT38 4軸目 押付け制限 [255=100%]; [39] OUT39 4軸目 制御信号（DSTR/SON等）; [40] OUT40 5軸目 目標位置 下位 [0.01mm]; [41] OUT41 5軸目 目標位置 上位 [0.01mm]; [42] OUT42 5軸目 位置決め幅 下位 [0.01mm]; [43] OUT43 5軸目 位置決め幅 上位 [0.01mm]; [44] OUT44 5軸目 速度指令 [実機単位]; [45] OUT45 5軸目 共通加減速 [0.01G]; [46] OUT46 5軸目 押付け制限 [255=100%]; [47] OUT47 5軸目 制御信号（DSTR/SON等）; [48] OUT48 6軸目 目標位置 下位 [0.01mm]; [49] OUT49 6軸目 目標位置 上位 [0.01mm]; [50] OUT50 6軸目 位置決め幅 下位 [0.01mm]; [51] OUT51 6軸目 位置決め幅 上位 [0.01mm]; [52] OUT52 6軸目 速度指令 [実機単位]; [53] OUT53 6軸目 共通加減速 [0.01G]; [54] OUT54 6軸目 押付け制限 [255=100%]; [55] OUT55 6軸目 制御信号（DSTR/SON等） *)
    RCON1_WriteEnable : BOOL;  (* RCON1 実出力書込み許可（OFF=前値保持・停止不可） *)
    RCON2_AxisApply : ARRAY[1..5] OF BOOL;  (* RCON2 軸別出力更新許可（OFF=前値保持）; [1] 1軸目（No.0）出力更新許可（OFF=前値保持）; [2] 2軸目（No.1）出力更新許可（OFF=前値保持）; [3] 3軸目（No.2）出力更新許可（OFF=前値保持）; [4] 4軸目（No.3）出力更新許可（OFF=前値保持）; [5] 5軸目（No.4）出力更新許可（OFF=前値保持） *)
    RCON2_AxisLinked : ARRAY[1..5] OF BOOL;  (* RCON2 軸別リンク状態; [1] 1軸目（No.0）リンク状態; [2] 2軸目（No.1）リンク状態; [3] 3軸目（No.2）リンク状態; [4] 4軸目（No.3）リンク状態; [5] 5軸目（No.4）リンク状態 *)
    RCON2_AxisWritten : ARRAY[1..5] OF BOOL;  (* RCON2 軸別出力代入済み（RCON受付とは別）; [1] 1軸目（No.0）出力代入済み（RCON受付とは別）; [2] 2軸目（No.1）出力代入済み（RCON受付とは別）; [3] 3軸目（No.2）出力代入済み（RCON受付とは別）; [4] 4軸目（No.3）出力代入済み（RCON受付とは別）; [5] 5軸目（No.4）出力代入済み（RCON受付とは別） *)
    RCON2_ByteOrderConfirmed : BOOL;  (* RCON2 ワード・バイト順確認済み（初期OFF） *)
    RCON2_CommOK : BOOL;  (* RCON2 通信正常（外部判定・固定ON不可） *)
    RCON2_EncodeError : ARRAY[1..5] OF UINT;  (* RCON2 軸別変換エラー番号（0=正常）; [1] 1軸目（No.0）変換エラー番号; [2] 2軸目（No.1）変換エラー番号; [3] 3軸目（No.2）変換エラー番号; [4] 4軸目（No.3）変換エラー番号; [5] 5軸目（No.4）変換エラー番号 *)
    RCON2_EncodeOK : ARRAY[1..5] OF BOOL;  (* RCON2 軸別変換正常（運転許可とは別）; [1] 1軸目（No.0）変換正常; [2] 2軸目（No.1）変換正常; [3] 3軸目（No.2）変換正常; [4] 4軸目（No.3）変換正常; [5] 5軸目（No.4）変換正常 *)
    RCON2_GwAlarmCode : UINT;  (* RCON2 GW異常コード（ALMC/b0～7） *)
    RCON2_GwApply : BOOL;  (* RCON2 共通出力更新許可（OFF=前値保持） *)
    RCON2_GwAxisCommError : BOOL;  (* RCON2 GW－軸 通信異常（ERRT/b13） *)
    RCON2_GwControllerCommLatch : BOOL;  (* RCON2 GW通信異常保持（LERC/b14） *)
    RCON2_GwHeavyAlarm : BOOL;  (* RCON2 GW重故障（ALMH/b11） *)
    RCON2_GwLightAlarm : BOOL;  (* RCON2 GW軽故障（ALML/b10） *)
    RCON2_GwMON_Request : BOOL;  (* RCON2 MON要求（b15） *)
    RCON2_GwManual : BOOL;  (* RCON2 手動モード（MOD/b12） *)
    RCON2_GwRTE_Request : BOOL;  (* RCON2 通信異常ラッチ解除要求（b13） *)
    RCON2_GwRun : BOOL;  (* RCON2 GW動作中（RUN/b15） *)
    RCON2_GwSystemStop : BOOL;  (* RCON2 システム停止状態（SEMG/b8・監視用） *)
    RCON2_GwWritten : BOOL;  (* RCON2 共通出力代入済み（RCON受付とは別） *)
    RCON2_IN : ARRAY[1..5] OF ST_RCON_Direct_IN_Axis;  (* RCON2 入力情報（RCON→PLC）; [1] 1軸目（No.0）入力情報; [2] 2軸目（No.1）入力情報; [3] 3軸目（No.2）入力情報; [4] 4軸目（No.3）入力情報; [5] 5軸目（No.4）入力情報 *)
    RCON2_LayoutConfirmed : BOOL;  (* RCON2 I/O配置確認済み（初期OFF） *)
    RCON2_MotionPermit : ARRAY[1..5] OF BOOL;  (* RCON2 軸別運転許可（外部判定・初期OFF）; [1] 1軸目（No.0）運転許可（外部判定）; [2] 2軸目（No.1）運転許可（外部判定）; [3] 3軸目（No.2）運転許可（外部判定）; [4] 4軸目（No.3）運転許可（外部判定）; [5] 5軸目（No.4）運転許可（外部判定） *)
    RCON2_OUT : ARRAY[1..5] OF ST_RCON_Direct_OUT_Axis;  (* RCON2 出力指令（PLC→RCON）; [1] 1軸目（No.0）出力指令; [2] 2軸目（No.1）出力指令; [3] 3軸目（No.2）出力指令; [4] 4軸目（No.3）出力指令; [5] 5軸目（No.4）出力指令 *)
    RCON2_PowerStateRaw : ARRAY[0..4] OF WORD;  (* RCON2 電源状態ワード（詳細未確認）; [0] IN02 電源状態0（詳細未確認）; [1] IN03 電源状態1（詳細未確認）; [2] IN04 電源状態2（詳細未確認）; [3] IN05 電源状態3（詳細未確認）; [4] IN06 電源状態4（詳細未確認） *)
    RCON2_RxRaw : ARRAY[0..55] OF UINT;  (* RCON2 受信値（バイト交換前）; [0] IN00 GW状態; [1] IN01 軸リンク状態; [2] IN02 電源状態0; [3] IN03 電源状態1; [4] IN04 電源状態2; [5] IN05 電源状態3; [6] IN06 電源状態4（構成依存）; [7] IN07 予約（使用禁止）; [8] IN08 1軸目 現在位置 下位 [0.01mm]; [9] IN09 1軸目 現在位置 上位 [0.01mm]; [10] IN10 1軸目 指令電流 下位 [mA]; [11] IN11 1軸目 指令電流 上位 [mA]; [12] IN12 1軸目 現在速度 [実機単位・符号付き]; [13] IN13 1軸目 予約（使用禁止）; [14] IN14 1軸目 軸異常コード; [15] IN15 1軸目 状態信号（PEND/SV等）; [16] IN16 2軸目 現在位置 下位 [0.01mm]; [17] IN17 2軸目 現在位置 上位 [0.01mm]; [18] IN18 2軸目 指令電流 下位 [mA]; [19] IN19 2軸目 指令電流 上位 [mA]; [20] IN20 2軸目 現在速度 [実機単位・符号付き]; [21] IN21 2軸目 予約（使用禁止）; [22] IN22 2軸目 軸異常コード; [23] IN23 2軸目 状態信号（PEND/SV等）; [24] IN24 3軸目 現在位置 下位 [0.01mm]; [25] IN25 3軸目 現在位置 上位 [0.01mm]; [26] IN26 3軸目 指令電流 下位 [mA]; [27] IN27 3軸目 指令電流 上位 [mA]; [28] IN28 3軸目 現在速度 [実機単位・符号付き]; [29] IN29 3軸目 予約（使用禁止）; [30] IN30 3軸目 軸異常コード; [31] IN31 3軸目 状態信号（PEND/SV等）; [32] IN32 4軸目 現在位置 下位 [0.01mm]; [33] IN33 4軸目 現在位置 上位 [0.01mm]; [34] IN34 4軸目 指令電流 下位 [mA]; [35] IN35 4軸目 指令電流 上位 [mA]; [36] IN36 4軸目 現在速度 [実機単位・符号付き]; [37] IN37 4軸目 予約（使用禁止）; [38] IN38 4軸目 軸異常コード; [39] IN39 4軸目 状態信号（PEND/SV等）; [40] IN40 5軸目 現在位置 下位 [0.01mm]; [41] IN41 5軸目 現在位置 上位 [0.01mm]; [42] IN42 5軸目 指令電流 下位 [mA]; [43] IN43 5軸目 指令電流 上位 [mA]; [44] IN44 5軸目 現在速度 [実機単位・符号付き]; [45] IN45 5軸目 予約（使用禁止）; [46] IN46 5軸目 軸異常コード; [47] IN47 5軸目 状態信号（PEND/SV等）; [48] IN48 用途未確認（今回未使用）; [49] IN49 用途未確認（今回未使用）; [50] IN50 用途未確認（今回未使用）; [51] IN51 用途未確認（今回未使用）; [52] IN52 用途未確認（今回未使用）; [53] IN53 用途未確認（今回未使用）; [54] IN54 用途未確認（今回未使用）; [55] IN55 用途未確認（今回未使用） *)
    RCON2_RxWord : ARRAY[0..55] OF WORD;  (* RCON2 受信ワード（正規化後）; [0] IN00 GW状態; [1] IN01 軸リンク状態; [2] IN02 電源状態0; [3] IN03 電源状態1; [4] IN04 電源状態2; [5] IN05 電源状態3; [6] IN06 電源状態4（構成依存）; [7] IN07 予約（使用禁止）; [8] IN08 1軸目 現在位置 下位 [0.01mm]; [9] IN09 1軸目 現在位置 上位 [0.01mm]; [10] IN10 1軸目 指令電流 下位 [mA]; [11] IN11 1軸目 指令電流 上位 [mA]; [12] IN12 1軸目 現在速度 [実機単位・符号付き]; [13] IN13 1軸目 予約（使用禁止）; [14] IN14 1軸目 軸異常コード; [15] IN15 1軸目 状態信号（PEND/SV等）; [16] IN16 2軸目 現在位置 下位 [0.01mm]; [17] IN17 2軸目 現在位置 上位 [0.01mm]; [18] IN18 2軸目 指令電流 下位 [mA]; [19] IN19 2軸目 指令電流 上位 [mA]; [20] IN20 2軸目 現在速度 [実機単位・符号付き]; [21] IN21 2軸目 予約（使用禁止）; [22] IN22 2軸目 軸異常コード; [23] IN23 2軸目 状態信号（PEND/SV等）; [24] IN24 3軸目 現在位置 下位 [0.01mm]; [25] IN25 3軸目 現在位置 上位 [0.01mm]; [26] IN26 3軸目 指令電流 下位 [mA]; [27] IN27 3軸目 指令電流 上位 [mA]; [28] IN28 3軸目 現在速度 [実機単位・符号付き]; [29] IN29 3軸目 予約（使用禁止）; [30] IN30 3軸目 軸異常コード; [31] IN31 3軸目 状態信号（PEND/SV等）; [32] IN32 4軸目 現在位置 下位 [0.01mm]; [33] IN33 4軸目 現在位置 上位 [0.01mm]; [34] IN34 4軸目 指令電流 下位 [mA]; [35] IN35 4軸目 指令電流 上位 [mA]; [36] IN36 4軸目 現在速度 [実機単位・符号付き]; [37] IN37 4軸目 予約（使用禁止）; [38] IN38 4軸目 軸異常コード; [39] IN39 4軸目 状態信号（PEND/SV等）; [40] IN40 5軸目 現在位置 下位 [0.01mm]; [41] IN41 5軸目 現在位置 上位 [0.01mm]; [42] IN42 5軸目 指令電流 下位 [mA]; [43] IN43 5軸目 指令電流 上位 [mA]; [44] IN44 5軸目 現在速度 [実機単位・符号付き]; [45] IN45 5軸目 予約（使用禁止）; [46] IN46 5軸目 軸異常コード; [47] IN47 5軸目 状態信号（PEND/SV等）; [48] IN48 用途未確認（今回未使用）; [49] IN49 用途未確認（今回未使用）; [50] IN50 用途未確認（今回未使用）; [51] IN51 用途未確認（今回未使用）; [52] IN52 用途未確認（今回未使用）; [53] IN53 用途未確認（今回未使用）; [54] IN54 用途未確認（今回未使用）; [55] IN55 用途未確認（今回未使用） *)
    RCON2_SpeedUnit_mm_s : LREAL;  (* RCON2 速度単位 [mm/s/カウント]（1.0/0.1） *)
    RCON2_SwapBytes : BOOL;  (* RCON2 上下バイト交換設定（ON=交換） *)
    RCON2_TxUInt : ARRAY[0..47] OF UINT;  (* RCON2 送信UINT候補（実I/Oではない）; [0] OUT00 共通制御（MON/RTE）; [1] OUT01 予約（書込禁止）; [2] OUT02 予約（書込禁止）; [3] OUT03 予約（書込禁止）; [4] OUT04 予約（書込禁止）; [5] OUT05 予約（書込禁止）; [6] OUT06 予約（書込禁止）; [7] OUT07 予約（書込禁止）; [8] OUT08 1軸目 目標位置 下位 [0.01mm]; [9] OUT09 1軸目 目標位置 上位 [0.01mm]; [10] OUT10 1軸目 位置決め幅 下位 [0.01mm]; [11] OUT11 1軸目 位置決め幅 上位 [0.01mm]; [12] OUT12 1軸目 速度指令 [実機単位]; [13] OUT13 1軸目 共通加減速 [0.01G]; [14] OUT14 1軸目 押付け制限 [255=100%]; [15] OUT15 1軸目 制御信号（DSTR/SON等）; [16] OUT16 2軸目 目標位置 下位 [0.01mm]; [17] OUT17 2軸目 目標位置 上位 [0.01mm]; [18] OUT18 2軸目 位置決め幅 下位 [0.01mm]; [19] OUT19 2軸目 位置決め幅 上位 [0.01mm]; [20] OUT20 2軸目 速度指令 [実機単位]; [21] OUT21 2軸目 共通加減速 [0.01G]; [22] OUT22 2軸目 押付け制限 [255=100%]; [23] OUT23 2軸目 制御信号（DSTR/SON等）; [24] OUT24 3軸目 目標位置 下位 [0.01mm]; [25] OUT25 3軸目 目標位置 上位 [0.01mm]; [26] OUT26 3軸目 位置決め幅 下位 [0.01mm]; [27] OUT27 3軸目 位置決め幅 上位 [0.01mm]; [28] OUT28 3軸目 速度指令 [実機単位]; [29] OUT29 3軸目 共通加減速 [0.01G]; [30] OUT30 3軸目 押付け制限 [255=100%]; [31] OUT31 3軸目 制御信号（DSTR/SON等）; [32] OUT32 4軸目 目標位置 下位 [0.01mm]; [33] OUT33 4軸目 目標位置 上位 [0.01mm]; [34] OUT34 4軸目 位置決め幅 下位 [0.01mm]; [35] OUT35 4軸目 位置決め幅 上位 [0.01mm]; [36] OUT36 4軸目 速度指令 [実機単位]; [37] OUT37 4軸目 共通加減速 [0.01G]; [38] OUT38 4軸目 押付け制限 [255=100%]; [39] OUT39 4軸目 制御信号（DSTR/SON等）; [40] OUT40 5軸目 目標位置 下位 [0.01mm]; [41] OUT41 5軸目 目標位置 上位 [0.01mm]; [42] OUT42 5軸目 位置決め幅 下位 [0.01mm]; [43] OUT43 5軸目 位置決め幅 上位 [0.01mm]; [44] OUT44 5軸目 速度指令 [実機単位]; [45] OUT45 5軸目 共通加減速 [0.01G]; [46] OUT46 5軸目 押付け制限 [255=100%]; [47] OUT47 5軸目 制御信号（DSTR/SON等） *)
    RCON2_TxWord : ARRAY[0..47] OF WORD;  (* RCON2 送信ワード候補; [0] OUT00 共通制御（MON/RTE）; [1] OUT01 予約（書込禁止）; [2] OUT02 予約（書込禁止）; [3] OUT03 予約（書込禁止）; [4] OUT04 予約（書込禁止）; [5] OUT05 予約（書込禁止）; [6] OUT06 予約（書込禁止）; [7] OUT07 予約（書込禁止）; [8] OUT08 1軸目 目標位置 下位 [0.01mm]; [9] OUT09 1軸目 目標位置 上位 [0.01mm]; [10] OUT10 1軸目 位置決め幅 下位 [0.01mm]; [11] OUT11 1軸目 位置決め幅 上位 [0.01mm]; [12] OUT12 1軸目 速度指令 [実機単位]; [13] OUT13 1軸目 共通加減速 [0.01G]; [14] OUT14 1軸目 押付け制限 [255=100%]; [15] OUT15 1軸目 制御信号（DSTR/SON等）; [16] OUT16 2軸目 目標位置 下位 [0.01mm]; [17] OUT17 2軸目 目標位置 上位 [0.01mm]; [18] OUT18 2軸目 位置決め幅 下位 [0.01mm]; [19] OUT19 2軸目 位置決め幅 上位 [0.01mm]; [20] OUT20 2軸目 速度指令 [実機単位]; [21] OUT21 2軸目 共通加減速 [0.01G]; [22] OUT22 2軸目 押付け制限 [255=100%]; [23] OUT23 2軸目 制御信号（DSTR/SON等）; [24] OUT24 3軸目 目標位置 下位 [0.01mm]; [25] OUT25 3軸目 目標位置 上位 [0.01mm]; [26] OUT26 3軸目 位置決め幅 下位 [0.01mm]; [27] OUT27 3軸目 位置決め幅 上位 [0.01mm]; [28] OUT28 3軸目 速度指令 [実機単位]; [29] OUT29 3軸目 共通加減速 [0.01G]; [30] OUT30 3軸目 押付け制限 [255=100%]; [31] OUT31 3軸目 制御信号（DSTR/SON等）; [32] OUT32 4軸目 目標位置 下位 [0.01mm]; [33] OUT33 4軸目 目標位置 上位 [0.01mm]; [34] OUT34 4軸目 位置決め幅 下位 [0.01mm]; [35] OUT35 4軸目 位置決め幅 上位 [0.01mm]; [36] OUT36 4軸目 速度指令 [実機単位]; [37] OUT37 4軸目 共通加減速 [0.01G]; [38] OUT38 4軸目 押付け制限 [255=100%]; [39] OUT39 4軸目 制御信号（DSTR/SON等）; [40] OUT40 5軸目 目標位置 下位 [0.01mm]; [41] OUT41 5軸目 目標位置 上位 [0.01mm]; [42] OUT42 5軸目 位置決め幅 下位 [0.01mm]; [43] OUT43 5軸目 位置決め幅 上位 [0.01mm]; [44] OUT44 5軸目 速度指令 [実機単位]; [45] OUT45 5軸目 共通加減速 [0.01G]; [46] OUT46 5軸目 押付け制限 [255=100%]; [47] OUT47 5軸目 制御信号（DSTR/SON等） *)
    RCON2_WriteEnable : BOOL;  (* RCON2 実出力書込み許可（OFF=前値保持・停止不可） *)
    RCON1_IAI_Auto : ARRAY[0..99] OF Bool;
    RCON1_OUT_PositionBand_mm : LREAL;  (* RCON1位置決め幅 [mm] *)
    RCON1_OUT_TargetPos_mm : LREAL;  (* RCON1目標位置 [mm] *)
    RCON1_OUT_Speed_mm_s : LREAL;  (* 指令速度 [mm/s] *)
    RCON1_OUT_AccDec_G : LREAL;  (* 共通加減速度 [G] *)
    RCON1_OUT_PushLimit_pct : LREAL;  (* 押付け電流制限 [%] *)
    RCON1_ActualPos_mm : LREAL;  (* 現在位置 [mm] *)
    RCON1_Current_mA : DINT;  (* 指令電流 [mA] *)
    RCON1_ActualSpeed_mm_s : LREAL;  (* 現在速度 [mm/s・符号付き] *)
    RCON1_AlarmCode : UINT;  (* 軸異常コード *)
    RCON1_DataValid : BOOL;  (* 入力有効（運転許可とは別） *)
    RCON1_1_IN_PositionDone : BOOL;  (* 位置決め完了 *)
    RCON1_1_IN_HomeDone : BOOL;  (* 原点復帰完了 *)
    RCON1_1_IN_Moving : BOOL;  (* 移動中 *)
    RCON1_1_IN_EmergencyStop : BOOL;  (* 非常停止状態 *)
    RCON1_1_IN_ControllerReady : BOOL;  (* コントローラー準備完了 *)
    RCON1_1_IN_Zone2 : BOOL;  (* ゾーン2内 *)
    RCON1_1_IN_Zone1 : BOOL;  (* ゾーン1内 *)
    RCON1_1_IN_CommandDone : BOOL;  (* 指令完了 *)
    RCON1_1_IN_OverloadWarning : BOOL;  (* 過負荷警告等 *)
    RCON1_1_IN_PushMiss : BOOL;  (* 押付け空振り *)
    RCON1_1_IN_ServoReady : BOOL;  (* サーボON状態 *)
    RCON1_1_IN_Alarm : BOOL;  (* 軸異常 *)
    RCON1_1_Ready : BOOL;  (* RCON1 運転可能状態 *)
    RCON1_1_Error_Clear : BOOL;
    Error_M : ARRAY[0..99] OF Bool;
    In_Sw_RESET : BOOL;
    RCON1_1_M : ARRAY[0..99] OF BOOL;
    TimerQ_In_SenCY_NG1_Pick_A_H : BOOL;
    Homing_Para_Stm : _sHOMING_REF;
END_VAR
VAR_EXTERNAL CONSTANT
    Stm_A_Rev_Axis000 : _sAXIS_REF;
END_VAR
VAR_EXTERNAL
    Stm_A_Rev_Axis000_OriginDone : BOOL;  (* A(左側) ST4 反転1 モータ原点復帰完了 *)
    Auto_A_Start : BOOL;
    HMI_Home_SW : BOOL;  (* HMI 原点復帰SW *)
    Stm_A_Rev_Axis000_Origin : BOOL;  (* A(左側) ST4 反転1 モータ原点復帰開始 *)
    Stm_A_Rev_Axis000_MovePos_Degree : LREAL;  (* A(左側)ステッピングモータ000 回転角度 *)
    Stm_A_Rev_Axis000_MoveAbsoluteDone : BOOL;  (* A(左側)ステッピング反転モータ1 絶対値位置決め 動作完了 *)
    Stm_A_Rev_Axis000_Auto : ARRAY[0..99] OF Bool;
END_VAR
VAR
    _e1 : R_TRIG;
    _e2 : R_TRIG;
    _e3 : R_TRIG;
    _p4 : BOOL;
    _e5 : R_TRIG;
    _p6 : BOOL;
    _e7 : R_TRIG;
    _p8 : BOOL;
    _e9 : R_TRIG;
    _p10 : BOOL;
    _e11 : R_TRIG;
    _e12 : R_TRIG;
    _p13 : BOOL;
    _e14 : R_TRIG;
    _e15 : R_TRIG;
    _p16 : BOOL;
    _p17 : BOOL;
    _p18 : BOOL;
END_VAR

(* Section RCON_IAI: ladder, written here as Structured Text *)

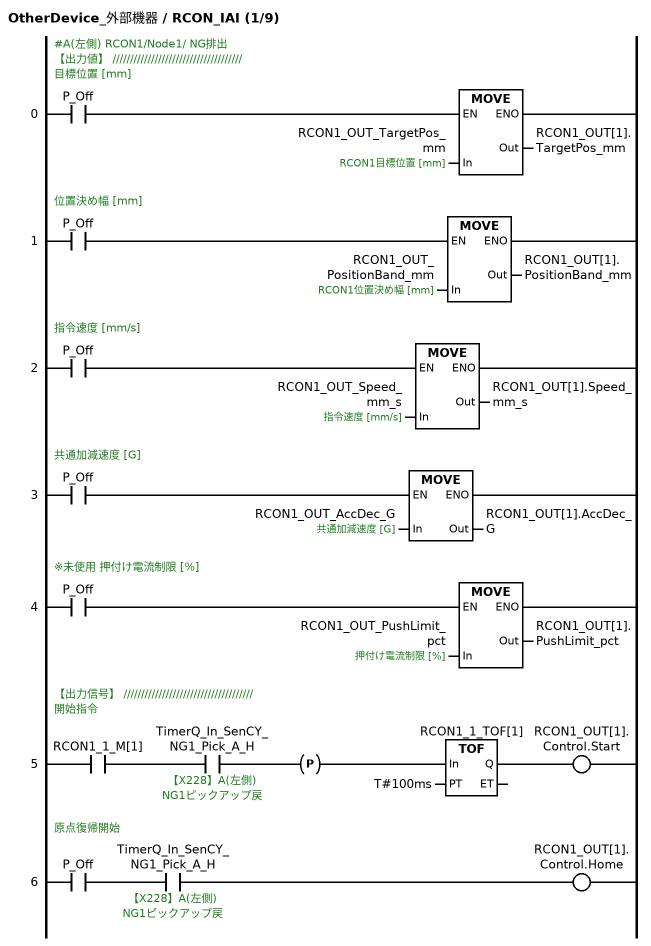
(* Rung 0: #A(左側) RCON1/Node1/ NG排出 / 【出力値】 ///////////////////////////////////// / 目標位置 [mm] *)
IF P_Off THEN RCON1_OUT[1].TargetPos_mm := RCON1_OUT_TargetPos_mm; END_IF;
(* Rung 1: 位置決め幅 [mm] *)
IF P_Off THEN RCON1_OUT[1].PositionBand_mm := RCON1_OUT_PositionBand_mm; END_IF;
(* Rung 2: 指令速度 [mm/s] *)
IF P_Off THEN RCON1_OUT[1].Speed_mm_s := RCON1_OUT_Speed_mm_s; END_IF;
(* Rung 3: 共通加減速度 [G] *)
IF P_Off THEN RCON1_OUT[1].AccDec_G := RCON1_OUT_AccDec_G; END_IF;
(* Rung 4: ※未使用 押付け電流制限 [%] *)
IF P_Off THEN RCON1_OUT[1].PushLimit_pct := RCON1_OUT_PushLimit_pct; END_IF;
(* Rung 5: 【出力信号】 ///////////////////////////////////// / 開始指令 *)
_e1(CLK := RCON1_1_M[1] AND TimerQ_In_SenCY_NG1_Pick_A_H);
RCON1_1_TOF[1](In := _e1.Q, PT := T#100ms);
RCON1_OUT[1].Control.Start := RCON1_1_TOF[1].Q;
(* Rung 6: 原点復帰開始 *)
RCON1_OUT[1].Control.Home := P_Off AND TimerQ_In_SenCY_NG1_Pick_A_H;

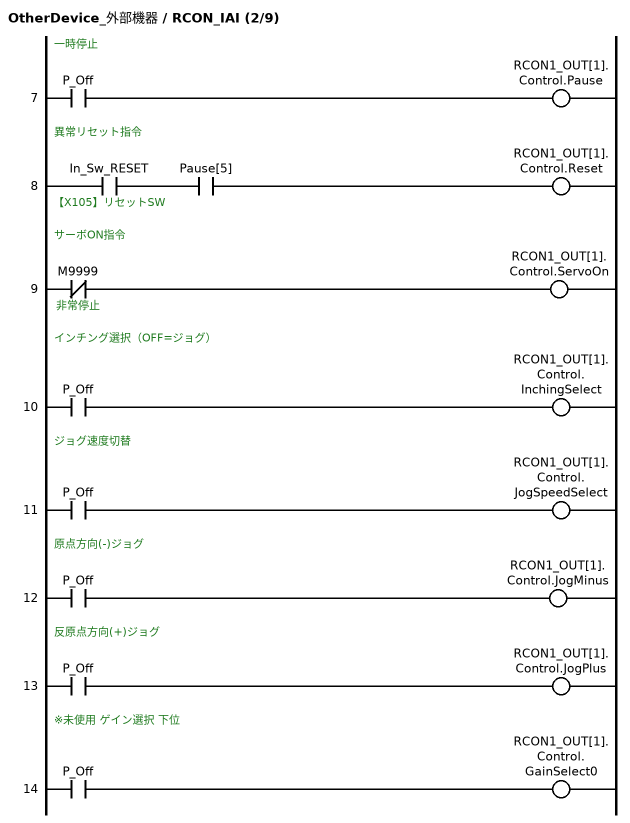
(* Rung 7: 一時停止 *)
RCON1_OUT[1].Control.Pause := P_Off;
(* Rung 8: 異常リセット指令 *)
RCON1_OUT[1].Control.Reset := In_Sw_RESET AND Pause[5];
(* Rung 9: サーボON指令 *)
RCON1_OUT[1].Control.ServoOn := NOT M9999;
(* Rung 10: インチング選択（OFF=ジョグ） *)
RCON1_OUT[1].Control.InchingSelect := P_Off;
(* Rung 11: ジョグ速度切替 *)
RCON1_OUT[1].Control.JogSpeedSelect := P_Off;
(* Rung 12: 原点方向(-)ジョグ *)
RCON1_OUT[1].Control.JogMinus := P_Off;
(* Rung 13: 反原点方向(+)ジョグ *)
RCON1_OUT[1].Control.JogPlus := P_Off;
(* Rung 14: ※未使用 ゲイン選択 下位 *)
RCON1_OUT[1].Control.GainSelect0 := P_Off;

